(* IEC 61131-3 sources: STAR-PLC-Agent/results/raw/codex_matrix_resume_20261114/codex_deepseek/PUB020/functional/attempt_0001, 1 file *)

(* ---- test_program.st ---- *)
PROGRAM PLC_PRG
VAR
 BenchStep : UDINT := 0;
 BenchCalls : UDINT := 0;
 BenchDone : BOOL := FALSE;
 BenchUut0 : FB_Task;
 BenchUut1 : FB_Task;
 BenchUut2 : FB_Task;
 BenchUut3 : FB_Task;
 BenchUut4 : FB_Task;
 BenchUut5 : FB_Task;
 BenchUut6 : FB_Task;
 BenchUut7 : FB_Task;
 BenchUut8 : FB_Task;
 BenchUut9 : FB_Task;
 BenchUut10 : FB_Task;
 TraceIn_Mode : ARRAY[0..155] OF BOOL;
 TraceIn_ForwardButton : ARRAY[0..155] OF BOOL;
 TraceIn_ReverseButton : ARRAY[0..155] OF BOOL;
 TraceIn_SensorFeed : ARRAY[0..155] OF BOOL;
 TraceIn_SensorWash : ARRAY[0..155] OF BOOL;
 TraceIn_SensorWeight : ARRAY[0..155] OF BOOL;
 TraceIn_SensorFiring : ARRAY[0..155] OF BOOL;
 TraceIn_SensorOutput : ARRAY[0..155] OF BOOL;
 TraceIn_washComplete : ARRAY[0..155] OF BOOL;
 TraceIn_weightComplete : ARRAY[0..155] OF BOOL;
 TraceIn_weight : ARRAY[0..155] OF REAL;
 TraceIn_firingComplete : ARRAY[0..155] OF BOOL;
 TraceOut_MotorForward : ARRAY[0..155] OF BOOL;
 TraceOut_MotorReverse : ARRAY[0..155] OF BOOL;
 TraceOut_kick : ARRAY[0..155] OF BOOL;
 TraceOut_CompletionLight : ARRAY[0..155] OF BOOL;
 TraceOut_firingTemp : ARRAY[0..155] OF REAL;
END_VAR

IF NOT BenchDone THEN
 CASE BenchStep OF
 0:
   BenchUut0.Mode := FALSE;
   BenchUut0.ForwardButton := FALSE;
   BenchUut0.ReverseButton := FALSE;
   BenchUut0.SensorFeed := FALSE;
   BenchUut0.SensorWash := FALSE;
   BenchUut0.SensorWeight := FALSE;
   BenchUut0.SensorFiring := FALSE;
   BenchUut0.SensorOutput := FALSE;
   BenchUut0.washComplete := FALSE;
   BenchUut0.weightComplete := FALSE;
   BenchUut0.weight := REAL#0.0;
   BenchUut0.firingComplete := FALSE;
   TraceIn_Mode[0] := BenchUut0.Mode;
   TraceIn_ForwardButton[0] := BenchUut0.ForwardButton;
   TraceIn_ReverseButton[0] := BenchUut0.ReverseButton;
   TraceIn_SensorFeed[0] := BenchUut0.SensorFeed;
   TraceIn_SensorWash[0] := BenchUut0.SensorWash;
   TraceIn_SensorWeight[0] := BenchUut0.SensorWeight;
   TraceIn_SensorFiring[0] := BenchUut0.SensorFiring;
   TraceIn_SensorOutput[0] := BenchUut0.SensorOutput;
   TraceIn_washComplete[0] := BenchUut0.washComplete;
   TraceIn_weightComplete[0] := BenchUut0.weightComplete;
   TraceIn_weight[0] := BenchUut0.weight;
   TraceIn_firingComplete[0] := BenchUut0.firingComplete;
   BenchUut0();
   TraceOut_MotorForward[0] := BenchUut0.MotorForward;
   TraceOut_MotorReverse[0] := BenchUut0.MotorReverse;
   TraceOut_kick[0] := BenchUut0.kick;
   TraceOut_CompletionLight[0] := BenchUut0.CompletionLight;
   TraceOut_firingTemp[0] := BenchUut0.firingTemp;
   BenchCalls := BenchCalls + 1;
 1:
   BenchUut0.Mode := FALSE;
   BenchUut0.ForwardButton := TRUE;
   BenchUut0.ReverseButton := FALSE;
   BenchUut0.SensorFeed := FALSE;
   BenchUut0.SensorWash := FALSE;
   BenchUut0.SensorWeight := FALSE;
   BenchUut0.SensorFiring := FALSE;
   BenchUut0.SensorOutput := FALSE;
   BenchUut0.washComplete := FALSE;
   BenchUut0.weightComplete := FALSE;
   BenchUut0.weight := REAL#0.0;
   BenchUut0.firingComplete := FALSE;
   TraceIn_Mode[1] := BenchUut0.Mode;
   TraceIn_ForwardButton[1] := BenchUut0.ForwardButton;
   TraceIn_ReverseButton[1] := BenchUut0.ReverseButton;
   TraceIn_SensorFeed[1] := BenchUut0.SensorFeed;
   TraceIn_SensorWash[1] := BenchUut0.SensorWash;
   TraceIn_SensorWeight[1] := BenchUut0.SensorWeight;
   TraceIn_SensorFiring[1] := BenchUut0.SensorFiring;
   TraceIn_SensorOutput[1] := BenchUut0.SensorOutput;
   TraceIn_washComplete[1] := BenchUut0.washComplete;
   TraceIn_weightComplete[1] := BenchUut0.weightComplete;
   TraceIn_weight[1] := BenchUut0.weight;
   TraceIn_firingComplete[1] := BenchUut0.firingComplete;
   BenchUut0();
   TraceOut_MotorForward[1] := BenchUut0.MotorForward;
   TraceOut_MotorReverse[1] := BenchUut0.MotorReverse;
   TraceOut_kick[1] := BenchUut0.kick;
   TraceOut_CompletionLight[1] := BenchUut0.CompletionLight;
   TraceOut_firingTemp[1] := BenchUut0.firingTemp;
   BenchCalls := BenchCalls + 1;
 2:
   BenchUut0.Mode := FALSE;
   BenchUut0.ForwardButton := FALSE;
   BenchUut0.ReverseButton := TRUE;
   BenchUut0.SensorFeed := FALSE;
   BenchUut0.SensorWash := FALSE;
   BenchUut0.SensorWeight := FALSE;
   BenchUut0.SensorFiring := FALSE;
   BenchUut0.SensorOutput := FALSE;
   BenchUut0.washComplete := FALSE;
   BenchUut0.weightComplete := FALSE;
   BenchUut0.weight := REAL#0.0;
   BenchUut0.firingComplete := FALSE;
   TraceIn_Mode[2] := BenchUut0.Mode;
   TraceIn_ForwardButton[2] := BenchUut0.ForwardButton;
   TraceIn_ReverseButton[2] := BenchUut0.ReverseButton;
   TraceIn_SensorFeed[2] := BenchUut0.SensorFeed;
   TraceIn_SensorWash[2] := BenchUut0.SensorWash;
   TraceIn_SensorWeight[2] := BenchUut0.SensorWeight;
   TraceIn_SensorFiring[2] := BenchUut0.SensorFiring;
   TraceIn_SensorOutput[2] := BenchUut0.SensorOutput;
   TraceIn_washComplete[2] := BenchUut0.washComplete;
   TraceIn_weightComplete[2] := BenchUut0.weightComplete;
   TraceIn_weight[2] := BenchUut0.weight;
   TraceIn_firingComplete[2] := BenchUut0.firingComplete;
   BenchUut0();
   TraceOut_MotorForward[2] := BenchUut0.MotorForward;
   TraceOut_MotorReverse[2] := BenchUut0.MotorReverse;
   TraceOut_kick[2] := BenchUut0.kick;
   TraceOut_CompletionLight[2] := BenchUut0.CompletionLight;
   TraceOut_firingTemp[2] := BenchUut0.firingTemp;
   BenchCalls := BenchCalls + 1;
 3:
   BenchUut0.Mode := FALSE;
   BenchUut0.ForwardButton := TRUE;
   BenchUut0.ReverseButton := TRUE;
   BenchUut0.SensorFeed := FALSE;
   BenchUut0.SensorWash := FALSE;
   BenchUut0.SensorWeight := FALSE;
   BenchUut0.SensorFiring := FALSE;
   BenchUut0.SensorOutput := FALSE;
   BenchUut0.washComplete := FALSE;
   BenchUut0.weightComplete := FALSE;
   BenchUut0.weight := REAL#0.0;
   BenchUut0.firingComplete := FALSE;
   TraceIn_Mode[3] := BenchUut0.Mode;
   TraceIn_ForwardButton[3] := BenchUut0.ForwardButton;
   TraceIn_ReverseButton[3] := BenchUut0.ReverseButton;
   TraceIn_SensorFeed[3] := BenchUut0.SensorFeed;
   TraceIn_SensorWash[3] := BenchUut0.SensorWash;
   TraceIn_SensorWeight[3] := BenchUut0.SensorWeight;
   TraceIn_SensorFiring[3] := BenchUut0.SensorFiring;
   TraceIn_SensorOutput[3] := BenchUut0.SensorOutput;
   TraceIn_washComplete[3] := BenchUut0.washComplete;
   TraceIn_weightComplete[3] := BenchUut0.weightComplete;
   TraceIn_weight[3] := BenchUut0.weight;
   TraceIn_firingComplete[3] := BenchUut0.firingComplete;
   BenchUut0();
   TraceOut_MotorForward[3] := BenchUut0.MotorForward;
   TraceOut_MotorReverse[3] := BenchUut0.MotorReverse;
   TraceOut_kick[3] := BenchUut0.kick;
   TraceOut_CompletionLight[3] := BenchUut0.CompletionLight;
   TraceOut_firingTemp[3] := BenchUut0.firingTemp;
   BenchCalls := BenchCalls + 1;
 4:
   BenchUut1.Mode := TRUE;
   BenchUut1.ForwardButton := FALSE;
   BenchUut1.ReverseButton := FALSE;
   BenchUut1.SensorFeed := FALSE;
   BenchUut1.SensorWash := FALSE;
   BenchUut1.SensorWeight := FALSE;
   BenchUut1.SensorFiring := FALSE;
   BenchUut1.SensorOutput := FALSE;
   BenchUut1.washComplete := FALSE;
   BenchUut1.weightComplete := FALSE;
   BenchUut1.weight := REAL#0.0;
   BenchUut1.firingComplete := FALSE;
   TraceIn_Mode[4] := BenchUut1.Mode;
   TraceIn_ForwardButton[4] := BenchUut1.ForwardButton;
   TraceIn_ReverseButton[4] := BenchUut1.ReverseButton;
   TraceIn_SensorFeed[4] := BenchUut1.SensorFeed;
   TraceIn_SensorWash[4] := BenchUut1.SensorWash;
   TraceIn_SensorWeight[4] := BenchUut1.SensorWeight;
   TraceIn_SensorFiring[4] := BenchUut1.SensorFiring;
   TraceIn_SensorOutput[4] := BenchUut1.SensorOutput;
   TraceIn_washComplete[4] := BenchUut1.washComplete;
   TraceIn_weightComplete[4] := BenchUut1.weightComplete;
   TraceIn_weight[4] := BenchUut1.weight;
   TraceIn_firingComplete[4] := BenchUut1.firingComplete;
   BenchUut1();
   TraceOut_MotorForward[4] := BenchUut1.MotorForward;
   TraceOut_MotorReverse[4] := BenchUut1.MotorReverse;
   TraceOut_kick[4] := BenchUut1.kick;
   TraceOut_CompletionLight[4] := BenchUut1.CompletionLight;
   TraceOut_firingTemp[4] := BenchUut1.firingTemp;
   BenchCalls := BenchCalls + 1;
 5:
   BenchUut1.Mode := TRUE;
   BenchUut1.ForwardButton := FALSE;
   BenchUut1.ReverseButton := FALSE;
   BenchUut1.SensorFeed := TRUE;
   BenchUut1.SensorWash := FALSE;
   BenchUut1.SensorWeight := FALSE;
   BenchUut1.SensorFiring := FALSE;
   BenchUut1.SensorOutput := FALSE;
   BenchUut1.washComplete := FALSE;
   BenchUut1.weightComplete := FALSE;
   BenchUut1.weight := REAL#0.0;
   BenchUut1.firingComplete := FALSE;
   TraceIn_Mode[5] := BenchUut1.Mode;
   TraceIn_ForwardButton[5] := BenchUut1.ForwardButton;
   TraceIn_ReverseButton[5] := BenchUut1.ReverseButton;
   TraceIn_SensorFeed[5] := BenchUut1.SensorFeed;
   TraceIn_SensorWash[5] := BenchUut1.SensorWash;
   TraceIn_SensorWeight[5] := BenchUut1.SensorWeight;
   TraceIn_SensorFiring[5] := BenchUut1.SensorFiring;
   TraceIn_SensorOutput[5] := BenchUut1.SensorOutput;
   TraceIn_washComplete[5] := BenchUut1.washComplete;
   TraceIn_weightComplete[5] := BenchUut1.weightComplete;
   TraceIn_weight[5] := BenchUut1.weight;
   TraceIn_firingComplete[5] := BenchUut1.firingComplete;
   BenchUut1();
   TraceOut_MotorForward[5] := BenchUut1.MotorForward;
   TraceOut_MotorReverse[5] := BenchUut1.MotorReverse;
   TraceOut_kick[5] := BenchUut1.kick;
   TraceOut_CompletionLight[5] := BenchUut1.CompletionLight;
   TraceOut_firingTemp[5] := BenchUut1.firingTemp;
   BenchCalls := BenchCalls + 1;
 6:
   BenchUut1.Mode := TRUE;
   BenchUut1.ForwardButton := FALSE;
   BenchUut1.ReverseButton := FALSE;
   BenchUut1.SensorFeed := FALSE;
   BenchUut1.SensorWash := TRUE;
   BenchUut1.SensorWeight := FALSE;
   BenchUut1.SensorFiring := FALSE;
   BenchUut1.SensorOutput := FALSE;
   BenchUut1.washComplete := FALSE;
   BenchUut1.weightComplete := FALSE;
   BenchUut1.weight := REAL#0.0;
   BenchUut1.firingComplete := FALSE;
   TraceIn_Mode[6] := BenchUut1.Mode;
   TraceIn_ForwardButton[6] := BenchUut1.ForwardButton;
   TraceIn_ReverseButton[6] := BenchUut1.ReverseButton;
   TraceIn_SensorFeed[6] := BenchUut1.SensorFeed;
   TraceIn_SensorWash[6] := BenchUut1.SensorWash;
   TraceIn_SensorWeight[6] := BenchUut1.SensorWeight;
   TraceIn_SensorFiring[6] := BenchUut1.SensorFiring;
   TraceIn_SensorOutput[6] := BenchUut1.SensorOutput;
   TraceIn_washComplete[6] := BenchUut1.washComplete;
   TraceIn_weightComplete[6] := BenchUut1.weightComplete;
   TraceIn_weight[6] := BenchUut1.weight;
   TraceIn_firingComplete[6] := BenchUut1.firingComplete;
   BenchUut1();
   TraceOut_MotorForward[6] := BenchUut1.MotorForward;
   TraceOut_MotorReverse[6] := BenchUut1.MotorReverse;
   TraceOut_kick[6] := BenchUut1.kick;
   TraceOut_CompletionLight[6] := BenchUut1.CompletionLight;
   TraceOut_firingTemp[6] := BenchUut1.firingTemp;
   BenchCalls := BenchCalls + 1;
 7:
   BenchUut1.Mode := TRUE;
   BenchUut1.ForwardButton := FALSE;
   BenchUut1.ReverseButton := FALSE;
   BenchUut1.SensorFeed := FALSE;
   BenchUut1.SensorWash := TRUE;
   BenchUut1.SensorWeight := FALSE;
   BenchUut1.SensorFiring := FALSE;
   BenchUut1.SensorOutput := FALSE;
   BenchUut1.washComplete := TRUE;
   BenchUut1.weightComplete := FALSE;
   BenchUut1.weight := REAL#0.0;
   BenchUut1.firingComplete := FALSE;
   TraceIn_Mode[7] := BenchUut1.Mode;
   TraceIn_ForwardButton[7] := BenchUut1.ForwardButton;
   TraceIn_ReverseButton[7] := BenchUut1.ReverseButton;
   TraceIn_SensorFeed[7] := BenchUut1.SensorFeed;
   TraceIn_SensorWash[7] := BenchUut1.SensorWash;
   TraceIn_SensorWeight[7] := BenchUut1.SensorWeight;
   TraceIn_SensorFiring[7] := BenchUut1.SensorFiring;
   TraceIn_SensorOutput[7] := BenchUut1.SensorOutput;
   TraceIn_washComplete[7] := BenchUut1.washComplete;
   TraceIn_weightComplete[7] := BenchUut1.weightComplete;
   TraceIn_weight[7] := BenchUut1.weight;
   TraceIn_firingComplete[7] := BenchUut1.firingComplete;
   BenchUut1();
   TraceOut_MotorForward[7] := BenchUut1.MotorForward;
   TraceOut_MotorReverse[7] := BenchUut1.MotorReverse;
   TraceOut_kick[7] := BenchUut1.kick;
   TraceOut_CompletionLight[7] := BenchUut1.CompletionLight;
   TraceOut_firingTemp[7] := BenchUut1.firingTemp;
   BenchCalls := BenchCalls + 1;
 8:
   BenchUut1.Mode := TRUE;
   BenchUut1.ForwardButton := FALSE;
   BenchUut1.ReverseButton := FALSE;
   BenchUut1.SensorFeed := FALSE;
   BenchUut1.SensorWash := FALSE;
   BenchUut1.SensorWeight := TRUE;
   BenchUut1.SensorFiring := FALSE;
   BenchUut1.SensorOutput := FALSE;
   BenchUut1.washComplete := FALSE;
   BenchUut1.weightComplete := FALSE;
   BenchUut1.weight := REAL#0.0;
   BenchUut1.firingComplete := FALSE;
   TraceIn_Mode[8] := BenchUut1.Mode;
   TraceIn_ForwardButton[8] := BenchUut1.ForwardButton;
   TraceIn_ReverseButton[8] := BenchUut1.ReverseButton;
   TraceIn_SensorFeed[8] := BenchUut1.SensorFeed;
   TraceIn_SensorWash[8] := BenchUut1.SensorWash;
   TraceIn_SensorWeight[8] := BenchUut1.SensorWeight;
   TraceIn_SensorFiring[8] := BenchUut1.SensorFiring;
   TraceIn_SensorOutput[8] := BenchUut1.SensorOutput;
   TraceIn_washComplete[8] := BenchUut1.washComplete;
   TraceIn_weightComplete[8] := BenchUut1.weightComplete;
   TraceIn_weight[8] := BenchUut1.weight;
   TraceIn_firingComplete[8] := BenchUut1.firingComplete;
   BenchUut1();
   TraceOut_MotorForward[8] := BenchUut1.MotorForward;
   TraceOut_MotorReverse[8] := BenchUut1.MotorReverse;
   TraceOut_kick[8] := BenchUut1.kick;
   TraceOut_CompletionLight[8] := BenchUut1.CompletionLight;
   TraceOut_firingTemp[8] := BenchUut1.firingTemp;
   BenchCalls := BenchCalls + 1;
 9:
   BenchUut1.Mode := TRUE;
   BenchUut1.ForwardButton := FALSE;
   BenchUut1.ReverseButton := FALSE;
   BenchUut1.SensorFeed := FALSE;
   BenchUut1.SensorWash := FALSE;
   BenchUut1.SensorWeight := TRUE;
   BenchUut1.SensorFiring := FALSE;
   BenchUut1.SensorOutput := FALSE;
   BenchUut1.washComplete := FALSE;
   BenchUut1.weightComplete := TRUE;
   BenchUut1.weight := REAL#100.0;
   BenchUut1.firingComplete := FALSE;
   TraceIn_Mode[9] := BenchUut1.Mode;
   TraceIn_ForwardButton[9] := BenchUut1.ForwardButton;
   TraceIn_ReverseButton[9] := BenchUut1.ReverseButton;
   TraceIn_SensorFeed[9] := BenchUut1.SensorFeed;
   TraceIn_SensorWash[9] := BenchUut1.SensorWash;
   TraceIn_SensorWeight[9] := BenchUut1.SensorWeight;
   TraceIn_SensorFiring[9] := BenchUut1.SensorFiring;
   TraceIn_SensorOutput[9] := BenchUut1.SensorOutput;
   TraceIn_washComplete[9] := BenchUut1.washComplete;
   TraceIn_weightComplete[9] := BenchUut1.weightComplete;
   TraceIn_weight[9] := BenchUut1.weight;
   TraceIn_firingComplete[9] := BenchUut1.firingComplete;
   BenchUut1();
   TraceOut_MotorForward[9] := BenchUut1.MotorForward;
   TraceOut_MotorReverse[9] := BenchUut1.MotorReverse;
   TraceOut_kick[9] := BenchUut1.kick;
   TraceOut_CompletionLight[9] := BenchUut1.CompletionLight;
   TraceOut_firingTemp[9] := BenchUut1.firingTemp;
   BenchCalls := BenchCalls + 1;
 10:
   BenchUut1.Mode := TRUE;
   BenchUut1.ForwardButton := FALSE;
   BenchUut1.ReverseButton := FALSE;
   BenchUut1.SensorFeed := FALSE;
   BenchUut1.SensorWash := FALSE;
   BenchUut1.SensorWeight := FALSE;
   BenchUut1.SensorFiring := TRUE;
   BenchUut1.SensorOutput := FALSE;
   BenchUut1.washComplete := FALSE;
   BenchUut1.weightComplete := FALSE;
   BenchUut1.weight := REAL#0.0;
   BenchUut1.firingComplete := FALSE;
   TraceIn_Mode[10] := BenchUut1.Mode;
   TraceIn_ForwardButton[10] := BenchUut1.ForwardButton;
   TraceIn_ReverseButton[10] := BenchUut1.ReverseButton;
   TraceIn_SensorFeed[10] := BenchUut1.SensorFeed;
   TraceIn_SensorWash[10] := BenchUut1.SensorWash;
   TraceIn_SensorWeight[10] := BenchUut1.SensorWeight;
   TraceIn_SensorFiring[10] := BenchUut1.SensorFiring;
   TraceIn_SensorOutput[10] := BenchUut1.SensorOutput;
   TraceIn_washComplete[10] := BenchUut1.washComplete;
   TraceIn_weightComplete[10] := BenchUut1.weightComplete;
   TraceIn_weight[10] := BenchUut1.weight;
   TraceIn_firingComplete[10] := BenchUut1.firingComplete;
   BenchUut1();
   TraceOut_MotorForward[10] := BenchUut1.MotorForward;
   TraceOut_MotorReverse[10] := BenchUut1.MotorReverse;
   TraceOut_kick[10] := BenchUut1.kick;
   TraceOut_CompletionLight[10] := BenchUut1.CompletionLight;
   TraceOut_firingTemp[10] := BenchUut1.firingTemp;
   BenchCalls := BenchCalls + 1;
 11:
   BenchUut1.Mode := TRUE;
   BenchUut1.ForwardButton := FALSE;
   BenchUut1.ReverseButton := FALSE;
   BenchUut1.SensorFeed := FALSE;
   BenchUut1.SensorWash := FALSE;
   BenchUut1.SensorWeight := FALSE;
   BenchUut1.SensorFiring := TRUE;
   BenchUut1.SensorOutput := FALSE;
   BenchUut1.washComplete := FALSE;
   BenchUut1.weightComplete := FALSE;
   BenchUut1.weight := REAL#0.0;
   BenchUut1.firingComplete := TRUE;
   TraceIn_Mode[11] := BenchUut1.Mode;
   TraceIn_ForwardButton[11] := BenchUut1.ForwardButton;
   TraceIn_ReverseButton[11] := BenchUut1.ReverseButton;
   TraceIn_SensorFeed[11] := BenchUut1.SensorFeed;
   TraceIn_SensorWash[11] := BenchUut1.SensorWash;
   TraceIn_SensorWeight[11] := BenchUut1.SensorWeight;
   TraceIn_SensorFiring[11] := BenchUut1.SensorFiring;
   TraceIn_SensorOutput[11] := BenchUut1.SensorOutput;
   TraceIn_washComplete[11] := BenchUut1.washComplete;
   TraceIn_weightComplete[11] := BenchUut1.weightComplete;
   TraceIn_weight[11] := BenchUut1.weight;
   TraceIn_firingComplete[11] := BenchUut1.firingComplete;
   BenchUut1();
   TraceOut_MotorForward[11] := BenchUut1.MotorForward;
   TraceOut_MotorReverse[11] := BenchUut1.MotorReverse;
   TraceOut_kick[11] := BenchUut1.kick;
   TraceOut_CompletionLight[11] := BenchUut1.CompletionLight;
   TraceOut_firingTemp[11] := BenchUut1.firingTemp;
   BenchCalls := BenchCalls + 1;
 12:
   BenchUut1.Mode := TRUE;
   BenchUut1.ForwardButton := FALSE;
   BenchUut1.ReverseButton := FALSE;
   BenchUut1.SensorFeed := FALSE;
   BenchUut1.SensorWash := FALSE;
   BenchUut1.SensorWeight := FALSE;
   BenchUut1.SensorFiring := FALSE;
   BenchUut1.SensorOutput := TRUE;
   BenchUut1.washComplete := FALSE;
   BenchUut1.weightComplete := FALSE;
   BenchUut1.weight := REAL#0.0;
   BenchUut1.firingComplete := FALSE;
   TraceIn_Mode[12] := BenchUut1.Mode;
   TraceIn_ForwardButton[12] := BenchUut1.ForwardButton;
   TraceIn_ReverseButton[12] := BenchUut1.ReverseButton;
   TraceIn_SensorFeed[12] := BenchUut1.SensorFeed;
   TraceIn_SensorWash[12] := BenchUut1.SensorWash;
   TraceIn_SensorWeight[12] := BenchUut1.SensorWeight;
   TraceIn_SensorFiring[12] := BenchUut1.SensorFiring;
   TraceIn_SensorOutput[12] := BenchUut1.SensorOutput;
   TraceIn_washComplete[12] := BenchUut1.washComplete;
   TraceIn_weightComplete[12] := BenchUut1.weightComplete;
   TraceIn_weight[12] := BenchUut1.weight;
   TraceIn_firingComplete[12] := BenchUut1.firingComplete;
   BenchUut1();
   TraceOut_MotorForward[12] := BenchUut1.MotorForward;
   TraceOut_MotorReverse[12] := BenchUut1.MotorReverse;
   TraceOut_kick[12] := BenchUut1.kick;
   TraceOut_CompletionLight[12] := BenchUut1.CompletionLight;
   TraceOut_firingTemp[12] := BenchUut1.firingTemp;
   BenchCalls := BenchCalls + 1;
 13:
   BenchUut1.Mode := TRUE;
   BenchUut1.ForwardButton := FALSE;
   BenchUut1.ReverseButton := FALSE;
   BenchUut1.SensorFeed := FALSE;
   BenchUut1.SensorWash := FALSE;
   BenchUut1.SensorWeight := FALSE;
   BenchUut1.SensorFiring := FALSE;
   BenchUut1.SensorOutput := TRUE;
   BenchUut1.washComplete := FALSE;
   BenchUut1.weightComplete := FALSE;
   BenchUut1.weight := REAL#0.0;
   BenchUut1.firingComplete := FALSE;
   TraceIn_Mode[13] := BenchUut1.Mode;
   TraceIn_ForwardButton[13] := BenchUut1.ForwardButton;
   TraceIn_ReverseButton[13] := BenchUut1.ReverseButton;
   TraceIn_SensorFeed[13] := BenchUut1.SensorFeed;
   TraceIn_SensorWash[13] := BenchUut1.SensorWash;
   TraceIn_SensorWeight[13] := BenchUut1.SensorWeight;
   TraceIn_SensorFiring[13] := BenchUut1.SensorFiring;
   TraceIn_SensorOutput[13] := BenchUut1.SensorOutput;
   TraceIn_washComplete[13] := BenchUut1.washComplete;
   TraceIn_weightComplete[13] := BenchUut1.weightComplete;
   TraceIn_weight[13] := BenchUut1.weight;
   TraceIn_firingComplete[13] := BenchUut1.firingComplete;
   BenchUut1();
   TraceOut_MotorForward[13] := BenchUut1.MotorForward;
   TraceOut_MotorReverse[13] := BenchUut1.MotorReverse;
   TraceOut_kick[13] := BenchUut1.kick;
   TraceOut_CompletionLight[13] := BenchUut1.CompletionLight;
   TraceOut_firingTemp[13] := BenchUut1.firingTemp;
   BenchCalls := BenchCalls + 1;
 14:
   BenchUut1.Mode := TRUE;
   BenchUut1.ForwardButton := FALSE;
   BenchUut1.ReverseButton := FALSE;
   BenchUut1.SensorFeed := FALSE;
   BenchUut1.SensorWash := FALSE;
   BenchUut1.SensorWeight := FALSE;
   BenchUut1.SensorFiring := FALSE;
   BenchUut1.SensorOutput := FALSE;
   BenchUut1.washComplete := FALSE;
   BenchUut1.weightComplete := FALSE;
   BenchUut1.weight := REAL#0.0;
   BenchUut1.firingComplete := FALSE;
   TraceIn_Mode[14] := BenchUut1.Mode;
   TraceIn_ForwardButton[14] := BenchUut1.ForwardButton;
   TraceIn_ReverseButton[14] := BenchUut1.ReverseButton;
   TraceIn_SensorFeed[14] := BenchUut1.SensorFeed;
   TraceIn_SensorWash[14] := BenchUut1.SensorWash;
   TraceIn_SensorWeight[14] := BenchUut1.SensorWeight;
   TraceIn_SensorFiring[14] := BenchUut1.SensorFiring;
   TraceIn_SensorOutput[14] := BenchUut1.SensorOutput;
   TraceIn_washComplete[14] := BenchUut1.washComplete;
   TraceIn_weightComplete[14] := BenchUut1.weightComplete;
   TraceIn_weight[14] := BenchUut1.weight;
   TraceIn_firingComplete[14] := BenchUut1.firingComplete;
   BenchUut1();
   TraceOut_MotorForward[14] := BenchUut1.MotorForward;
   TraceOut_MotorReverse[14] := BenchUut1.MotorReverse;
   TraceOut_kick[14] := BenchUut1.kick;
   TraceOut_CompletionLight[14] := BenchUut1.CompletionLight;
   TraceOut_firingTemp[14] := BenchUut1.firingTemp;
   BenchCalls := BenchCalls + 1;
 15:
   BenchUut2.Mode := TRUE;
   BenchUut2.ForwardButton := FALSE;
   BenchUut2.ReverseButton := FALSE;
   BenchUut2.SensorFeed := FALSE;
   BenchUut2.SensorWash := FALSE;
   BenchUut2.SensorWeight := FALSE;
   BenchUut2.SensorFiring := FALSE;
   BenchUut2.SensorOutput := FALSE;
   BenchUut2.washComplete := FALSE;
   BenchUut2.weightComplete := FALSE;
   BenchUut2.weight := REAL#0.0;
   BenchUut2.firingComplete := FALSE;
   TraceIn_Mode[15] := BenchUut2.Mode;
   TraceIn_ForwardButton[15] := BenchUut2.ForwardButton;
   TraceIn_ReverseButton[15] := BenchUut2.ReverseButton;
   TraceIn_SensorFeed[15] := BenchUut2.SensorFeed;
   TraceIn_SensorWash[15] := BenchUut2.SensorWash;
   TraceIn_SensorWeight[15] := BenchUut2.SensorWeight;
   TraceIn_SensorFiring[15] := BenchUut2.SensorFiring;
   TraceIn_SensorOutput[15] := BenchUut2.SensorOutput;
   TraceIn_washComplete[15] := BenchUut2.washComplete;
   TraceIn_weightComplete[15] := BenchUut2.weightComplete;
   TraceIn_weight[15] := BenchUut2.weight;
   TraceIn_firingComplete[15] := BenchUut2.firingComplete;
   BenchUut2();
   TraceOut_MotorForward[15] := BenchUut2.MotorForward;
   TraceOut_MotorReverse[15] := BenchUut2.MotorReverse;
   TraceOut_kick[15] := BenchUut2.kick;
   TraceOut_CompletionLight[15] := BenchUut2.CompletionLight;
   TraceOut_firingTemp[15] := BenchUut2.firingTemp;
   BenchCalls := BenchCalls + 1;
 16:
   BenchUut2.Mode := TRUE;
   BenchUut2.ForwardButton := FALSE;
   BenchUut2.ReverseButton := FALSE;
   BenchUut2.SensorFeed := TRUE;
   BenchUut2.SensorWash := FALSE;
   BenchUut2.SensorWeight := FALSE;
   BenchUut2.SensorFiring := FALSE;
   BenchUut2.SensorOutput := FALSE;
   BenchUut2.washComplete := FALSE;
   BenchUut2.weightComplete := FALSE;
   BenchUut2.weight := REAL#0.0;
   BenchUut2.firingComplete := FALSE;
   TraceIn_Mode[16] := BenchUut2.Mode;
   TraceIn_ForwardButton[16] := BenchUut2.ForwardButton;
   TraceIn_ReverseButton[16] := BenchUut2.ReverseButton;
   TraceIn_SensorFeed[16] := BenchUut2.SensorFeed;
   TraceIn_SensorWash[16] := BenchUut2.SensorWash;
   TraceIn_SensorWeight[16] := BenchUut2.SensorWeight;
   TraceIn_SensorFiring[16] := BenchUut2.SensorFiring;
   TraceIn_SensorOutput[16] := BenchUut2.SensorOutput;
   TraceIn_washComplete[16] := BenchUut2.washComplete;
   TraceIn_weightComplete[16] := BenchUut2.weightComplete;
   TraceIn_weight[16] := BenchUut2.weight;
   TraceIn_firingComplete[16] := BenchUut2.firingComplete;
   BenchUut2();
   TraceOut_MotorForward[16] := BenchUut2.MotorForward;
   TraceOut_MotorReverse[16] := BenchUut2.MotorReverse;
   TraceOut_kick[16] := BenchUut2.kick;
   TraceOut_CompletionLight[16] := BenchUut2.CompletionLight;
   TraceOut_firingTemp[16] := BenchUut2.firingTemp;
   BenchCalls := BenchCalls + 1;
 17:
   BenchUut2.Mode := TRUE;
   BenchUut2.ForwardButton := FALSE;
   BenchUut2.ReverseButton := FALSE;
   BenchUut2.SensorFeed := FALSE;
   BenchUut2.SensorWash := TRUE;
   BenchUut2.SensorWeight := FALSE;
   BenchUut2.SensorFiring := FALSE;
   BenchUut2.SensorOutput := FALSE;
   BenchUut2.washComplete := FALSE;
   BenchUut2.weightComplete := FALSE;
   BenchUut2.weight := REAL#0.0;
   BenchUut2.firingComplete := FALSE;
   TraceIn_Mode[17] := BenchUut2.Mode;
   TraceIn_ForwardButton[17] := BenchUut2.ForwardButton;
   TraceIn_ReverseButton[17] := BenchUut2.ReverseButton;
   TraceIn_SensorFeed[17] := BenchUut2.SensorFeed;
   TraceIn_SensorWash[17] := BenchUut2.SensorWash;
   TraceIn_SensorWeight[17] := BenchUut2.SensorWeight;
   TraceIn_SensorFiring[17] := BenchUut2.SensorFiring;
   TraceIn_SensorOutput[17] := BenchUut2.SensorOutput;
   TraceIn_washComplete[17] := BenchUut2.washComplete;
   TraceIn_weightComplete[17] := BenchUut2.weightComplete;
   TraceIn_weight[17] := BenchUut2.weight;
   TraceIn_firingComplete[17] := BenchUut2.firingComplete;
   BenchUut2();
   TraceOut_MotorForward[17] := BenchUut2.MotorForward;
   TraceOut_MotorReverse[17] := BenchUut2.MotorReverse;
   TraceOut_kick[17] := BenchUut2.kick;
   TraceOut_CompletionLight[17] := BenchUut2.CompletionLight;
   TraceOut_firingTemp[17] := BenchUut2.firingTemp;
   BenchCalls := BenchCalls + 1;
 18:
   BenchUut2.Mode := TRUE;
   BenchUut2.ForwardButton := FALSE;
   BenchUut2.ReverseButton := FALSE;
   BenchUut2.SensorFeed := FALSE;
   BenchUut2.SensorWash := TRUE;
   BenchUut2.SensorWeight := FALSE;
   BenchUut2.SensorFiring := FALSE;
   BenchUut2.SensorOutput := FALSE;
   BenchUut2.washComplete := TRUE;
   BenchUut2.weightComplete := FALSE;
   BenchUut2.weight := REAL#0.0;
   BenchUut2.firingComplete := FALSE;
   TraceIn_Mode[18] := BenchUut2.Mode;
   TraceIn_ForwardButton[18] := BenchUut2.ForwardButton;
   TraceIn_ReverseButton[18] := BenchUut2.ReverseButton;
   TraceIn_SensorFeed[18] := BenchUut2.SensorFeed;
   TraceIn_SensorWash[18] := BenchUut2.SensorWash;
   TraceIn_SensorWeight[18] := BenchUut2.SensorWeight;
   TraceIn_SensorFiring[18] := BenchUut2.SensorFiring;
   TraceIn_SensorOutput[18] := BenchUut2.SensorOutput;
   TraceIn_washComplete[18] := BenchUut2.washComplete;
   TraceIn_weightComplete[18] := BenchUut2.weightComplete;
   TraceIn_weight[18] := BenchUut2.weight;
   TraceIn_firingComplete[18] := BenchUut2.firingComplete;
   BenchUut2();
   TraceOut_MotorForward[18] := BenchUut2.MotorForward;
   TraceOut_MotorReverse[18] := BenchUut2.MotorReverse;
   TraceOut_kick[18] := BenchUut2.kick;
   TraceOut_CompletionLight[18] := BenchUut2.CompletionLight;
   TraceOut_firingTemp[18] := BenchUut2.firingTemp;
   BenchCalls := BenchCalls + 1;
 19:
   BenchUut2.Mode := TRUE;
   BenchUut2.ForwardButton := FALSE;
   BenchUut2.ReverseButton := FALSE;
   BenchUut2.SensorFeed := FALSE;
   BenchUut2.SensorWash := FALSE;
   BenchUut2.SensorWeight := TRUE;
   BenchUut2.SensorFiring := FALSE;
   BenchUut2.SensorOutput := FALSE;
   BenchUut2.washComplete := FALSE;
   BenchUut2.weightComplete := FALSE;
   BenchUut2.weight := REAL#0.0;
   BenchUut2.firingComplete := FALSE;
   TraceIn_Mode[19] := BenchUut2.Mode;
   TraceIn_ForwardButton[19] := BenchUut2.ForwardButton;
   TraceIn_ReverseButton[19] := BenchUut2.ReverseButton;
   TraceIn_SensorFeed[19] := BenchUut2.SensorFeed;
   TraceIn_SensorWash[19] := BenchUut2.SensorWash;
   TraceIn_SensorWeight[19] := BenchUut2.SensorWeight;
   TraceIn_SensorFiring[19] := BenchUut2.SensorFiring;
   TraceIn_SensorOutput[19] := BenchUut2.SensorOutput;
   TraceIn_washComplete[19] := BenchUut2.washComplete;
   TraceIn_weightComplete[19] := BenchUut2.weightComplete;
   TraceIn_weight[19] := BenchUut2.weight;
   TraceIn_firingComplete[19] := BenchUut2.firingComplete;
   BenchUut2();
   TraceOut_MotorForward[19] := BenchUut2.MotorForward;
   TraceOut_MotorReverse[19] := BenchUut2.MotorReverse;
   TraceOut_kick[19] := BenchUut2.kick;
   TraceOut_CompletionLight[19] := BenchUut2.CompletionLight;
   TraceOut_firingTemp[19] := BenchUut2.firingTemp;
   BenchCalls := BenchCalls + 1;
 20:
   BenchUut2.Mode := TRUE;
   BenchUut2.ForwardButton := FALSE;
   BenchUut2.ReverseButton := FALSE;
   BenchUut2.SensorFeed := FALSE;
   BenchUut2.SensorWash := FALSE;
   BenchUut2.SensorWeight := TRUE;
   BenchUut2.SensorFiring := FALSE;
   BenchUut2.SensorOutput := FALSE;
   BenchUut2.washComplete := FALSE;
   BenchUut2.weightComplete := TRUE;
   BenchUut2.weight := REAL#150.0;
   BenchUut2.firingComplete := FALSE;
   TraceIn_Mode[20] := BenchUut2.Mode;
   TraceIn_ForwardButton[20] := BenchUut2.ForwardButton;
   TraceIn_ReverseButton[20] := BenchUut2.ReverseButton;
   TraceIn_SensorFeed[20] := BenchUut2.SensorFeed;
   TraceIn_SensorWash[20] := BenchUut2.SensorWash;
   TraceIn_SensorWeight[20] := BenchUut2.SensorWeight;
   TraceIn_SensorFiring[20] := BenchUut2.SensorFiring;
   TraceIn_SensorOutput[20] := BenchUut2.SensorOutput;
   TraceIn_washComplete[20] := BenchUut2.washComplete;
   TraceIn_weightComplete[20] := BenchUut2.weightComplete;
   TraceIn_weight[20] := BenchUut2.weight;
   TraceIn_firingComplete[20] := BenchUut2.firingComplete;
   BenchUut2();
   TraceOut_MotorForward[20] := BenchUut2.MotorForward;
   TraceOut_MotorReverse[20] := BenchUut2.MotorReverse;
   TraceOut_kick[20] := BenchUut2.kick;
   TraceOut_CompletionLight[20] := BenchUut2.CompletionLight;
   TraceOut_firingTemp[20] := BenchUut2.firingTemp;
   BenchCalls := BenchCalls + 1;
 21:
   BenchUut2.Mode := TRUE;
   BenchUut2.ForwardButton := FALSE;
   BenchUut2.ReverseButton := FALSE;
   BenchUut2.SensorFeed := FALSE;
   BenchUut2.SensorWash := FALSE;
   BenchUut2.SensorWeight := FALSE;
   BenchUut2.SensorFiring := TRUE;
   BenchUut2.SensorOutput := FALSE;
   BenchUut2.washComplete := FALSE;
   BenchUut2.weightComplete := FALSE;
   BenchUut2.weight := REAL#0.0;
   BenchUut2.firingComplete := FALSE;
   TraceIn_Mode[21] := BenchUut2.Mode;
   TraceIn_ForwardButton[21] := BenchUut2.ForwardButton;
   TraceIn_ReverseButton[21] := BenchUut2.ReverseButton;
   TraceIn_SensorFeed[21] := BenchUut2.SensorFeed;
   TraceIn_SensorWash[21] := BenchUut2.SensorWash;
   TraceIn_SensorWeight[21] := BenchUut2.SensorWeight;
   TraceIn_SensorFiring[21] := BenchUut2.SensorFiring;
   TraceIn_SensorOutput[21] := BenchUut2.SensorOutput;
   TraceIn_washComplete[21] := BenchUut2.washComplete;
   TraceIn_weightComplete[21] := BenchUut2.weightComplete;
   TraceIn_weight[21] := BenchUut2.weight;
   TraceIn_firingComplete[21] := BenchUut2.firingComplete;
   BenchUut2();
   TraceOut_MotorForward[21] := BenchUut2.MotorForward;
   TraceOut_MotorReverse[21] := BenchUut2.MotorReverse;
   TraceOut_kick[21] := BenchUut2.kick;
   TraceOut_CompletionLight[21] := BenchUut2.CompletionLight;
   TraceOut_firingTemp[21] := BenchUut2.firingTemp;
   BenchCalls := BenchCalls + 1;
 22:
   BenchUut2.Mode := TRUE;
   BenchUut2.ForwardButton := FALSE;
   BenchUut2.ReverseButton := FALSE;
   BenchUut2.SensorFeed := FALSE;
   BenchUut2.SensorWash := FALSE;
   BenchUut2.SensorWeight := FALSE;
   BenchUut2.SensorFiring := TRUE;
   BenchUut2.SensorOutput := FALSE;
   BenchUut2.washComplete := FALSE;
   BenchUut2.weightComplete := FALSE;
   BenchUut2.weight := REAL#0.0;
   BenchUut2.firingComplete := TRUE;
   TraceIn_Mode[22] := BenchUut2.Mode;
   TraceIn_ForwardButton[22] := BenchUut2.ForwardButton;
   TraceIn_ReverseButton[22] := BenchUut2.ReverseButton;
   TraceIn_SensorFeed[22] := BenchUut2.SensorFeed;
   TraceIn_SensorWash[22] := BenchUut2.SensorWash;
   TraceIn_SensorWeight[22] := BenchUut2.SensorWeight;
   TraceIn_SensorFiring[22] := BenchUut2.SensorFiring;
   TraceIn_SensorOutput[22] := BenchUut2.SensorOutput;
   TraceIn_washComplete[22] := BenchUut2.washComplete;
   TraceIn_weightComplete[22] := BenchUut2.weightComplete;
   TraceIn_weight[22] := BenchUut2.weight;
   TraceIn_firingComplete[22] := BenchUut2.firingComplete;
   BenchUut2();
   TraceOut_MotorForward[22] := BenchUut2.MotorForward;
   TraceOut_MotorReverse[22] := BenchUut2.MotorReverse;
   TraceOut_kick[22] := BenchUut2.kick;
   TraceOut_CompletionLight[22] := BenchUut2.CompletionLight;
   TraceOut_firingTemp[22] := BenchUut2.firingTemp;
   BenchCalls := BenchCalls + 1;
 23:
   BenchUut2.Mode := TRUE;
   BenchUut2.ForwardButton := FALSE;
   BenchUut2.ReverseButton := FALSE;
   BenchUut2.SensorFeed := FALSE;
   BenchUut2.SensorWash := FALSE;
   BenchUut2.SensorWeight := FALSE;
   BenchUut2.SensorFiring := FALSE;
   BenchUut2.SensorOutput := TRUE;
   BenchUut2.washComplete := FALSE;
   BenchUut2.weightComplete := FALSE;
   BenchUut2.weight := REAL#0.0;
   BenchUut2.firingComplete := FALSE;
   TraceIn_Mode[23] := BenchUut2.Mode;
   TraceIn_ForwardButton[23] := BenchUut2.ForwardButton;
   TraceIn_ReverseButton[23] := BenchUut2.ReverseButton;
   TraceIn_SensorFeed[23] := BenchUut2.SensorFeed;
   TraceIn_SensorWash[23] := BenchUut2.SensorWash;
   TraceIn_SensorWeight[23] := BenchUut2.SensorWeight;
   TraceIn_SensorFiring[23] := BenchUut2.SensorFiring;
   TraceIn_SensorOutput[23] := BenchUut2.SensorOutput;
   TraceIn_washComplete[23] := BenchUut2.washComplete;
   TraceIn_weightComplete[23] := BenchUut2.weightComplete;
   TraceIn_weight[23] := BenchUut2.weight;
   TraceIn_firingComplete[23] := BenchUut2.firingComplete;
   BenchUut2();
   TraceOut_MotorForward[23] := BenchUut2.MotorForward;
   TraceOut_MotorReverse[23] := BenchUut2.MotorReverse;
   TraceOut_kick[23] := BenchUut2.kick;
   TraceOut_CompletionLight[23] := BenchUut2.CompletionLight;
   TraceOut_firingTemp[23] := BenchUut2.firingTemp;
   BenchCalls := BenchCalls + 1;
 24:
   BenchUut2.Mode := TRUE;
   BenchUut2.ForwardButton := FALSE;
   BenchUut2.ReverseButton := FALSE;
   BenchUut2.SensorFeed := FALSE;
   BenchUut2.SensorWash := FALSE;
   BenchUut2.SensorWeight := FALSE;
   BenchUut2.SensorFiring := FALSE;
   BenchUut2.SensorOutput := TRUE;
   BenchUut2.washComplete := FALSE;
   BenchUut2.weightComplete := FALSE;
   BenchUut2.weight := REAL#0.0;
   BenchUut2.firingComplete := FALSE;
   TraceIn_Mode[24] := BenchUut2.Mode;
   TraceIn_ForwardButton[24] := BenchUut2.ForwardButton;
   TraceIn_ReverseButton[24] := BenchUut2.ReverseButton;
   TraceIn_SensorFeed[24] := BenchUut2.SensorFeed;
   TraceIn_SensorWash[24] := BenchUut2.SensorWash;
   TraceIn_SensorWeight[24] := BenchUut2.SensorWeight;
   TraceIn_SensorFiring[24] := BenchUut2.SensorFiring;
   TraceIn_SensorOutput[24] := BenchUut2.SensorOutput;
   TraceIn_washComplete[24] := BenchUut2.washComplete;
   TraceIn_weightComplete[24] := BenchUut2.weightComplete;
   TraceIn_weight[24] := BenchUut2.weight;
   TraceIn_firingComplete[24] := BenchUut2.firingComplete;
   BenchUut2();
   TraceOut_MotorForward[24] := BenchUut2.MotorForward;
   TraceOut_MotorReverse[24] := BenchUut2.MotorReverse;
   TraceOut_kick[24] := BenchUut2.kick;
   TraceOut_CompletionLight[24] := BenchUut2.CompletionLight;
   TraceOut_firingTemp[24] := BenchUut2.firingTemp;
   BenchCalls := BenchCalls + 1;
 25:
   BenchUut2.Mode := TRUE;
   BenchUut2.ForwardButton := FALSE;
   BenchUut2.ReverseButton := FALSE;
   BenchUut2.SensorFeed := FALSE;
   BenchUut2.SensorWash := FALSE;
   BenchUut2.SensorWeight := FALSE;
   BenchUut2.SensorFiring := FALSE;
   BenchUut2.SensorOutput := FALSE;
   BenchUut2.washComplete := FALSE;
   BenchUut2.weightComplete := FALSE;
   BenchUut2.weight := REAL#0.0;
   BenchUut2.firingComplete := FALSE;
   TraceIn_Mode[25] := BenchUut2.Mode;
   TraceIn_ForwardButton[25] := BenchUut2.ForwardButton;
   TraceIn_ReverseButton[25] := BenchUut2.ReverseButton;
   TraceIn_SensorFeed[25] := BenchUut2.SensorFeed;
   TraceIn_SensorWash[25] := BenchUut2.SensorWash;
   TraceIn_SensorWeight[25] := BenchUut2.SensorWeight;
   TraceIn_SensorFiring[25] := BenchUut2.SensorFiring;
   TraceIn_SensorOutput[25] := BenchUut2.SensorOutput;
   TraceIn_washComplete[25] := BenchUut2.washComplete;
   TraceIn_weightComplete[25] := BenchUut2.weightComplete;
   TraceIn_weight[25] := BenchUut2.weight;
   TraceIn_firingComplete[25] := BenchUut2.firingComplete;
   BenchUut2();
   TraceOut_MotorForward[25] := BenchUut2.MotorForward;
   TraceOut_MotorReverse[25] := BenchUut2.MotorReverse;
   TraceOut_kick[25] := BenchUut2.kick;
   TraceOut_CompletionLight[25] := BenchUut2.CompletionLight;
   TraceOut_firingTemp[25] := BenchUut2.firingTemp;
   BenchCalls := BenchCalls + 1;
 26:
   BenchUut3.Mode := TRUE;
   BenchUut3.ForwardButton := FALSE;
   BenchUut3.ReverseButton := FALSE;
   BenchUut3.SensorFeed := FALSE;
   BenchUut3.SensorWash := FALSE;
   BenchUut3.SensorWeight := FALSE;
   BenchUut3.SensorFiring := FALSE;
   BenchUut3.SensorOutput := FALSE;
   BenchUut3.washComplete := FALSE;
   BenchUut3.weightComplete := FALSE;
   BenchUut3.weight := REAL#0.0;
   BenchUut3.firingComplete := FALSE;
   TraceIn_Mode[26] := BenchUut3.Mode;
   TraceIn_ForwardButton[26] := BenchUut3.ForwardButton;
   TraceIn_ReverseButton[26] := BenchUut3.ReverseButton;
   TraceIn_SensorFeed[26] := BenchUut3.SensorFeed;
   TraceIn_SensorWash[26] := BenchUut3.SensorWash;
   TraceIn_SensorWeight[26] := BenchUut3.SensorWeight;
   TraceIn_SensorFiring[26] := BenchUut3.SensorFiring;
   TraceIn_SensorOutput[26] := BenchUut3.SensorOutput;
   TraceIn_washComplete[26] := BenchUut3.washComplete;
   TraceIn_weightComplete[26] := BenchUut3.weightComplete;
   TraceIn_weight[26] := BenchUut3.weight;
   TraceIn_firingComplete[26] := BenchUut3.firingComplete;
   BenchUut3();
   TraceOut_MotorForward[26] := BenchUut3.MotorForward;
   TraceOut_MotorReverse[26] := BenchUut3.MotorReverse;
   TraceOut_kick[26] := BenchUut3.kick;
   TraceOut_CompletionLight[26] := BenchUut3.CompletionLight;
   TraceOut_firingTemp[26] := BenchUut3.firingTemp;
   BenchCalls := BenchCalls + 1;
 27:
   BenchUut3.Mode := TRUE;
   BenchUut3.ForwardButton := FALSE;
   BenchUut3.ReverseButton := FALSE;
   BenchUut3.SensorFeed := TRUE;
   BenchUut3.SensorWash := FALSE;
   BenchUut3.SensorWeight := FALSE;
   BenchUut3.SensorFiring := FALSE;
   BenchUut3.SensorOutput := FALSE;
   BenchUut3.washComplete := FALSE;
   BenchUut3.weightComplete := FALSE;
   BenchUut3.weight := REAL#0.0;
   BenchUut3.firingComplete := FALSE;
   TraceIn_Mode[27] := BenchUut3.Mode;
   TraceIn_ForwardButton[27] := BenchUut3.ForwardButton;
   TraceIn_ReverseButton[27] := BenchUut3.ReverseButton;
   TraceIn_SensorFeed[27] := BenchUut3.SensorFeed;
   TraceIn_SensorWash[27] := BenchUut3.SensorWash;
   TraceIn_SensorWeight[27] := BenchUut3.SensorWeight;
   TraceIn_SensorFiring[27] := BenchUut3.SensorFiring;
   TraceIn_SensorOutput[27] := BenchUut3.SensorOutput;
   TraceIn_washComplete[27] := BenchUut3.washComplete;
   TraceIn_weightComplete[27] := BenchUut3.weightComplete;
   TraceIn_weight[27] := BenchUut3.weight;
   TraceIn_firingComplete[27] := BenchUut3.firingComplete;
   BenchUut3();
   TraceOut_MotorForward[27] := BenchUut3.MotorForward;
   TraceOut_MotorReverse[27] := BenchUut3.MotorReverse;
   TraceOut_kick[27] := BenchUut3.kick;
   TraceOut_CompletionLight[27] := BenchUut3.CompletionLight;
   TraceOut_firingTemp[27] := BenchUut3.firingTemp;
   BenchCalls := BenchCalls + 1;
 28:
   BenchUut3.Mode := TRUE;
   BenchUut3.ForwardButton := FALSE;
   BenchUut3.ReverseButton := FALSE;
   BenchUut3.SensorFeed := FALSE;
   BenchUut3.SensorWash := TRUE;
   BenchUut3.SensorWeight := FALSE;
   BenchUut3.SensorFiring := FALSE;
   BenchUut3.SensorOutput := FALSE;
   BenchUut3.washComplete := FALSE;
   BenchUut3.weightComplete := FALSE;
   BenchUut3.weight := REAL#0.0;
   BenchUut3.firingComplete := FALSE;
   TraceIn_Mode[28] := BenchUut3.Mode;
   TraceIn_ForwardButton[28] := BenchUut3.ForwardButton;
   TraceIn_ReverseButton[28] := BenchUut3.ReverseButton;
   TraceIn_SensorFeed[28] := BenchUut3.SensorFeed;
   TraceIn_SensorWash[28] := BenchUut3.SensorWash;
   TraceIn_SensorWeight[28] := BenchUut3.SensorWeight;
   TraceIn_SensorFiring[28] := BenchUut3.SensorFiring;
   TraceIn_SensorOutput[28] := BenchUut3.SensorOutput;
   TraceIn_washComplete[28] := BenchUut3.washComplete;
   TraceIn_weightComplete[28] := BenchUut3.weightComplete;
   TraceIn_weight[28] := BenchUut3.weight;
   TraceIn_firingComplete[28] := BenchUut3.firingComplete;
   BenchUut3();
   TraceOut_MotorForward[28] := BenchUut3.MotorForward;
   TraceOut_MotorReverse[28] := BenchUut3.MotorReverse;
   TraceOut_kick[28] := BenchUut3.kick;
   TraceOut_CompletionLight[28] := BenchUut3.CompletionLight;
   TraceOut_firingTemp[28] := BenchUut3.firingTemp;
   BenchCalls := BenchCalls + 1;
 29:
   BenchUut3.Mode := TRUE;
   BenchUut3.ForwardButton := FALSE;
   BenchUut3.ReverseButton := FALSE;
   BenchUut3.SensorFeed := FALSE;
   BenchUut3.SensorWash := TRUE;
   BenchUut3.SensorWeight := FALSE;
   BenchUut3.SensorFiring := FALSE;
   BenchUut3.SensorOutput := FALSE;
   BenchUut3.washComplete := TRUE;
   BenchUut3.weightComplete := FALSE;
   BenchUut3.weight := REAL#0.0;
   BenchUut3.firingComplete := FALSE;
   TraceIn_Mode[29] := BenchUut3.Mode;
   TraceIn_ForwardButton[29] := BenchUut3.ForwardButton;
   TraceIn_ReverseButton[29] := BenchUut3.ReverseButton;
   TraceIn_SensorFeed[29] := BenchUut3.SensorFeed;
   TraceIn_SensorWash[29] := BenchUut3.SensorWash;
   TraceIn_SensorWeight[29] := BenchUut3.SensorWeight;
   TraceIn_SensorFiring[29] := BenchUut3.SensorFiring;
   TraceIn_SensorOutput[29] := BenchUut3.SensorOutput;
   TraceIn_washComplete[29] := BenchUut3.washComplete;
   TraceIn_weightComplete[29] := BenchUut3.weightComplete;
   TraceIn_weight[29] := BenchUut3.weight;
   TraceIn_firingComplete[29] := BenchUut3.firingComplete;
   BenchUut3();
   TraceOut_MotorForward[29] := BenchUut3.MotorForward;
   TraceOut_MotorReverse[29] := BenchUut3.MotorReverse;
   TraceOut_kick[29] := BenchUut3.kick;
   TraceOut_CompletionLight[29] := BenchUut3.CompletionLight;
   TraceOut_firingTemp[29] := BenchUut3.firingTemp;
   BenchCalls := BenchCalls + 1;
 30:
   BenchUut3.Mode := TRUE;
   BenchUut3.ForwardButton := FALSE;
   BenchUut3.ReverseButton := FALSE;
   BenchUut3.SensorFeed := FALSE;
   BenchUut3.SensorWash := FALSE;
   BenchUut3.SensorWeight := TRUE;
   BenchUut3.SensorFiring := FALSE;
   BenchUut3.SensorOutput := FALSE;
   BenchUut3.washComplete := FALSE;
   BenchUut3.weightComplete := FALSE;
   BenchUut3.weight := REAL#0.0;
   BenchUut3.firingComplete := FALSE;
   TraceIn_Mode[30] := BenchUut3.Mode;
   TraceIn_ForwardButton[30] := BenchUut3.ForwardButton;
   TraceIn_ReverseButton[30] := BenchUut3.ReverseButton;
   TraceIn_SensorFeed[30] := BenchUut3.SensorFeed;
   TraceIn_SensorWash[30] := BenchUut3.SensorWash;
   TraceIn_SensorWeight[30] := BenchUut3.SensorWeight;
   TraceIn_SensorFiring[30] := BenchUut3.SensorFiring;
   TraceIn_SensorOutput[30] := BenchUut3.SensorOutput;
   TraceIn_washComplete[30] := BenchUut3.washComplete;
   TraceIn_weightComplete[30] := BenchUut3.weightComplete;
   TraceIn_weight[30] := BenchUut3.weight;
   TraceIn_firingComplete[30] := BenchUut3.firingComplete;
   BenchUut3();
   TraceOut_MotorForward[30] := BenchUut3.MotorForward;
   TraceOut_MotorReverse[30] := BenchUut3.MotorReverse;
   TraceOut_kick[30] := BenchUut3.kick;
   TraceOut_CompletionLight[30] := BenchUut3.CompletionLight;
   TraceOut_firingTemp[30] := BenchUut3.firingTemp;
   BenchCalls := BenchCalls + 1;
 31:
   BenchUut3.Mode := TRUE;
   BenchUut3.ForwardButton := FALSE;
   BenchUut3.ReverseButton := FALSE;
   BenchUut3.SensorFeed := FALSE;
   BenchUut3.SensorWash := FALSE;
   BenchUut3.SensorWeight := TRUE;
   BenchUut3.SensorFiring := FALSE;
   BenchUut3.SensorOutput := FALSE;
   BenchUut3.washComplete := FALSE;
   BenchUut3.weightComplete := TRUE;
   BenchUut3.weight := REAL#200.0;
   BenchUut3.firingComplete := FALSE;
   TraceIn_Mode[31] := BenchUut3.Mode;
   TraceIn_ForwardButton[31] := BenchUut3.ForwardButton;
   TraceIn_ReverseButton[31] := BenchUut3.ReverseButton;
   TraceIn_SensorFeed[31] := BenchUut3.SensorFeed;
   TraceIn_SensorWash[31] := BenchUut3.SensorWash;
   TraceIn_SensorWeight[31] := BenchUut3.SensorWeight;
   TraceIn_SensorFiring[31] := BenchUut3.SensorFiring;
   TraceIn_SensorOutput[31] := BenchUut3.SensorOutput;
   TraceIn_washComplete[31] := BenchUut3.washComplete;
   TraceIn_weightComplete[31] := BenchUut3.weightComplete;
   TraceIn_weight[31] := BenchUut3.weight;
   TraceIn_firingComplete[31] := BenchUut3.firingComplete;
   BenchUut3();
   TraceOut_MotorForward[31] := BenchUut3.MotorForward;
   TraceOut_MotorReverse[31] := BenchUut3.MotorReverse;
   TraceOut_kick[31] := BenchUut3.kick;
   TraceOut_CompletionLight[31] := BenchUut3.CompletionLight;
   TraceOut_firingTemp[31] := BenchUut3.firingTemp;
   BenchCalls := BenchCalls + 1;
 32:
   BenchUut3.Mode := TRUE;
   BenchUut3.ForwardButton := FALSE;
   BenchUut3.ReverseButton := FALSE;
   BenchUut3.SensorFeed := FALSE;
   BenchUut3.SensorWash := FALSE;
   BenchUut3.SensorWeight := FALSE;
   BenchUut3.SensorFiring := TRUE;
   BenchUut3.SensorOutput := FALSE;
   BenchUut3.washComplete := FALSE;
   BenchUut3.weightComplete := FALSE;
   BenchUut3.weight := REAL#0.0;
   BenchUut3.firingComplete := FALSE;
   TraceIn_Mode[32] := BenchUut3.Mode;
   TraceIn_ForwardButton[32] := BenchUut3.ForwardButton;
   TraceIn_ReverseButton[32] := BenchUut3.ReverseButton;
   TraceIn_SensorFeed[32] := BenchUut3.SensorFeed;
   TraceIn_SensorWash[32] := BenchUut3.SensorWash;
   TraceIn_SensorWeight[32] := BenchUut3.SensorWeight;
   TraceIn_SensorFiring[32] := BenchUut3.SensorFiring;
   TraceIn_SensorOutput[32] := BenchUut3.SensorOutput;
   TraceIn_washComplete[32] := BenchUut3.washComplete;
   TraceIn_weightComplete[32] := BenchUut3.weightComplete;
   TraceIn_weight[32] := BenchUut3.weight;
   TraceIn_firingComplete[32] := BenchUut3.firingComplete;
   BenchUut3();
   TraceOut_MotorForward[32] := BenchUut3.MotorForward;
   TraceOut_MotorReverse[32] := BenchUut3.MotorReverse;
   TraceOut_kick[32] := BenchUut3.kick;
   TraceOut_CompletionLight[32] := BenchUut3.CompletionLight;
   TraceOut_firingTemp[32] := BenchUut3.firingTemp;
   BenchCalls := BenchCalls + 1;
 33:
   BenchUut3.Mode := TRUE;
   BenchUut3.ForwardButton := FALSE;
   BenchUut3.ReverseButton := FALSE;
   BenchUut3.SensorFeed := FALSE;
   BenchUut3.SensorWash := FALSE;
   BenchUut3.SensorWeight := FALSE;
   BenchUut3.SensorFiring := TRUE;
   BenchUut3.SensorOutput := FALSE;
   BenchUut3.washComplete := FALSE;
   BenchUut3.weightComplete := FALSE;
   BenchUut3.weight := REAL#0.0;
   BenchUut3.firingComplete := TRUE;
   TraceIn_Mode[33] := BenchUut3.Mode;
   TraceIn_ForwardButton[33] := BenchUut3.ForwardButton;
   TraceIn_ReverseButton[33] := BenchUut3.ReverseButton;
   TraceIn_SensorFeed[33] := BenchUut3.SensorFeed;
   TraceIn_SensorWash[33] := BenchUut3.SensorWash;
   TraceIn_SensorWeight[33] := BenchUut3.SensorWeight;
   TraceIn_SensorFiring[33] := BenchUut3.SensorFiring;
   TraceIn_SensorOutput[33] := BenchUut3.SensorOutput;
   TraceIn_washComplete[33] := BenchUut3.washComplete;
   TraceIn_weightComplete[33] := BenchUut3.weightComplete;
   TraceIn_weight[33] := BenchUut3.weight;
   TraceIn_firingComplete[33] := BenchUut3.firingComplete;
   BenchUut3();
   TraceOut_MotorForward[33] := BenchUut3.MotorForward;
   TraceOut_MotorReverse[33] := BenchUut3.MotorReverse;
   TraceOut_kick[33] := BenchUut3.kick;
   TraceOut_CompletionLight[33] := BenchUut3.CompletionLight;
   TraceOut_firingTemp[33] := BenchUut3.firingTemp;
   BenchCalls := BenchCalls + 1;
 34:
   BenchUut3.Mode := TRUE;
   BenchUut3.ForwardButton := FALSE;
   BenchUut3.ReverseButton := FALSE;
   BenchUut3.SensorFeed := FALSE;
   BenchUut3.SensorWash := FALSE;
   BenchUut3.SensorWeight := FALSE;
   BenchUut3.SensorFiring := FALSE;
   BenchUut3.SensorOutput := TRUE;
   BenchUut3.washComplete := FALSE;
   BenchUut3.weightComplete := FALSE;
   BenchUut3.weight := REAL#0.0;
   BenchUut3.firingComplete := FALSE;
   TraceIn_Mode[34] := BenchUut3.Mode;
   TraceIn_ForwardButton[34] := BenchUut3.ForwardButton;
   TraceIn_ReverseButton[34] := BenchUut3.ReverseButton;
   TraceIn_SensorFeed[34] := BenchUut3.SensorFeed;
   TraceIn_SensorWash[34] := BenchUut3.SensorWash;
   TraceIn_SensorWeight[34] := BenchUut3.SensorWeight;
   TraceIn_SensorFiring[34] := BenchUut3.SensorFiring;
   TraceIn_SensorOutput[34] := BenchUut3.SensorOutput;
   TraceIn_washComplete[34] := BenchUut3.washComplete;
   TraceIn_weightComplete[34] := BenchUut3.weightComplete;
   TraceIn_weight[34] := BenchUut3.weight;
   TraceIn_firingComplete[34] := BenchUut3.firingComplete;
   BenchUut3();
   TraceOut_MotorForward[34] := BenchUut3.MotorForward;
   TraceOut_MotorReverse[34] := BenchUut3.MotorReverse;
   TraceOut_kick[34] := BenchUut3.kick;
   TraceOut_CompletionLight[34] := BenchUut3.CompletionLight;
   TraceOut_firingTemp[34] := BenchUut3.firingTemp;
   BenchCalls := BenchCalls + 1;
 35:
   BenchUut3.Mode := TRUE;
   BenchUut3.ForwardButton := FALSE;
   BenchUut3.ReverseButton := FALSE;
   BenchUut3.SensorFeed := FALSE;
   BenchUut3.SensorWash := FALSE;
   BenchUut3.SensorWeight := FALSE;
   BenchUut3.SensorFiring := FALSE;
   BenchUut3.SensorOutput := TRUE;
   BenchUut3.washComplete := FALSE;
   BenchUut3.weightComplete := FALSE;
   BenchUut3.weight := REAL#0.0;
   BenchUut3.firingComplete := FALSE;
   TraceIn_Mode[35] := BenchUut3.Mode;
   TraceIn_ForwardButton[35] := BenchUut3.ForwardButton;
   TraceIn_ReverseButton[35] := BenchUut3.ReverseButton;
   TraceIn_SensorFeed[35] := BenchUut3.SensorFeed;
   TraceIn_SensorWash[35] := BenchUut3.SensorWash;
   TraceIn_SensorWeight[35] := BenchUut3.SensorWeight;
   TraceIn_SensorFiring[35] := BenchUut3.SensorFiring;
   TraceIn_SensorOutput[35] := BenchUut3.SensorOutput;
   TraceIn_washComplete[35] := BenchUut3.washComplete;
   TraceIn_weightComplete[35] := BenchUut3.weightComplete;
   TraceIn_weight[35] := BenchUut3.weight;
   TraceIn_firingComplete[35] := BenchUut3.firingComplete;
   BenchUut3();
   TraceOut_MotorForward[35] := BenchUut3.MotorForward;
   TraceOut_MotorReverse[35] := BenchUut3.MotorReverse;
   TraceOut_kick[35] := BenchUut3.kick;
   TraceOut_CompletionLight[35] := BenchUut3.CompletionLight;
   TraceOut_firingTemp[35] := BenchUut3.firingTemp;
   BenchCalls := BenchCalls + 1;
 36:
   BenchUut3.Mode := TRUE;
   BenchUut3.ForwardButton := FALSE;
   BenchUut3.ReverseButton := FALSE;
   BenchUut3.SensorFeed := FALSE;
   BenchUut3.SensorWash := FALSE;
   BenchUut3.SensorWeight := FALSE;
   BenchUut3.SensorFiring := FALSE;
   BenchUut3.SensorOutput := FALSE;
   BenchUut3.washComplete := FALSE;
   BenchUut3.weightComplete := FALSE;
   BenchUut3.weight := REAL#0.0;
   BenchUut3.firingComplete := FALSE;
   TraceIn_Mode[36] := BenchUut3.Mode;
   TraceIn_ForwardButton[36] := BenchUut3.ForwardButton;
   TraceIn_ReverseButton[36] := BenchUut3.ReverseButton;
   TraceIn_SensorFeed[36] := BenchUut3.SensorFeed;
   TraceIn_SensorWash[36] := BenchUut3.SensorWash;
   TraceIn_SensorWeight[36] := BenchUut3.SensorWeight;
   TraceIn_SensorFiring[36] := BenchUut3.SensorFiring;
   TraceIn_SensorOutput[36] := BenchUut3.SensorOutput;
   TraceIn_washComplete[36] := BenchUut3.washComplete;
   TraceIn_weightComplete[36] := BenchUut3.weightComplete;
   TraceIn_weight[36] := BenchUut3.weight;
   TraceIn_firingComplete[36] := BenchUut3.firingComplete;
   BenchUut3();
   TraceOut_MotorForward[36] := BenchUut3.MotorForward;
   TraceOut_MotorReverse[36] := BenchUut3.MotorReverse;
   TraceOut_kick[36] := BenchUut3.kick;
   TraceOut_CompletionLight[36] := BenchUut3.CompletionLight;
   TraceOut_firingTemp[36] := BenchUut3.firingTemp;
   BenchCalls := BenchCalls + 1;
 37:
   BenchUut4.Mode := TRUE;
   BenchUut4.ForwardButton := FALSE;
   BenchUut4.ReverseButton := FALSE;
   BenchUut4.SensorFeed := FALSE;
   BenchUut4.SensorWash := FALSE;
   BenchUut4.SensorWeight := FALSE;
   BenchUut4.SensorFiring := FALSE;
   BenchUut4.SensorOutput := FALSE;
   BenchUut4.washComplete := FALSE;
   BenchUut4.weightComplete := FALSE;
   BenchUut4.weight := REAL#0.0;
   BenchUut4.firingComplete := FALSE;
   TraceIn_Mode[37] := BenchUut4.Mode;
   TraceIn_ForwardButton[37] := BenchUut4.ForwardButton;
   TraceIn_ReverseButton[37] := BenchUut4.ReverseButton;
   TraceIn_SensorFeed[37] := BenchUut4.SensorFeed;
   TraceIn_SensorWash[37] := BenchUut4.SensorWash;
   TraceIn_SensorWeight[37] := BenchUut4.SensorWeight;
   TraceIn_SensorFiring[37] := BenchUut4.SensorFiring;
   TraceIn_SensorOutput[37] := BenchUut4.SensorOutput;
   TraceIn_washComplete[37] := BenchUut4.washComplete;
   TraceIn_weightComplete[37] := BenchUut4.weightComplete;
   TraceIn_weight[37] := BenchUut4.weight;
   TraceIn_firingComplete[37] := BenchUut4.firingComplete;
   BenchUut4();
   TraceOut_MotorForward[37] := BenchUut4.MotorForward;
   TraceOut_MotorReverse[37] := BenchUut4.MotorReverse;
   TraceOut_kick[37] := BenchUut4.kick;
   TraceOut_CompletionLight[37] := BenchUut4.CompletionLight;
   TraceOut_firingTemp[37] := BenchUut4.firingTemp;
   BenchCalls := BenchCalls + 1;
 38:
   BenchUut4.Mode := TRUE;
   BenchUut4.ForwardButton := FALSE;
   BenchUut4.ReverseButton := FALSE;
   BenchUut4.SensorFeed := TRUE;
   BenchUut4.SensorWash := FALSE;
   BenchUut4.SensorWeight := FALSE;
   BenchUut4.SensorFiring := FALSE;
   BenchUut4.SensorOutput := FALSE;
   BenchUut4.washComplete := FALSE;
   BenchUut4.weightComplete := FALSE;
   BenchUut4.weight := REAL#0.0;
   BenchUut4.firingComplete := FALSE;
   TraceIn_Mode[38] := BenchUut4.Mode;
   TraceIn_ForwardButton[38] := BenchUut4.ForwardButton;
   TraceIn_ReverseButton[38] := BenchUut4.ReverseButton;
   TraceIn_SensorFeed[38] := BenchUut4.SensorFeed;
   TraceIn_SensorWash[38] := BenchUut4.SensorWash;
   TraceIn_SensorWeight[38] := BenchUut4.SensorWeight;
   TraceIn_SensorFiring[38] := BenchUut4.SensorFiring;
   TraceIn_SensorOutput[38] := BenchUut4.SensorOutput;
   TraceIn_washComplete[38] := BenchUut4.washComplete;
   TraceIn_weightComplete[38] := BenchUut4.weightComplete;
   TraceIn_weight[38] := BenchUut4.weight;
   TraceIn_firingComplete[38] := BenchUut4.firingComplete;
   BenchUut4();
   TraceOut_MotorForward[38] := BenchUut4.MotorForward;
   TraceOut_MotorReverse[38] := BenchUut4.MotorReverse;
   TraceOut_kick[38] := BenchUut4.kick;
   TraceOut_CompletionLight[38] := BenchUut4.CompletionLight;
   TraceOut_firingTemp[38] := BenchUut4.firingTemp;
   BenchCalls := BenchCalls + 1;
 39:
   BenchUut4.Mode := TRUE;
   BenchUut4.ForwardButton := FALSE;
   BenchUut4.ReverseButton := FALSE;
   BenchUut4.SensorFeed := FALSE;
   BenchUut4.SensorWash := TRUE;
   BenchUut4.SensorWeight := FALSE;
   BenchUut4.SensorFiring := FALSE;
   BenchUut4.SensorOutput := FALSE;
   BenchUut4.washComplete := FALSE;
   BenchUut4.weightComplete := FALSE;
   BenchUut4.weight := REAL#0.0;
   BenchUut4.firingComplete := FALSE;
   TraceIn_Mode[39] := BenchUut4.Mode;
   TraceIn_ForwardButton[39] := BenchUut4.ForwardButton;
   TraceIn_ReverseButton[39] := BenchUut4.ReverseButton;
   TraceIn_SensorFeed[39] := BenchUut4.SensorFeed;
   TraceIn_SensorWash[39] := BenchUut4.SensorWash;
   TraceIn_SensorWeight[39] := BenchUut4.SensorWeight;
   TraceIn_SensorFiring[39] := BenchUut4.SensorFiring;
   TraceIn_SensorOutput[39] := BenchUut4.SensorOutput;
   TraceIn_washComplete[39] := BenchUut4.washComplete;
   TraceIn_weightComplete[39] := BenchUut4.weightComplete;
   TraceIn_weight[39] := BenchUut4.weight;
   TraceIn_firingComplete[39] := BenchUut4.firingComplete;
   BenchUut4();
   TraceOut_MotorForward[39] := BenchUut4.MotorForward;
   TraceOut_MotorReverse[39] := BenchUut4.MotorReverse;
   TraceOut_kick[39] := BenchUut4.kick;
   TraceOut_CompletionLight[39] := BenchUut4.CompletionLight;
   TraceOut_firingTemp[39] := BenchUut4.firingTemp;
   BenchCalls := BenchCalls + 1;
 40:
   BenchUut4.Mode := TRUE;
   BenchUut4.ForwardButton := FALSE;
   BenchUut4.ReverseButton := FALSE;
   BenchUut4.SensorFeed := FALSE;
   BenchUut4.SensorWash := TRUE;
   BenchUut4.SensorWeight := FALSE;
   BenchUut4.SensorFiring := FALSE;
   BenchUut4.SensorOutput := FALSE;
   BenchUut4.washComplete := TRUE;
   BenchUut4.weightComplete := FALSE;
   BenchUut4.weight := REAL#0.0;
   BenchUut4.firingComplete := FALSE;
   TraceIn_Mode[40] := BenchUut4.Mode;
   TraceIn_ForwardButton[40] := BenchUut4.ForwardButton;
   TraceIn_ReverseButton[40] := BenchUut4.ReverseButton;
   TraceIn_SensorFeed[40] := BenchUut4.SensorFeed;
   TraceIn_SensorWash[40] := BenchUut4.SensorWash;
   TraceIn_SensorWeight[40] := BenchUut4.SensorWeight;
   TraceIn_SensorFiring[40] := BenchUut4.SensorFiring;
   TraceIn_SensorOutput[40] := BenchUut4.SensorOutput;
   TraceIn_washComplete[40] := BenchUut4.washComplete;
   TraceIn_weightComplete[40] := BenchUut4.weightComplete;
   TraceIn_weight[40] := BenchUut4.weight;
   TraceIn_firingComplete[40] := BenchUut4.firingComplete;
   BenchUut4();
   TraceOut_MotorForward[40] := BenchUut4.MotorForward;
   TraceOut_MotorReverse[40] := BenchUut4.MotorReverse;
   TraceOut_kick[40] := BenchUut4.kick;
   TraceOut_CompletionLight[40] := BenchUut4.CompletionLight;
   TraceOut_firingTemp[40] := BenchUut4.firingTemp;
   BenchCalls := BenchCalls + 1;
 41:
   BenchUut4.Mode := TRUE;
   BenchUut4.ForwardButton := FALSE;
   BenchUut4.ReverseButton := FALSE;
   BenchUut4.SensorFeed := FALSE;
   BenchUut4.SensorWash := FALSE;
   BenchUut4.SensorWeight := TRUE;
   BenchUut4.SensorFiring := FALSE;
   BenchUut4.SensorOutput := FALSE;
   BenchUut4.washComplete := FALSE;
   BenchUut4.weightComplete := FALSE;
   BenchUut4.weight := REAL#0.0;
   BenchUut4.firingComplete := FALSE;
   TraceIn_Mode[41] := BenchUut4.Mode;
   TraceIn_ForwardButton[41] := BenchUut4.ForwardButton;
   TraceIn_ReverseButton[41] := BenchUut4.ReverseButton;
   TraceIn_SensorFeed[41] := BenchUut4.SensorFeed;
   TraceIn_SensorWash[41] := BenchUut4.SensorWash;
   TraceIn_SensorWeight[41] := BenchUut4.SensorWeight;
   TraceIn_SensorFiring[41] := BenchUut4.SensorFiring;
   TraceIn_SensorOutput[41] := BenchUut4.SensorOutput;
   TraceIn_washComplete[41] := BenchUut4.washComplete;
   TraceIn_weightComplete[41] := BenchUut4.weightComplete;
   TraceIn_weight[41] := BenchUut4.weight;
   TraceIn_firingComplete[41] := BenchUut4.firingComplete;
   BenchUut4();
   TraceOut_MotorForward[41] := BenchUut4.MotorForward;
   TraceOut_MotorReverse[41] := BenchUut4.MotorReverse;
   TraceOut_kick[41] := BenchUut4.kick;
   TraceOut_CompletionLight[41] := BenchUut4.CompletionLight;
   TraceOut_firingTemp[41] := BenchUut4.firingTemp;
   BenchCalls := BenchCalls + 1;
 42:
   BenchUut4.Mode := TRUE;
   BenchUut4.ForwardButton := FALSE;
   BenchUut4.ReverseButton := FALSE;
   BenchUut4.SensorFeed := FALSE;
   BenchUut4.SensorWash := FALSE;
   BenchUut4.SensorWeight := TRUE;
   BenchUut4.SensorFiring := FALSE;
   BenchUut4.SensorOutput := FALSE;
   BenchUut4.washComplete := FALSE;
   BenchUut4.weightComplete := TRUE;
   BenchUut4.weight := REAL#99.9;
   BenchUut4.firingComplete := FALSE;
   TraceIn_Mode[42] := BenchUut4.Mode;
   TraceIn_ForwardButton[42] := BenchUut4.ForwardButton;
   TraceIn_ReverseButton[42] := BenchUut4.ReverseButton;
   TraceIn_SensorFeed[42] := BenchUut4.SensorFeed;
   TraceIn_SensorWash[42] := BenchUut4.SensorWash;
   TraceIn_SensorWeight[42] := BenchUut4.SensorWeight;
   TraceIn_SensorFiring[42] := BenchUut4.SensorFiring;
   TraceIn_SensorOutput[42] := BenchUut4.SensorOutput;
   TraceIn_washComplete[42] := BenchUut4.washComplete;
   TraceIn_weightComplete[42] := BenchUut4.weightComplete;
   TraceIn_weight[42] := BenchUut4.weight;
   TraceIn_firingComplete[42] := BenchUut4.firingComplete;
   BenchUut4();
   TraceOut_MotorForward[42] := BenchUut4.MotorForward;
   TraceOut_MotorReverse[42] := BenchUut4.MotorReverse;
   TraceOut_kick[42] := BenchUut4.kick;
   TraceOut_CompletionLight[42] := BenchUut4.CompletionLight;
   TraceOut_firingTemp[42] := BenchUut4.firingTemp;
   BenchCalls := BenchCalls + 1;
 43:
   BenchUut4.Mode := TRUE;
   BenchUut4.ForwardButton := FALSE;
   BenchUut4.ReverseButton := FALSE;
   BenchUut4.SensorFeed := FALSE;
   BenchUut4.SensorWash := FALSE;
   BenchUut4.SensorWeight := TRUE;
   BenchUut4.SensorFiring := FALSE;
   BenchUut4.SensorOutput := FALSE;
   BenchUut4.washComplete := FALSE;
   BenchUut4.weightComplete := FALSE;
   BenchUut4.weight := REAL#0.0;
   BenchUut4.firingComplete := FALSE;
   TraceIn_Mode[43] := BenchUut4.Mode;
   TraceIn_ForwardButton[43] := BenchUut4.ForwardButton;
   TraceIn_ReverseButton[43] := BenchUut4.ReverseButton;
   TraceIn_SensorFeed[43] := BenchUut4.SensorFeed;
   TraceIn_SensorWash[43] := BenchUut4.SensorWash;
   TraceIn_SensorWeight[43] := BenchUut4.SensorWeight;
   TraceIn_SensorFiring[43] := BenchUut4.SensorFiring;
   TraceIn_SensorOutput[43] := BenchUut4.SensorOutput;
   TraceIn_washComplete[43] := BenchUut4.washComplete;
   TraceIn_weightComplete[43] := BenchUut4.weightComplete;
   TraceIn_weight[43] := BenchUut4.weight;
   TraceIn_firingComplete[43] := BenchUut4.firingComplete;
   BenchUut4();
   TraceOut_MotorForward[43] := BenchUut4.MotorForward;
   TraceOut_MotorReverse[43] := BenchUut4.MotorReverse;
   TraceOut_kick[43] := BenchUut4.kick;
   TraceOut_CompletionLight[43] := BenchUut4.CompletionLight;
   TraceOut_firingTemp[43] := BenchUut4.firingTemp;
   BenchCalls := BenchCalls + 1;
 44:
   BenchUut4.Mode := TRUE;
   BenchUut4.ForwardButton := FALSE;
   BenchUut4.ReverseButton := FALSE;
   BenchUut4.SensorFeed := FALSE;
   BenchUut4.SensorWash := FALSE;
   BenchUut4.SensorWeight := FALSE;
   BenchUut4.SensorFiring := FALSE;
   BenchUut4.SensorOutput := FALSE;
   BenchUut4.washComplete := FALSE;
   BenchUut4.weightComplete := FALSE;
   BenchUut4.weight := REAL#0.0;
   BenchUut4.firingComplete := FALSE;
   TraceIn_Mode[44] := BenchUut4.Mode;
   TraceIn_ForwardButton[44] := BenchUut4.ForwardButton;
   TraceIn_ReverseButton[44] := BenchUut4.ReverseButton;
   TraceIn_SensorFeed[44] := BenchUut4.SensorFeed;
   TraceIn_SensorWash[44] := BenchUut4.SensorWash;
   TraceIn_SensorWeight[44] := BenchUut4.SensorWeight;
   TraceIn_SensorFiring[44] := BenchUut4.SensorFiring;
   TraceIn_SensorOutput[44] := BenchUut4.SensorOutput;
   TraceIn_washComplete[44] := BenchUut4.washComplete;
   TraceIn_weightComplete[44] := BenchUut4.weightComplete;
   TraceIn_weight[44] := BenchUut4.weight;
   TraceIn_firingComplete[44] := BenchUut4.firingComplete;
   BenchUut4();
   TraceOut_MotorForward[44] := BenchUut4.MotorForward;
   TraceOut_MotorReverse[44] := BenchUut4.MotorReverse;
   TraceOut_kick[44] := BenchUut4.kick;
   TraceOut_CompletionLight[44] := BenchUut4.CompletionLight;
   TraceOut_firingTemp[44] := BenchUut4.firingTemp;
   BenchCalls := BenchCalls + 1;
 45:
   BenchUut4.Mode := TRUE;
   BenchUut4.ForwardButton := FALSE;
   BenchUut4.ReverseButton := FALSE;
   BenchUut4.SensorFeed := TRUE;
   BenchUut4.SensorWash := FALSE;
   BenchUut4.SensorWeight := FALSE;
   BenchUut4.SensorFiring := FALSE;
   BenchUut4.SensorOutput := FALSE;
   BenchUut4.washComplete := FALSE;
   BenchUut4.weightComplete := FALSE;
   BenchUut4.weight := REAL#0.0;
   BenchUut4.firingComplete := FALSE;
   TraceIn_Mode[45] := BenchUut4.Mode;
   TraceIn_ForwardButton[45] := BenchUut4.ForwardButton;
   TraceIn_ReverseButton[45] := BenchUut4.ReverseButton;
   TraceIn_SensorFeed[45] := BenchUut4.SensorFeed;
   TraceIn_SensorWash[45] := BenchUut4.SensorWash;
   TraceIn_SensorWeight[45] := BenchUut4.SensorWeight;
   TraceIn_SensorFiring[45] := BenchUut4.SensorFiring;
   TraceIn_SensorOutput[45] := BenchUut4.SensorOutput;
   TraceIn_washComplete[45] := BenchUut4.washComplete;
   TraceIn_weightComplete[45] := BenchUut4.weightComplete;
   TraceIn_weight[45] := BenchUut4.weight;
   TraceIn_firingComplete[45] := BenchUut4.firingComplete;
   BenchUut4();
   TraceOut_MotorForward[45] := BenchUut4.MotorForward;
   TraceOut_MotorReverse[45] := BenchUut4.MotorReverse;
   TraceOut_kick[45] := BenchUut4.kick;
   TraceOut_CompletionLight[45] := BenchUut4.CompletionLight;
   TraceOut_firingTemp[45] := BenchUut4.firingTemp;
   BenchCalls := BenchCalls + 1;
 46:
   BenchUut5.Mode := TRUE;
   BenchUut5.ForwardButton := FALSE;
   BenchUut5.ReverseButton := FALSE;
   BenchUut5.SensorFeed := FALSE;
   BenchUut5.SensorWash := FALSE;
   BenchUut5.SensorWeight := FALSE;
   BenchUut5.SensorFiring := FALSE;
   BenchUut5.SensorOutput := FALSE;
   BenchUut5.washComplete := FALSE;
   BenchUut5.weightComplete := FALSE;
   BenchUut5.weight := REAL#0.0;
   BenchUut5.firingComplete := FALSE;
   TraceIn_Mode[46] := BenchUut5.Mode;
   TraceIn_ForwardButton[46] := BenchUut5.ForwardButton;
   TraceIn_ReverseButton[46] := BenchUut5.ReverseButton;
   TraceIn_SensorFeed[46] := BenchUut5.SensorFeed;
   TraceIn_SensorWash[46] := BenchUut5.SensorWash;
   TraceIn_SensorWeight[46] := BenchUut5.SensorWeight;
   TraceIn_SensorFiring[46] := BenchUut5.SensorFiring;
   TraceIn_SensorOutput[46] := BenchUut5.SensorOutput;
   TraceIn_washComplete[46] := BenchUut5.washComplete;
   TraceIn_weightComplete[46] := BenchUut5.weightComplete;
   TraceIn_weight[46] := BenchUut5.weight;
   TraceIn_firingComplete[46] := BenchUut5.firingComplete;
   BenchUut5();
   TraceOut_MotorForward[46] := BenchUut5.MotorForward;
   TraceOut_MotorReverse[46] := BenchUut5.MotorReverse;
   TraceOut_kick[46] := BenchUut5.kick;
   TraceOut_CompletionLight[46] := BenchUut5.CompletionLight;
   TraceOut_firingTemp[46] := BenchUut5.firingTemp;
   BenchCalls := BenchCalls + 1;
 47:
   BenchUut5.Mode := TRUE;
   BenchUut5.ForwardButton := FALSE;
   BenchUut5.ReverseButton := FALSE;
   BenchUut5.SensorFeed := TRUE;
   BenchUut5.SensorWash := FALSE;
   BenchUut5.SensorWeight := FALSE;
   BenchUut5.SensorFiring := FALSE;
   BenchUut5.SensorOutput := FALSE;
   BenchUut5.washComplete := FALSE;
   BenchUut5.weightComplete := FALSE;
   BenchUut5.weight := REAL#0.0;
   BenchUut5.firingComplete := FALSE;
   TraceIn_Mode[47] := BenchUut5.Mode;
   TraceIn_ForwardButton[47] := BenchUut5.ForwardButton;
   TraceIn_ReverseButton[47] := BenchUut5.ReverseButton;
   TraceIn_SensorFeed[47] := BenchUut5.SensorFeed;
   TraceIn_SensorWash[47] := BenchUut5.SensorWash;
   TraceIn_SensorWeight[47] := BenchUut5.SensorWeight;
   TraceIn_SensorFiring[47] := BenchUut5.SensorFiring;
   TraceIn_SensorOutput[47] := BenchUut5.SensorOutput;
   TraceIn_washComplete[47] := BenchUut5.washComplete;
   TraceIn_weightComplete[47] := BenchUut5.weightComplete;
   TraceIn_weight[47] := BenchUut5.weight;
   TraceIn_firingComplete[47] := BenchUut5.firingComplete;
   BenchUut5();
   TraceOut_MotorForward[47] := BenchUut5.MotorForward;
   TraceOut_MotorReverse[47] := BenchUut5.MotorReverse;
   TraceOut_kick[47] := BenchUut5.kick;
   TraceOut_CompletionLight[47] := BenchUut5.CompletionLight;
   TraceOut_firingTemp[47] := BenchUut5.firingTemp;
   BenchCalls := BenchCalls + 1;
 48:
   BenchUut5.Mode := TRUE;
   BenchUut5.ForwardButton := FALSE;
   BenchUut5.ReverseButton := FALSE;
   BenchUut5.SensorFeed := FALSE;
   BenchUut5.SensorWash := TRUE;
   BenchUut5.SensorWeight := FALSE;
   BenchUut5.SensorFiring := FALSE;
   BenchUut5.SensorOutput := FALSE;
   BenchUut5.washComplete := FALSE;
   BenchUut5.weightComplete := FALSE;
   BenchUut5.weight := REAL#0.0;
   BenchUut5.firingComplete := FALSE;
   TraceIn_Mode[48] := BenchUut5.Mode;
   TraceIn_ForwardButton[48] := BenchUut5.ForwardButton;
   TraceIn_ReverseButton[48] := BenchUut5.ReverseButton;
   TraceIn_SensorFeed[48] := BenchUut5.SensorFeed;
   TraceIn_SensorWash[48] := BenchUut5.SensorWash;
   TraceIn_SensorWeight[48] := BenchUut5.SensorWeight;
   TraceIn_SensorFiring[48] := BenchUut5.SensorFiring;
   TraceIn_SensorOutput[48] := BenchUut5.SensorOutput;
   TraceIn_washComplete[48] := BenchUut5.washComplete;
   TraceIn_weightComplete[48] := BenchUut5.weightComplete;
   TraceIn_weight[48] := BenchUut5.weight;
   TraceIn_firingComplete[48] := BenchUut5.firingComplete;
   BenchUut5();
   TraceOut_MotorForward[48] := BenchUut5.MotorForward;
   TraceOut_MotorReverse[48] := BenchUut5.MotorReverse;
   TraceOut_kick[48] := BenchUut5.kick;
   TraceOut_CompletionLight[48] := BenchUut5.CompletionLight;
   TraceOut_firingTemp[48] := BenchUut5.firingTemp;
   BenchCalls := BenchCalls + 1;
 49:
   BenchUut5.Mode := TRUE;
   BenchUut5.ForwardButton := FALSE;
   BenchUut5.ReverseButton := FALSE;
   BenchUut5.SensorFeed := FALSE;
   BenchUut5.SensorWash := TRUE;
   BenchUut5.SensorWeight := FALSE;
   BenchUut5.SensorFiring := FALSE;
   BenchUut5.SensorOutput := FALSE;
   BenchUut5.washComplete := TRUE;
   BenchUut5.weightComplete := FALSE;
   BenchUut5.weight := REAL#0.0;
   BenchUut5.firingComplete := FALSE;
   TraceIn_Mode[49] := BenchUut5.Mode;
   TraceIn_ForwardButton[49] := BenchUut5.ForwardButton;
   TraceIn_ReverseButton[49] := BenchUut5.ReverseButton;
   TraceIn_SensorFeed[49] := BenchUut5.SensorFeed;
   TraceIn_SensorWash[49] := BenchUut5.SensorWash;
   TraceIn_SensorWeight[49] := BenchUut5.SensorWeight;
   TraceIn_SensorFiring[49] := BenchUut5.SensorFiring;
   TraceIn_SensorOutput[49] := BenchUut5.SensorOutput;
   TraceIn_washComplete[49] := BenchUut5.washComplete;
   TraceIn_weightComplete[49] := BenchUut5.weightComplete;
   TraceIn_weight[49] := BenchUut5.weight;
   TraceIn_firingComplete[49] := BenchUut5.firingComplete;
   BenchUut5();
   TraceOut_MotorForward[49] := BenchUut5.MotorForward;
   TraceOut_MotorReverse[49] := BenchUut5.MotorReverse;
   TraceOut_kick[49] := BenchUut5.kick;
   TraceOut_CompletionLight[49] := BenchUut5.CompletionLight;
   TraceOut_firingTemp[49] := BenchUut5.firingTemp;
   BenchCalls := BenchCalls + 1;
 50:
   BenchUut5.Mode := TRUE;
   BenchUut5.ForwardButton := FALSE;
   BenchUut5.ReverseButton := FALSE;
   BenchUut5.SensorFeed := FALSE;
   BenchUut5.SensorWash := FALSE;
   BenchUut5.SensorWeight := TRUE;
   BenchUut5.SensorFiring := FALSE;
   BenchUut5.SensorOutput := FALSE;
   BenchUut5.washComplete := FALSE;
   BenchUut5.weightComplete := FALSE;
   BenchUut5.weight := REAL#0.0;
   BenchUut5.firingComplete := FALSE;
   TraceIn_Mode[50] := BenchUut5.Mode;
   TraceIn_ForwardButton[50] := BenchUut5.ForwardButton;
   TraceIn_ReverseButton[50] := BenchUut5.ReverseButton;
   TraceIn_SensorFeed[50] := BenchUut5.SensorFeed;
   TraceIn_SensorWash[50] := BenchUut5.SensorWash;
   TraceIn_SensorWeight[50] := BenchUut5.SensorWeight;
   TraceIn_SensorFiring[50] := BenchUut5.SensorFiring;
   TraceIn_SensorOutput[50] := BenchUut5.SensorOutput;
   TraceIn_washComplete[50] := BenchUut5.washComplete;
   TraceIn_weightComplete[50] := BenchUut5.weightComplete;
   TraceIn_weight[50] := BenchUut5.weight;
   TraceIn_firingComplete[50] := BenchUut5.firingComplete;
   BenchUut5();
   TraceOut_MotorForward[50] := BenchUut5.MotorForward;
   TraceOut_MotorReverse[50] := BenchUut5.MotorReverse;
   TraceOut_kick[50] := BenchUut5.kick;
   TraceOut_CompletionLight[50] := BenchUut5.CompletionLight;
   TraceOut_firingTemp[50] := BenchUut5.firingTemp;
   BenchCalls := BenchCalls + 1;
 51:
   BenchUut5.Mode := TRUE;
   BenchUut5.ForwardButton := FALSE;
   BenchUut5.ReverseButton := FALSE;
   BenchUut5.SensorFeed := FALSE;
   BenchUut5.SensorWash := FALSE;
   BenchUut5.SensorWeight := TRUE;
   BenchUut5.SensorFiring := FALSE;
   BenchUut5.SensorOutput := FALSE;
   BenchUut5.washComplete := FALSE;
   BenchUut5.weightComplete := TRUE;
   BenchUut5.weight := REAL#200.1;
   BenchUut5.firingComplete := FALSE;
   TraceIn_Mode[51] := BenchUut5.Mode;
   TraceIn_ForwardButton[51] := BenchUut5.ForwardButton;
   TraceIn_ReverseButton[51] := BenchUut5.ReverseButton;
   TraceIn_SensorFeed[51] := BenchUut5.SensorFeed;
   TraceIn_SensorWash[51] := BenchUut5.SensorWash;
   TraceIn_SensorWeight[51] := BenchUut5.SensorWeight;
   TraceIn_SensorFiring[51] := BenchUut5.SensorFiring;
   TraceIn_SensorOutput[51] := BenchUut5.SensorOutput;
   TraceIn_washComplete[51] := BenchUut5.washComplete;
   TraceIn_weightComplete[51] := BenchUut5.weightComplete;
   TraceIn_weight[51] := BenchUut5.weight;
   TraceIn_firingComplete[51] := BenchUut5.firingComplete;
   BenchUut5();
   TraceOut_MotorForward[51] := BenchUut5.MotorForward;
   TraceOut_MotorReverse[51] := BenchUut5.MotorReverse;
   TraceOut_kick[51] := BenchUut5.kick;
   TraceOut_CompletionLight[51] := BenchUut5.CompletionLight;
   TraceOut_firingTemp[51] := BenchUut5.firingTemp;
   BenchCalls := BenchCalls + 1;
 52:
   BenchUut5.Mode := TRUE;
   BenchUut5.ForwardButton := FALSE;
   BenchUut5.ReverseButton := FALSE;
   BenchUut5.SensorFeed := FALSE;
   BenchUut5.SensorWash := FALSE;
   BenchUut5.SensorWeight := TRUE;
   BenchUut5.SensorFiring := FALSE;
   BenchUut5.SensorOutput := FALSE;
   BenchUut5.washComplete := FALSE;
   BenchUut5.weightComplete := FALSE;
   BenchUut5.weight := REAL#0.0;
   BenchUut5.firingComplete := FALSE;
   TraceIn_Mode[52] := BenchUut5.Mode;
   TraceIn_ForwardButton[52] := BenchUut5.ForwardButton;
   TraceIn_ReverseButton[52] := BenchUut5.ReverseButton;
   TraceIn_SensorFeed[52] := BenchUut5.SensorFeed;
   TraceIn_SensorWash[52] := BenchUut5.SensorWash;
   TraceIn_SensorWeight[52] := BenchUut5.SensorWeight;
   TraceIn_SensorFiring[52] := BenchUut5.SensorFiring;
   TraceIn_SensorOutput[52] := BenchUut5.SensorOutput;
   TraceIn_washComplete[52] := BenchUut5.washComplete;
   TraceIn_weightComplete[52] := BenchUut5.weightComplete;
   TraceIn_weight[52] := BenchUut5.weight;
   TraceIn_firingComplete[52] := BenchUut5.firingComplete;
   BenchUut5();
   TraceOut_MotorForward[52] := BenchUut5.MotorForward;
   TraceOut_MotorReverse[52] := BenchUut5.MotorReverse;
   TraceOut_kick[52] := BenchUut5.kick;
   TraceOut_CompletionLight[52] := BenchUut5.CompletionLight;
   TraceOut_firingTemp[52] := BenchUut5.firingTemp;
   BenchCalls := BenchCalls + 1;
 53:
   BenchUut5.Mode := TRUE;
   BenchUut5.ForwardButton := FALSE;
   BenchUut5.ReverseButton := FALSE;
   BenchUut5.SensorFeed := FALSE;
   BenchUut5.SensorWash := FALSE;
   BenchUut5.SensorWeight := FALSE;
   BenchUut5.SensorFiring := FALSE;
   BenchUut5.SensorOutput := FALSE;
   BenchUut5.washComplete := FALSE;
   BenchUut5.weightComplete := FALSE;
   BenchUut5.weight := REAL#0.0;
   BenchUut5.firingComplete := FALSE;
   TraceIn_Mode[53] := BenchUut5.Mode;
   TraceIn_ForwardButton[53] := BenchUut5.ForwardButton;
   TraceIn_ReverseButton[53] := BenchUut5.ReverseButton;
   TraceIn_SensorFeed[53] := BenchUut5.SensorFeed;
   TraceIn_SensorWash[53] := BenchUut5.SensorWash;
   TraceIn_SensorWeight[53] := BenchUut5.SensorWeight;
   TraceIn_SensorFiring[53] := BenchUut5.SensorFiring;
   TraceIn_SensorOutput[53] := BenchUut5.SensorOutput;
   TraceIn_washComplete[53] := BenchUut5.washComplete;
   TraceIn_weightComplete[53] := BenchUut5.weightComplete;
   TraceIn_weight[53] := BenchUut5.weight;
   TraceIn_firingComplete[53] := BenchUut5.firingComplete;
   BenchUut5();
   TraceOut_MotorForward[53] := BenchUut5.MotorForward;
   TraceOut_MotorReverse[53] := BenchUut5.MotorReverse;
   TraceOut_kick[53] := BenchUut5.kick;
   TraceOut_CompletionLight[53] := BenchUut5.CompletionLight;
   TraceOut_firingTemp[53] := BenchUut5.firingTemp;
   BenchCalls := BenchCalls + 1;
 54:
   BenchUut5.Mode := TRUE;
   BenchUut5.ForwardButton := FALSE;
   BenchUut5.ReverseButton := FALSE;
   BenchUut5.SensorFeed := TRUE;
   BenchUut5.SensorWash := FALSE;
   BenchUut5.SensorWeight := FALSE;
   BenchUut5.SensorFiring := FALSE;
   BenchUut5.SensorOutput := FALSE;
   BenchUut5.washComplete := FALSE;
   BenchUut5.weightComplete := FALSE;
   BenchUut5.weight := REAL#0.0;
   BenchUut5.firingComplete := FALSE;
   TraceIn_Mode[54] := BenchUut5.Mode;
   TraceIn_ForwardButton[54] := BenchUut5.ForwardButton;
   TraceIn_ReverseButton[54] := BenchUut5.ReverseButton;
   TraceIn_SensorFeed[54] := BenchUut5.SensorFeed;
   TraceIn_SensorWash[54] := BenchUut5.SensorWash;
   TraceIn_SensorWeight[54] := BenchUut5.SensorWeight;
   TraceIn_SensorFiring[54] := BenchUut5.SensorFiring;
   TraceIn_SensorOutput[54] := BenchUut5.SensorOutput;
   TraceIn_washComplete[54] := BenchUut5.washComplete;
   TraceIn_weightComplete[54] := BenchUut5.weightComplete;
   TraceIn_weight[54] := BenchUut5.weight;
   TraceIn_firingComplete[54] := BenchUut5.firingComplete;
   BenchUut5();
   TraceOut_MotorForward[54] := BenchUut5.MotorForward;
   TraceOut_MotorReverse[54] := BenchUut5.MotorReverse;
   TraceOut_kick[54] := BenchUut5.kick;
   TraceOut_CompletionLight[54] := BenchUut5.CompletionLight;
   TraceOut_firingTemp[54] := BenchUut5.firingTemp;
   BenchCalls := BenchCalls + 1;
 55:
   BenchUut6.Mode := TRUE;
   BenchUut6.ForwardButton := FALSE;
   BenchUut6.ReverseButton := FALSE;
   BenchUut6.SensorFeed := FALSE;
   BenchUut6.SensorWash := FALSE;
   BenchUut6.SensorWeight := FALSE;
   BenchUut6.SensorFiring := FALSE;
   BenchUut6.SensorOutput := FALSE;
   BenchUut6.washComplete := TRUE;
   BenchUut6.weightComplete := TRUE;
   BenchUut6.weight := REAL#0.0;
   BenchUut6.firingComplete := TRUE;
   TraceIn_Mode[55] := BenchUut6.Mode;
   TraceIn_ForwardButton[55] := BenchUut6.ForwardButton;
   TraceIn_ReverseButton[55] := BenchUut6.ReverseButton;
   TraceIn_SensorFeed[55] := BenchUut6.SensorFeed;
   TraceIn_SensorWash[55] := BenchUut6.SensorWash;
   TraceIn_SensorWeight[55] := BenchUut6.SensorWeight;
   TraceIn_SensorFiring[55] := BenchUut6.SensorFiring;
   TraceIn_SensorOutput[55] := BenchUut6.SensorOutput;
   TraceIn_washComplete[55] := BenchUut6.washComplete;
   TraceIn_weightComplete[55] := BenchUut6.weightComplete;
   TraceIn_weight[55] := BenchUut6.weight;
   TraceIn_firingComplete[55] := BenchUut6.firingComplete;
   BenchUut6();
   TraceOut_MotorForward[55] := BenchUut6.MotorForward;
   TraceOut_MotorReverse[55] := BenchUut6.MotorReverse;
   TraceOut_kick[55] := BenchUut6.kick;
   TraceOut_CompletionLight[55] := BenchUut6.CompletionLight;
   TraceOut_firingTemp[55] := BenchUut6.firingTemp;
   BenchCalls := BenchCalls + 1;
 56:
   BenchUut6.Mode := TRUE;
   BenchUut6.ForwardButton := FALSE;
   BenchUut6.ReverseButton := FALSE;
   BenchUut6.SensorFeed := TRUE;
   BenchUut6.SensorWash := FALSE;
   BenchUut6.SensorWeight := FALSE;
   BenchUut6.SensorFiring := FALSE;
   BenchUut6.SensorOutput := FALSE;
   BenchUut6.washComplete := FALSE;
   BenchUut6.weightComplete := TRUE;
   BenchUut6.weight := REAL#0.0;
   BenchUut6.firingComplete := FALSE;
   TraceIn_Mode[56] := BenchUut6.Mode;
   TraceIn_ForwardButton[56] := BenchUut6.ForwardButton;
   TraceIn_ReverseButton[56] := BenchUut6.ReverseButton;
   TraceIn_SensorFeed[56] := BenchUut6.SensorFeed;
   TraceIn_SensorWash[56] := BenchUut6.SensorWash;
   TraceIn_SensorWeight[56] := BenchUut6.SensorWeight;
   TraceIn_SensorFiring[56] := BenchUut6.SensorFiring;
   TraceIn_SensorOutput[56] := BenchUut6.SensorOutput;
   TraceIn_washComplete[56] := BenchUut6.washComplete;
   TraceIn_weightComplete[56] := BenchUut6.weightComplete;
   TraceIn_weight[56] := BenchUut6.weight;
   TraceIn_firingComplete[56] := BenchUut6.firingComplete;
   BenchUut6();
   TraceOut_MotorForward[56] := BenchUut6.MotorForward;
   TraceOut_MotorReverse[56] := BenchUut6.MotorReverse;
   TraceOut_kick[56] := BenchUut6.kick;
   TraceOut_CompletionLight[56] := BenchUut6.CompletionLight;
   TraceOut_firingTemp[56] := BenchUut6.firingTemp;
   BenchCalls := BenchCalls + 1;
 57:
   BenchUut6.Mode := TRUE;
   BenchUut6.ForwardButton := FALSE;
   BenchUut6.ReverseButton := FALSE;
   BenchUut6.SensorFeed := FALSE;
   BenchUut6.SensorWash := TRUE;
   BenchUut6.SensorWeight := FALSE;
   BenchUut6.SensorFiring := FALSE;
   BenchUut6.SensorOutput := FALSE;
   BenchUut6.washComplete := TRUE;
   BenchUut6.weightComplete := FALSE;
   BenchUut6.weight := REAL#0.0;
   BenchUut6.firingComplete := FALSE;
   TraceIn_Mode[57] := BenchUut6.Mode;
   TraceIn_ForwardButton[57] := BenchUut6.ForwardButton;
   TraceIn_ReverseButton[57] := BenchUut6.ReverseButton;
   TraceIn_SensorFeed[57] := BenchUut6.SensorFeed;
   TraceIn_SensorWash[57] := BenchUut6.SensorWash;
   TraceIn_SensorWeight[57] := BenchUut6.SensorWeight;
   TraceIn_SensorFiring[57] := BenchUut6.SensorFiring;
   TraceIn_SensorOutput[57] := BenchUut6.SensorOutput;
   TraceIn_washComplete[57] := BenchUut6.washComplete;
   TraceIn_weightComplete[57] := BenchUut6.weightComplete;
   TraceIn_weight[57] := BenchUut6.weight;
   TraceIn_firingComplete[57] := BenchUut6.firingComplete;
   BenchUut6();
   TraceOut_MotorForward[57] := BenchUut6.MotorForward;
   TraceOut_MotorReverse[57] := BenchUut6.MotorReverse;
   TraceOut_kick[57] := BenchUut6.kick;
   TraceOut_CompletionLight[57] := BenchUut6.CompletionLight;
   TraceOut_firingTemp[57] := BenchUut6.firingTemp;
   BenchCalls := BenchCalls + 1;
 58:
   BenchUut6.Mode := TRUE;
   BenchUut6.ForwardButton := FALSE;
   BenchUut6.ReverseButton := FALSE;
   BenchUut6.SensorFeed := FALSE;
   BenchUut6.SensorWash := TRUE;
   BenchUut6.SensorWeight := FALSE;
   BenchUut6.SensorFiring := FALSE;
   BenchUut6.SensorOutput := FALSE;
   BenchUut6.washComplete := TRUE;
   BenchUut6.weightComplete := FALSE;
   BenchUut6.weight := REAL#0.0;
   BenchUut6.firingComplete := FALSE;
   TraceIn_Mode[58] := BenchUut6.Mode;
   TraceIn_ForwardButton[58] := BenchUut6.ForwardButton;
   TraceIn_ReverseButton[58] := BenchUut6.ReverseButton;
   TraceIn_SensorFeed[58] := BenchUut6.SensorFeed;
   TraceIn_SensorWash[58] := BenchUut6.SensorWash;
   TraceIn_SensorWeight[58] := BenchUut6.SensorWeight;
   TraceIn_SensorFiring[58] := BenchUut6.SensorFiring;
   TraceIn_SensorOutput[58] := BenchUut6.SensorOutput;
   TraceIn_washComplete[58] := BenchUut6.washComplete;
   TraceIn_weightComplete[58] := BenchUut6.weightComplete;
   TraceIn_weight[58] := BenchUut6.weight;
   TraceIn_firingComplete[58] := BenchUut6.firingComplete;
   BenchUut6();
   TraceOut_MotorForward[58] := BenchUut6.MotorForward;
   TraceOut_MotorReverse[58] := BenchUut6.MotorReverse;
   TraceOut_kick[58] := BenchUut6.kick;
   TraceOut_CompletionLight[58] := BenchUut6.CompletionLight;
   TraceOut_firingTemp[58] := BenchUut6.firingTemp;
   BenchCalls := BenchCalls + 1;
 59:
   BenchUut7.Mode := TRUE;
   BenchUut7.ForwardButton := FALSE;
   BenchUut7.ReverseButton := FALSE;
   BenchUut7.SensorFeed := TRUE;
   BenchUut7.SensorWash := FALSE;
   BenchUut7.SensorWeight := FALSE;
   BenchUut7.SensorFiring := FALSE;
   BenchUut7.SensorOutput := FALSE;
   BenchUut7.washComplete := FALSE;
   BenchUut7.weightComplete := FALSE;
   BenchUut7.weight := REAL#0.0;
   BenchUut7.firingComplete := FALSE;
   TraceIn_Mode[59] := BenchUut7.Mode;
   TraceIn_ForwardButton[59] := BenchUut7.ForwardButton;
   TraceIn_ReverseButton[59] := BenchUut7.ReverseButton;
   TraceIn_SensorFeed[59] := BenchUut7.SensorFeed;
   TraceIn_SensorWash[59] := BenchUut7.SensorWash;
   TraceIn_SensorWeight[59] := BenchUut7.SensorWeight;
   TraceIn_SensorFiring[59] := BenchUut7.SensorFiring;
   TraceIn_SensorOutput[59] := BenchUut7.SensorOutput;
   TraceIn_washComplete[59] := BenchUut7.washComplete;
   TraceIn_weightComplete[59] := BenchUut7.weightComplete;
   TraceIn_weight[59] := BenchUut7.weight;
   TraceIn_firingComplete[59] := BenchUut7.firingComplete;
   BenchUut7();
   TraceOut_MotorForward[59] := BenchUut7.MotorForward;
   TraceOut_MotorReverse[59] := BenchUut7.MotorReverse;
   TraceOut_kick[59] := BenchUut7.kick;
   TraceOut_CompletionLight[59] := BenchUut7.CompletionLight;
   TraceOut_firingTemp[59] := BenchUut7.firingTemp;
   BenchCalls := BenchCalls + 1;
 60:
   BenchUut7.Mode := TRUE;
   BenchUut7.ForwardButton := FALSE;
   BenchUut7.ReverseButton := FALSE;
   BenchUut7.SensorFeed := FALSE;
   BenchUut7.SensorWash := TRUE;
   BenchUut7.SensorWeight := FALSE;
   BenchUut7.SensorFiring := FALSE;
   BenchUut7.SensorOutput := FALSE;
   BenchUut7.washComplete := TRUE;
   BenchUut7.weightComplete := FALSE;
   BenchUut7.weight := REAL#0.0;
   BenchUut7.firingComplete := FALSE;
   TraceIn_Mode[60] := BenchUut7.Mode;
   TraceIn_ForwardButton[60] := BenchUut7.ForwardButton;
   TraceIn_ReverseButton[60] := BenchUut7.ReverseButton;
   TraceIn_SensorFeed[60] := BenchUut7.SensorFeed;
   TraceIn_SensorWash[60] := BenchUut7.SensorWash;
   TraceIn_SensorWeight[60] := BenchUut7.SensorWeight;
   TraceIn_SensorFiring[60] := BenchUut7.SensorFiring;
   TraceIn_SensorOutput[60] := BenchUut7.SensorOutput;
   TraceIn_washComplete[60] := BenchUut7.washComplete;
   TraceIn_weightComplete[60] := BenchUut7.weightComplete;
   TraceIn_weight[60] := BenchUut7.weight;
   TraceIn_firingComplete[60] := BenchUut7.firingComplete;
   BenchUut7();
   TraceOut_MotorForward[60] := BenchUut7.MotorForward;
   TraceOut_MotorReverse[60] := BenchUut7.MotorReverse;
   TraceOut_kick[60] := BenchUut7.kick;
   TraceOut_CompletionLight[60] := BenchUut7.CompletionLight;
   TraceOut_firingTemp[60] := BenchUut7.firingTemp;
   BenchCalls := BenchCalls + 1;
 61:
   BenchUut7.Mode := TRUE;
   BenchUut7.ForwardButton := FALSE;
   BenchUut7.ReverseButton := FALSE;
   BenchUut7.SensorFeed := FALSE;
   BenchUut7.SensorWash := TRUE;
   BenchUut7.SensorWeight := FALSE;
   BenchUut7.SensorFiring := FALSE;
   BenchUut7.SensorOutput := FALSE;
   BenchUut7.washComplete := TRUE;
   BenchUut7.weightComplete := FALSE;
   BenchUut7.weight := REAL#0.0;
   BenchUut7.firingComplete := FALSE;
   TraceIn_Mode[61] := BenchUut7.Mode;
   TraceIn_ForwardButton[61] := BenchUut7.ForwardButton;
   TraceIn_ReverseButton[61] := BenchUut7.ReverseButton;
   TraceIn_SensorFeed[61] := BenchUut7.SensorFeed;
   TraceIn_SensorWash[61] := BenchUut7.SensorWash;
   TraceIn_SensorWeight[61] := BenchUut7.SensorWeight;
   TraceIn_SensorFiring[61] := BenchUut7.SensorFiring;
   TraceIn_SensorOutput[61] := BenchUut7.SensorOutput;
   TraceIn_washComplete[61] := BenchUut7.washComplete;
   TraceIn_weightComplete[61] := BenchUut7.weightComplete;
   TraceIn_weight[61] := BenchUut7.weight;
   TraceIn_firingComplete[61] := BenchUut7.firingComplete;
   BenchUut7();
   TraceOut_MotorForward[61] := BenchUut7.MotorForward;
   TraceOut_MotorReverse[61] := BenchUut7.MotorReverse;
   TraceOut_kick[61] := BenchUut7.kick;
   TraceOut_CompletionLight[61] := BenchUut7.CompletionLight;
   TraceOut_firingTemp[61] := BenchUut7.firingTemp;
   BenchCalls := BenchCalls + 1;
 62:
   BenchUut7.Mode := TRUE;
   BenchUut7.ForwardButton := FALSE;
   BenchUut7.ReverseButton := FALSE;
   BenchUut7.SensorFeed := FALSE;
   BenchUut7.SensorWash := FALSE;
   BenchUut7.SensorWeight := TRUE;
   BenchUut7.SensorFiring := FALSE;
   BenchUut7.SensorOutput := FALSE;
   BenchUut7.washComplete := FALSE;
   BenchUut7.weightComplete := FALSE;
   BenchUut7.weight := REAL#0.0;
   BenchUut7.firingComplete := FALSE;
   TraceIn_Mode[62] := BenchUut7.Mode;
   TraceIn_ForwardButton[62] := BenchUut7.ForwardButton;
   TraceIn_ReverseButton[62] := BenchUut7.ReverseButton;
   TraceIn_SensorFeed[62] := BenchUut7.SensorFeed;
   TraceIn_SensorWash[62] := BenchUut7.SensorWash;
   TraceIn_SensorWeight[62] := BenchUut7.SensorWeight;
   TraceIn_SensorFiring[62] := BenchUut7.SensorFiring;
   TraceIn_SensorOutput[62] := BenchUut7.SensorOutput;
   TraceIn_washComplete[62] := BenchUut7.washComplete;
   TraceIn_weightComplete[62] := BenchUut7.weightComplete;
   TraceIn_weight[62] := BenchUut7.weight;
   TraceIn_firingComplete[62] := BenchUut7.firingComplete;
   BenchUut7();
   TraceOut_MotorForward[62] := BenchUut7.MotorForward;
   TraceOut_MotorReverse[62] := BenchUut7.MotorReverse;
   TraceOut_kick[62] := BenchUut7.kick;
   TraceOut_CompletionLight[62] := BenchUut7.CompletionLight;
   TraceOut_firingTemp[62] := BenchUut7.firingTemp;
   BenchCalls := BenchCalls + 1;
 63:
   BenchUut7.Mode := TRUE;
   BenchUut7.ForwardButton := FALSE;
   BenchUut7.ReverseButton := FALSE;
   BenchUut7.SensorFeed := FALSE;
   BenchUut7.SensorWash := FALSE;
   BenchUut7.SensorWeight := TRUE;
   BenchUut7.SensorFiring := FALSE;
   BenchUut7.SensorOutput := FALSE;
   BenchUut7.washComplete := FALSE;
   BenchUut7.weightComplete := TRUE;
   BenchUut7.weight := REAL#150.0;
   BenchUut7.firingComplete := FALSE;
   TraceIn_Mode[63] := BenchUut7.Mode;
   TraceIn_ForwardButton[63] := BenchUut7.ForwardButton;
   TraceIn_ReverseButton[63] := BenchUut7.ReverseButton;
   TraceIn_SensorFeed[63] := BenchUut7.SensorFeed;
   TraceIn_SensorWash[63] := BenchUut7.SensorWash;
   TraceIn_SensorWeight[63] := BenchUut7.SensorWeight;
   TraceIn_SensorFiring[63] := BenchUut7.SensorFiring;
   TraceIn_SensorOutput[63] := BenchUut7.SensorOutput;
   TraceIn_washComplete[63] := BenchUut7.washComplete;
   TraceIn_weightComplete[63] := BenchUut7.weightComplete;
   TraceIn_weight[63] := BenchUut7.weight;
   TraceIn_firingComplete[63] := BenchUut7.firingComplete;
   BenchUut7();
   TraceOut_MotorForward[63] := BenchUut7.MotorForward;
   TraceOut_MotorReverse[63] := BenchUut7.MotorReverse;
   TraceOut_kick[63] := BenchUut7.kick;
   TraceOut_CompletionLight[63] := BenchUut7.CompletionLight;
   TraceOut_firingTemp[63] := BenchUut7.firingTemp;
   BenchCalls := BenchCalls + 1;
 64:
   BenchUut7.Mode := TRUE;
   BenchUut7.ForwardButton := FALSE;
   BenchUut7.ReverseButton := FALSE;
   BenchUut7.SensorFeed := FALSE;
   BenchUut7.SensorWash := FALSE;
   BenchUut7.SensorWeight := FALSE;
   BenchUut7.SensorFiring := TRUE;
   BenchUut7.SensorOutput := FALSE;
   BenchUut7.washComplete := FALSE;
   BenchUut7.weightComplete := FALSE;
   BenchUut7.weight := REAL#0.0;
   BenchUut7.firingComplete := FALSE;
   TraceIn_Mode[64] := BenchUut7.Mode;
   TraceIn_ForwardButton[64] := BenchUut7.ForwardButton;
   TraceIn_ReverseButton[64] := BenchUut7.ReverseButton;
   TraceIn_SensorFeed[64] := BenchUut7.SensorFeed;
   TraceIn_SensorWash[64] := BenchUut7.SensorWash;
   TraceIn_SensorWeight[64] := BenchUut7.SensorWeight;
   TraceIn_SensorFiring[64] := BenchUut7.SensorFiring;
   TraceIn_SensorOutput[64] := BenchUut7.SensorOutput;
   TraceIn_washComplete[64] := BenchUut7.washComplete;
   TraceIn_weightComplete[64] := BenchUut7.weightComplete;
   TraceIn_weight[64] := BenchUut7.weight;
   TraceIn_firingComplete[64] := BenchUut7.firingComplete;
   BenchUut7();
   TraceOut_MotorForward[64] := BenchUut7.MotorForward;
   TraceOut_MotorReverse[64] := BenchUut7.MotorReverse;
   TraceOut_kick[64] := BenchUut7.kick;
   TraceOut_CompletionLight[64] := BenchUut7.CompletionLight;
   TraceOut_firingTemp[64] := BenchUut7.firingTemp;
   BenchCalls := BenchCalls + 1;
 65:
   BenchUut7.Mode := TRUE;
   BenchUut7.ForwardButton := FALSE;
   BenchUut7.ReverseButton := FALSE;
   BenchUut7.SensorFeed := FALSE;
   BenchUut7.SensorWash := FALSE;
   BenchUut7.SensorWeight := FALSE;
   BenchUut7.SensorFiring := TRUE;
   BenchUut7.SensorOutput := FALSE;
   BenchUut7.washComplete := FALSE;
   BenchUut7.weightComplete := FALSE;
   BenchUut7.weight := REAL#0.0;
   BenchUut7.firingComplete := TRUE;
   TraceIn_Mode[65] := BenchUut7.Mode;
   TraceIn_ForwardButton[65] := BenchUut7.ForwardButton;
   TraceIn_ReverseButton[65] := BenchUut7.ReverseButton;
   TraceIn_SensorFeed[65] := BenchUut7.SensorFeed;
   TraceIn_SensorWash[65] := BenchUut7.SensorWash;
   TraceIn_SensorWeight[65] := BenchUut7.SensorWeight;
   TraceIn_SensorFiring[65] := BenchUut7.SensorFiring;
   TraceIn_SensorOutput[65] := BenchUut7.SensorOutput;
   TraceIn_washComplete[65] := BenchUut7.washComplete;
   TraceIn_weightComplete[65] := BenchUut7.weightComplete;
   TraceIn_weight[65] := BenchUut7.weight;
   TraceIn_firingComplete[65] := BenchUut7.firingComplete;
   BenchUut7();
   TraceOut_MotorForward[65] := BenchUut7.MotorForward;
   TraceOut_MotorReverse[65] := BenchUut7.MotorReverse;
   TraceOut_kick[65] := BenchUut7.kick;
   TraceOut_CompletionLight[65] := BenchUut7.CompletionLight;
   TraceOut_firingTemp[65] := BenchUut7.firingTemp;
   BenchCalls := BenchCalls + 1;
 66:
   BenchUut7.Mode := TRUE;
   BenchUut7.ForwardButton := FALSE;
   BenchUut7.ReverseButton := FALSE;
   BenchUut7.SensorFeed := FALSE;
   BenchUut7.SensorWash := FALSE;
   BenchUut7.SensorWeight := FALSE;
   BenchUut7.SensorFiring := FALSE;
   BenchUut7.SensorOutput := TRUE;
   BenchUut7.washComplete := FALSE;
   BenchUut7.weightComplete := FALSE;
   BenchUut7.weight := REAL#0.0;
   BenchUut7.firingComplete := FALSE;
   TraceIn_Mode[66] := BenchUut7.Mode;
   TraceIn_ForwardButton[66] := BenchUut7.ForwardButton;
   TraceIn_ReverseButton[66] := BenchUut7.ReverseButton;
   TraceIn_SensorFeed[66] := BenchUut7.SensorFeed;
   TraceIn_SensorWash[66] := BenchUut7.SensorWash;
   TraceIn_SensorWeight[66] := BenchUut7.SensorWeight;
   TraceIn_SensorFiring[66] := BenchUut7.SensorFiring;
   TraceIn_SensorOutput[66] := BenchUut7.SensorOutput;
   TraceIn_washComplete[66] := BenchUut7.washComplete;
   TraceIn_weightComplete[66] := BenchUut7.weightComplete;
   TraceIn_weight[66] := BenchUut7.weight;
   TraceIn_firingComplete[66] := BenchUut7.firingComplete;
   BenchUut7();
   TraceOut_MotorForward[66] := BenchUut7.MotorForward;
   TraceOut_MotorReverse[66] := BenchUut7.MotorReverse;
   TraceOut_kick[66] := BenchUut7.kick;
   TraceOut_CompletionLight[66] := BenchUut7.CompletionLight;
   TraceOut_firingTemp[66] := BenchUut7.firingTemp;
   BenchCalls := BenchCalls + 1;
 67:
   BenchUut7.Mode := TRUE;
   BenchUut7.ForwardButton := FALSE;
   BenchUut7.ReverseButton := FALSE;
   BenchUut7.SensorFeed := FALSE;
   BenchUut7.SensorWash := FALSE;
   BenchUut7.SensorWeight := FALSE;
   BenchUut7.SensorFiring := FALSE;
   BenchUut7.SensorOutput := FALSE;
   BenchUut7.washComplete := FALSE;
   BenchUut7.weightComplete := FALSE;
   BenchUut7.weight := REAL#0.0;
   BenchUut7.firingComplete := FALSE;
   TraceIn_Mode[67] := BenchUut7.Mode;
   TraceIn_ForwardButton[67] := BenchUut7.ForwardButton;
   TraceIn_ReverseButton[67] := BenchUut7.ReverseButton;
   TraceIn_SensorFeed[67] := BenchUut7.SensorFeed;
   TraceIn_SensorWash[67] := BenchUut7.SensorWash;
   TraceIn_SensorWeight[67] := BenchUut7.SensorWeight;
   TraceIn_SensorFiring[67] := BenchUut7.SensorFiring;
   TraceIn_SensorOutput[67] := BenchUut7.SensorOutput;
   TraceIn_washComplete[67] := BenchUut7.washComplete;
   TraceIn_weightComplete[67] := BenchUut7.weightComplete;
   TraceIn_weight[67] := BenchUut7.weight;
   TraceIn_firingComplete[67] := BenchUut7.firingComplete;
   BenchUut7();
   TraceOut_MotorForward[67] := BenchUut7.MotorForward;
   TraceOut_MotorReverse[67] := BenchUut7.MotorReverse;
   TraceOut_kick[67] := BenchUut7.kick;
   TraceOut_CompletionLight[67] := BenchUut7.CompletionLight;
   TraceOut_firingTemp[67] := BenchUut7.firingTemp;
   BenchCalls := BenchCalls + 1;
 68:
   BenchUut7.Mode := TRUE;
   BenchUut7.ForwardButton := FALSE;
   BenchUut7.ReverseButton := FALSE;
   BenchUut7.SensorFeed := TRUE;
   BenchUut7.SensorWash := FALSE;
   BenchUut7.SensorWeight := FALSE;
   BenchUut7.SensorFiring := FALSE;
   BenchUut7.SensorOutput := FALSE;
   BenchUut7.washComplete := FALSE;
   BenchUut7.weightComplete := FALSE;
   BenchUut7.weight := REAL#0.0;
   BenchUut7.firingComplete := FALSE;
   TraceIn_Mode[68] := BenchUut7.Mode;
   TraceIn_ForwardButton[68] := BenchUut7.ForwardButton;
   TraceIn_ReverseButton[68] := BenchUut7.ReverseButton;
   TraceIn_SensorFeed[68] := BenchUut7.SensorFeed;
   TraceIn_SensorWash[68] := BenchUut7.SensorWash;
   TraceIn_SensorWeight[68] := BenchUut7.SensorWeight;
   TraceIn_SensorFiring[68] := BenchUut7.SensorFiring;
   TraceIn_SensorOutput[68] := BenchUut7.SensorOutput;
   TraceIn_washComplete[68] := BenchUut7.washComplete;
   TraceIn_weightComplete[68] := BenchUut7.weightComplete;
   TraceIn_weight[68] := BenchUut7.weight;
   TraceIn_firingComplete[68] := BenchUut7.firingComplete;
   BenchUut7();
   TraceOut_MotorForward[68] := BenchUut7.MotorForward;
   TraceOut_MotorReverse[68] := BenchUut7.MotorReverse;
   TraceOut_kick[68] := BenchUut7.kick;
   TraceOut_CompletionLight[68] := BenchUut7.CompletionLight;
   TraceOut_firingTemp[68] := BenchUut7.firingTemp;
   BenchCalls := BenchCalls + 1;
 69:
   BenchUut7.Mode := TRUE;
   BenchUut7.ForwardButton := FALSE;
   BenchUut7.ReverseButton := FALSE;
   BenchUut7.SensorFeed := FALSE;
   BenchUut7.SensorWash := TRUE;
   BenchUut7.SensorWeight := FALSE;
   BenchUut7.SensorFiring := FALSE;
   BenchUut7.SensorOutput := FALSE;
   BenchUut7.washComplete := FALSE;
   BenchUut7.weightComplete := FALSE;
   BenchUut7.weight := REAL#0.0;
   BenchUut7.firingComplete := FALSE;
   TraceIn_Mode[69] := BenchUut7.Mode;
   TraceIn_ForwardButton[69] := BenchUut7.ForwardButton;
   TraceIn_ReverseButton[69] := BenchUut7.ReverseButton;
   TraceIn_SensorFeed[69] := BenchUut7.SensorFeed;
   TraceIn_SensorWash[69] := BenchUut7.SensorWash;
   TraceIn_SensorWeight[69] := BenchUut7.SensorWeight;
   TraceIn_SensorFiring[69] := BenchUut7.SensorFiring;
   TraceIn_SensorOutput[69] := BenchUut7.SensorOutput;
   TraceIn_washComplete[69] := BenchUut7.washComplete;
   TraceIn_weightComplete[69] := BenchUut7.weightComplete;
   TraceIn_weight[69] := BenchUut7.weight;
   TraceIn_firingComplete[69] := BenchUut7.firingComplete;
   BenchUut7();
   TraceOut_MotorForward[69] := BenchUut7.MotorForward;
   TraceOut_MotorReverse[69] := BenchUut7.MotorReverse;
   TraceOut_kick[69] := BenchUut7.kick;
   TraceOut_CompletionLight[69] := BenchUut7.CompletionLight;
   TraceOut_firingTemp[69] := BenchUut7.firingTemp;
   BenchCalls := BenchCalls + 1;
 70:
   BenchUut7.Mode := TRUE;
   BenchUut7.ForwardButton := FALSE;
   BenchUut7.ReverseButton := FALSE;
   BenchUut7.SensorFeed := FALSE;
   BenchUut7.SensorWash := TRUE;
   BenchUut7.SensorWeight := FALSE;
   BenchUut7.SensorFiring := FALSE;
   BenchUut7.SensorOutput := FALSE;
   BenchUut7.washComplete := TRUE;
   BenchUut7.weightComplete := FALSE;
   BenchUut7.weight := REAL#0.0;
   BenchUut7.firingComplete := FALSE;
   TraceIn_Mode[70] := BenchUut7.Mode;
   TraceIn_ForwardButton[70] := BenchUut7.ForwardButton;
   TraceIn_ReverseButton[70] := BenchUut7.ReverseButton;
   TraceIn_SensorFeed[70] := BenchUut7.SensorFeed;
   TraceIn_SensorWash[70] := BenchUut7.SensorWash;
   TraceIn_SensorWeight[70] := BenchUut7.SensorWeight;
   TraceIn_SensorFiring[70] := BenchUut7.SensorFiring;
   TraceIn_SensorOutput[70] := BenchUut7.SensorOutput;
   TraceIn_washComplete[70] := BenchUut7.washComplete;
   TraceIn_weightComplete[70] := BenchUut7.weightComplete;
   TraceIn_weight[70] := BenchUut7.weight;
   TraceIn_firingComplete[70] := BenchUut7.firingComplete;
   BenchUut7();
   TraceOut_MotorForward[70] := BenchUut7.MotorForward;
   TraceOut_MotorReverse[70] := BenchUut7.MotorReverse;
   TraceOut_kick[70] := BenchUut7.kick;
   TraceOut_CompletionLight[70] := BenchUut7.CompletionLight;
   TraceOut_firingTemp[70] := BenchUut7.firingTemp;
   BenchCalls := BenchCalls + 1;
 71:
   BenchUut7.Mode := TRUE;
   BenchUut7.ForwardButton := FALSE;
   BenchUut7.ReverseButton := FALSE;
   BenchUut7.SensorFeed := FALSE;
   BenchUut7.SensorWash := FALSE;
   BenchUut7.SensorWeight := TRUE;
   BenchUut7.SensorFiring := FALSE;
   BenchUut7.SensorOutput := FALSE;
   BenchUut7.washComplete := FALSE;
   BenchUut7.weightComplete := FALSE;
   BenchUut7.weight := REAL#0.0;
   BenchUut7.firingComplete := FALSE;
   TraceIn_Mode[71] := BenchUut7.Mode;
   TraceIn_ForwardButton[71] := BenchUut7.ForwardButton;
   TraceIn_ReverseButton[71] := BenchUut7.ReverseButton;
   TraceIn_SensorFeed[71] := BenchUut7.SensorFeed;
   TraceIn_SensorWash[71] := BenchUut7.SensorWash;
   TraceIn_SensorWeight[71] := BenchUut7.SensorWeight;
   TraceIn_SensorFiring[71] := BenchUut7.SensorFiring;
   TraceIn_SensorOutput[71] := BenchUut7.SensorOutput;
   TraceIn_washComplete[71] := BenchUut7.washComplete;
   TraceIn_weightComplete[71] := BenchUut7.weightComplete;
   TraceIn_weight[71] := BenchUut7.weight;
   TraceIn_firingComplete[71] := BenchUut7.firingComplete;
   BenchUut7();
   TraceOut_MotorForward[71] := BenchUut7.MotorForward;
   TraceOut_MotorReverse[71] := BenchUut7.MotorReverse;
   TraceOut_kick[71] := BenchUut7.kick;
   TraceOut_CompletionLight[71] := BenchUut7.CompletionLight;
   TraceOut_firingTemp[71] := BenchUut7.firingTemp;
   BenchCalls := BenchCalls + 1;
 72:
   BenchUut7.Mode := TRUE;
   BenchUut7.ForwardButton := FALSE;
   BenchUut7.ReverseButton := FALSE;
   BenchUut7.SensorFeed := FALSE;
   BenchUut7.SensorWash := FALSE;
   BenchUut7.SensorWeight := TRUE;
   BenchUut7.SensorFiring := FALSE;
   BenchUut7.SensorOutput := FALSE;
   BenchUut7.washComplete := FALSE;
   BenchUut7.weightComplete := TRUE;
   BenchUut7.weight := REAL#99.9;
   BenchUut7.firingComplete := FALSE;
   TraceIn_Mode[72] := BenchUut7.Mode;
   TraceIn_ForwardButton[72] := BenchUut7.ForwardButton;
   TraceIn_ReverseButton[72] := BenchUut7.ReverseButton;
   TraceIn_SensorFeed[72] := BenchUut7.SensorFeed;
   TraceIn_SensorWash[72] := BenchUut7.SensorWash;
   TraceIn_SensorWeight[72] := BenchUut7.SensorWeight;
   TraceIn_SensorFiring[72] := BenchUut7.SensorFiring;
   TraceIn_SensorOutput[72] := BenchUut7.SensorOutput;
   TraceIn_washComplete[72] := BenchUut7.washComplete;
   TraceIn_weightComplete[72] := BenchUut7.weightComplete;
   TraceIn_weight[72] := BenchUut7.weight;
   TraceIn_firingComplete[72] := BenchUut7.firingComplete;
   BenchUut7();
   TraceOut_MotorForward[72] := BenchUut7.MotorForward;
   TraceOut_MotorReverse[72] := BenchUut7.MotorReverse;
   TraceOut_kick[72] := BenchUut7.kick;
   TraceOut_CompletionLight[72] := BenchUut7.CompletionLight;
   TraceOut_firingTemp[72] := BenchUut7.firingTemp;
   BenchCalls := BenchCalls + 1;
 73:
   BenchUut7.Mode := TRUE;
   BenchUut7.ForwardButton := FALSE;
   BenchUut7.ReverseButton := FALSE;
   BenchUut7.SensorFeed := FALSE;
   BenchUut7.SensorWash := FALSE;
   BenchUut7.SensorWeight := TRUE;
   BenchUut7.SensorFiring := FALSE;
   BenchUut7.SensorOutput := FALSE;
   BenchUut7.washComplete := FALSE;
   BenchUut7.weightComplete := FALSE;
   BenchUut7.weight := REAL#0.0;
   BenchUut7.firingComplete := FALSE;
   TraceIn_Mode[73] := BenchUut7.Mode;
   TraceIn_ForwardButton[73] := BenchUut7.ForwardButton;
   TraceIn_ReverseButton[73] := BenchUut7.ReverseButton;
   TraceIn_SensorFeed[73] := BenchUut7.SensorFeed;
   TraceIn_SensorWash[73] := BenchUut7.SensorWash;
   TraceIn_SensorWeight[73] := BenchUut7.SensorWeight;
   TraceIn_SensorFiring[73] := BenchUut7.SensorFiring;
   TraceIn_SensorOutput[73] := BenchUut7.SensorOutput;
   TraceIn_washComplete[73] := BenchUut7.washComplete;
   TraceIn_weightComplete[73] := BenchUut7.weightComplete;
   TraceIn_weight[73] := BenchUut7.weight;
   TraceIn_firingComplete[73] := BenchUut7.firingComplete;
   BenchUut7();
   TraceOut_MotorForward[73] := BenchUut7.MotorForward;
   TraceOut_MotorReverse[73] := BenchUut7.MotorReverse;
   TraceOut_kick[73] := BenchUut7.kick;
   TraceOut_CompletionLight[73] := BenchUut7.CompletionLight;
   TraceOut_firingTemp[73] := BenchUut7.firingTemp;
   BenchCalls := BenchCalls + 1;
 74:
   BenchUut7.Mode := TRUE;
   BenchUut7.ForwardButton := FALSE;
   BenchUut7.ReverseButton := FALSE;
   BenchUut7.SensorFeed := FALSE;
   BenchUut7.SensorWash := FALSE;
   BenchUut7.SensorWeight := FALSE;
   BenchUut7.SensorFiring := FALSE;
   BenchUut7.SensorOutput := FALSE;
   BenchUut7.washComplete := FALSE;
   BenchUut7.weightComplete := FALSE;
   BenchUut7.weight := REAL#0.0;
   BenchUut7.firingComplete := FALSE;
   TraceIn_Mode[74] := BenchUut7.Mode;
   TraceIn_ForwardButton[74] := BenchUut7.ForwardButton;
   TraceIn_ReverseButton[74] := BenchUut7.ReverseButton;
   TraceIn_SensorFeed[74] := BenchUut7.SensorFeed;
   TraceIn_SensorWash[74] := BenchUut7.SensorWash;
   TraceIn_SensorWeight[74] := BenchUut7.SensorWeight;
   TraceIn_SensorFiring[74] := BenchUut7.SensorFiring;
   TraceIn_SensorOutput[74] := BenchUut7.SensorOutput;
   TraceIn_washComplete[74] := BenchUut7.washComplete;
   TraceIn_weightComplete[74] := BenchUut7.weightComplete;
   TraceIn_weight[74] := BenchUut7.weight;
   TraceIn_firingComplete[74] := BenchUut7.firingComplete;
   BenchUut7();
   TraceOut_MotorForward[74] := BenchUut7.MotorForward;
   TraceOut_MotorReverse[74] := BenchUut7.MotorReverse;
   TraceOut_kick[74] := BenchUut7.kick;
   TraceOut_CompletionLight[74] := BenchUut7.CompletionLight;
   TraceOut_firingTemp[74] := BenchUut7.firingTemp;
   BenchCalls := BenchCalls + 1;
 75:
   BenchUut8.Mode := TRUE;
   BenchUut8.ForwardButton := FALSE;
   BenchUut8.ReverseButton := FALSE;
   BenchUut8.SensorFeed := TRUE;
   BenchUut8.SensorWash := FALSE;
   BenchUut8.SensorWeight := FALSE;
   BenchUut8.SensorFiring := FALSE;
   BenchUut8.SensorOutput := FALSE;
   BenchUut8.washComplete := FALSE;
   BenchUut8.weightComplete := FALSE;
   BenchUut8.weight := REAL#150.0;
   BenchUut8.firingComplete := FALSE;
   TraceIn_Mode[75] := BenchUut8.Mode;
   TraceIn_ForwardButton[75] := BenchUut8.ForwardButton;
   TraceIn_ReverseButton[75] := BenchUut8.ReverseButton;
   TraceIn_SensorFeed[75] := BenchUut8.SensorFeed;
   TraceIn_SensorWash[75] := BenchUut8.SensorWash;
   TraceIn_SensorWeight[75] := BenchUut8.SensorWeight;
   TraceIn_SensorFiring[75] := BenchUut8.SensorFiring;
   TraceIn_SensorOutput[75] := BenchUut8.SensorOutput;
   TraceIn_washComplete[75] := BenchUut8.washComplete;
   TraceIn_weightComplete[75] := BenchUut8.weightComplete;
   TraceIn_weight[75] := BenchUut8.weight;
   TraceIn_firingComplete[75] := BenchUut8.firingComplete;
   BenchUut8();
   TraceOut_MotorForward[75] := BenchUut8.MotorForward;
   TraceOut_MotorReverse[75] := BenchUut8.MotorReverse;
   TraceOut_kick[75] := BenchUut8.kick;
   TraceOut_CompletionLight[75] := BenchUut8.CompletionLight;
   TraceOut_firingTemp[75] := BenchUut8.firingTemp;
   BenchCalls := BenchCalls + 1;
 76:
   BenchUut8.Mode := TRUE;
   BenchUut8.ForwardButton := FALSE;
   BenchUut8.ReverseButton := FALSE;
   BenchUut8.SensorFeed := FALSE;
   BenchUut8.SensorWash := FALSE;
   BenchUut8.SensorWeight := FALSE;
   BenchUut8.SensorFiring := FALSE;
   BenchUut8.SensorOutput := FALSE;
   BenchUut8.washComplete := FALSE;
   BenchUut8.weightComplete := FALSE;
   BenchUut8.weight := REAL#150.0;
   BenchUut8.firingComplete := FALSE;
   TraceIn_Mode[76] := BenchUut8.Mode;
   TraceIn_ForwardButton[76] := BenchUut8.ForwardButton;
   TraceIn_ReverseButton[76] := BenchUut8.ReverseButton;
   TraceIn_SensorFeed[76] := BenchUut8.SensorFeed;
   TraceIn_SensorWash[76] := BenchUut8.SensorWash;
   TraceIn_SensorWeight[76] := BenchUut8.SensorWeight;
   TraceIn_SensorFiring[76] := BenchUut8.SensorFiring;
   TraceIn_SensorOutput[76] := BenchUut8.SensorOutput;
   TraceIn_washComplete[76] := BenchUut8.washComplete;
   TraceIn_weightComplete[76] := BenchUut8.weightComplete;
   TraceIn_weight[76] := BenchUut8.weight;
   TraceIn_firingComplete[76] := BenchUut8.firingComplete;
   BenchUut8();
   TraceOut_MotorForward[76] := BenchUut8.MotorForward;
   TraceOut_MotorReverse[76] := BenchUut8.MotorReverse;
   TraceOut_kick[76] := BenchUut8.kick;
   TraceOut_CompletionLight[76] := BenchUut8.CompletionLight;
   TraceOut_firingTemp[76] := BenchUut8.firingTemp;
   BenchCalls := BenchCalls + 1;
 77:
   BenchUut8.Mode := TRUE;
   BenchUut8.ForwardButton := FALSE;
   BenchUut8.ReverseButton := FALSE;
   BenchUut8.SensorFeed := FALSE;
   BenchUut8.SensorWash := TRUE;
   BenchUut8.SensorWeight := FALSE;
   BenchUut8.SensorFiring := FALSE;
   BenchUut8.SensorOutput := FALSE;
   BenchUut8.washComplete := TRUE;
   BenchUut8.weightComplete := FALSE;
   BenchUut8.weight := REAL#150.0;
   BenchUut8.firingComplete := FALSE;
   TraceIn_Mode[77] := BenchUut8.Mode;
   TraceIn_ForwardButton[77] := BenchUut8.ForwardButton;
   TraceIn_ReverseButton[77] := BenchUut8.ReverseButton;
   TraceIn_SensorFeed[77] := BenchUut8.SensorFeed;
   TraceIn_SensorWash[77] := BenchUut8.SensorWash;
   TraceIn_SensorWeight[77] := BenchUut8.SensorWeight;
   TraceIn_SensorFiring[77] := BenchUut8.SensorFiring;
   TraceIn_SensorOutput[77] := BenchUut8.SensorOutput;
   TraceIn_washComplete[77] := BenchUut8.washComplete;
   TraceIn_weightComplete[77] := BenchUut8.weightComplete;
   TraceIn_weight[77] := BenchUut8.weight;
   TraceIn_firingComplete[77] := BenchUut8.firingComplete;
   BenchUut8();
   TraceOut_MotorForward[77] := BenchUut8.MotorForward;
   TraceOut_MotorReverse[77] := BenchUut8.MotorReverse;
   TraceOut_kick[77] := BenchUut8.kick;
   TraceOut_CompletionLight[77] := BenchUut8.CompletionLight;
   TraceOut_firingTemp[77] := BenchUut8.firingTemp;
   BenchCalls := BenchCalls + 1;
 78:
   BenchUut8.Mode := TRUE;
   BenchUut8.ForwardButton := FALSE;
   BenchUut8.ReverseButton := FALSE;
   BenchUut8.SensorFeed := FALSE;
   BenchUut8.SensorWash := TRUE;
   BenchUut8.SensorWeight := FALSE;
   BenchUut8.SensorFiring := FALSE;
   BenchUut8.SensorOutput := FALSE;
   BenchUut8.washComplete := TRUE;
   BenchUut8.weightComplete := FALSE;
   BenchUut8.weight := REAL#150.0;
   BenchUut8.firingComplete := FALSE;
   TraceIn_Mode[78] := BenchUut8.Mode;
   TraceIn_ForwardButton[78] := BenchUut8.ForwardButton;
   TraceIn_ReverseButton[78] := BenchUut8.ReverseButton;
   TraceIn_SensorFeed[78] := BenchUut8.SensorFeed;
   TraceIn_SensorWash[78] := BenchUut8.SensorWash;
   TraceIn_SensorWeight[78] := BenchUut8.SensorWeight;
   TraceIn_SensorFiring[78] := BenchUut8.SensorFiring;
   TraceIn_SensorOutput[78] := BenchUut8.SensorOutput;
   TraceIn_washComplete[78] := BenchUut8.washComplete;
   TraceIn_weightComplete[78] := BenchUut8.weightComplete;
   TraceIn_weight[78] := BenchUut8.weight;
   TraceIn_firingComplete[78] := BenchUut8.firingComplete;
   BenchUut8();
   TraceOut_MotorForward[78] := BenchUut8.MotorForward;
   TraceOut_MotorReverse[78] := BenchUut8.MotorReverse;
   TraceOut_kick[78] := BenchUut8.kick;
   TraceOut_CompletionLight[78] := BenchUut8.CompletionLight;
   TraceOut_firingTemp[78] := BenchUut8.firingTemp;
   BenchCalls := BenchCalls + 1;
 79:
   BenchUut8.Mode := TRUE;
   BenchUut8.ForwardButton := FALSE;
   BenchUut8.ReverseButton := FALSE;
   BenchUut8.SensorFeed := FALSE;
   BenchUut8.SensorWash := FALSE;
   BenchUut8.SensorWeight := FALSE;
   BenchUut8.SensorFiring := FALSE;
   BenchUut8.SensorOutput := FALSE;
   BenchUut8.washComplete := FALSE;
   BenchUut8.weightComplete := FALSE;
   BenchUut8.weight := REAL#150.0;
   BenchUut8.firingComplete := FALSE;
   TraceIn_Mode[79] := BenchUut8.Mode;
   TraceIn_ForwardButton[79] := BenchUut8.ForwardButton;
   TraceIn_ReverseButton[79] := BenchUut8.ReverseButton;
   TraceIn_SensorFeed[79] := BenchUut8.SensorFeed;
   TraceIn_SensorWash[79] := BenchUut8.SensorWash;
   TraceIn_SensorWeight[79] := BenchUut8.SensorWeight;
   TraceIn_SensorFiring[79] := BenchUut8.SensorFiring;
   TraceIn_SensorOutput[79] := BenchUut8.SensorOutput;
   TraceIn_washComplete[79] := BenchUut8.washComplete;
   TraceIn_weightComplete[79] := BenchUut8.weightComplete;
   TraceIn_weight[79] := BenchUut8.weight;
   TraceIn_firingComplete[79] := BenchUut8.firingComplete;
   BenchUut8();
   TraceOut_MotorForward[79] := BenchUut8.MotorForward;
   TraceOut_MotorReverse[79] := BenchUut8.MotorReverse;
   TraceOut_kick[79] := BenchUut8.kick;
   TraceOut_CompletionLight[79] := BenchUut8.CompletionLight;
   TraceOut_firingTemp[79] := BenchUut8.firingTemp;
   BenchCalls := BenchCalls + 1;
 80:
   BenchUut8.Mode := TRUE;
   BenchUut8.ForwardButton := FALSE;
   BenchUut8.ReverseButton := FALSE;
   BenchUut8.SensorFeed := FALSE;
   BenchUut8.SensorWash := FALSE;
   BenchUut8.SensorWeight := TRUE;
   BenchUut8.SensorFiring := FALSE;
   BenchUut8.SensorOutput := FALSE;
   BenchUut8.washComplete := FALSE;
   BenchUut8.weightComplete := FALSE;
   BenchUut8.weight := REAL#150.0;
   BenchUut8.firingComplete := FALSE;
   TraceIn_Mode[80] := BenchUut8.Mode;
   TraceIn_ForwardButton[80] := BenchUut8.ForwardButton;
   TraceIn_ReverseButton[80] := BenchUut8.ReverseButton;
   TraceIn_SensorFeed[80] := BenchUut8.SensorFeed;
   TraceIn_SensorWash[80] := BenchUut8.SensorWash;
   TraceIn_SensorWeight[80] := BenchUut8.SensorWeight;
   TraceIn_SensorFiring[80] := BenchUut8.SensorFiring;
   TraceIn_SensorOutput[80] := BenchUut8.SensorOutput;
   TraceIn_washComplete[80] := BenchUut8.washComplete;
   TraceIn_weightComplete[80] := BenchUut8.weightComplete;
   TraceIn_weight[80] := BenchUut8.weight;
   TraceIn_firingComplete[80] := BenchUut8.firingComplete;
   BenchUut8();
   TraceOut_MotorForward[80] := BenchUut8.MotorForward;
   TraceOut_MotorReverse[80] := BenchUut8.MotorReverse;
   TraceOut_kick[80] := BenchUut8.kick;
   TraceOut_CompletionLight[80] := BenchUut8.CompletionLight;
   TraceOut_firingTemp[80] := BenchUut8.firingTemp;
   BenchCalls := BenchCalls + 1;
 81:
   BenchUut8.Mode := TRUE;
   BenchUut8.ForwardButton := FALSE;
   BenchUut8.ReverseButton := FALSE;
   BenchUut8.SensorFeed := FALSE;
   BenchUut8.SensorWash := FALSE;
   BenchUut8.SensorWeight := TRUE;
   BenchUut8.SensorFiring := FALSE;
   BenchUut8.SensorOutput := FALSE;
   BenchUut8.washComplete := FALSE;
   BenchUut8.weightComplete := TRUE;
   BenchUut8.weight := REAL#100.0001;
   BenchUut8.firingComplete := FALSE;
   TraceIn_Mode[81] := BenchUut8.Mode;
   TraceIn_ForwardButton[81] := BenchUut8.ForwardButton;
   TraceIn_ReverseButton[81] := BenchUut8.ReverseButton;
   TraceIn_SensorFeed[81] := BenchUut8.SensorFeed;
   TraceIn_SensorWash[81] := BenchUut8.SensorWash;
   TraceIn_SensorWeight[81] := BenchUut8.SensorWeight;
   TraceIn_SensorFiring[81] := BenchUut8.SensorFiring;
   TraceIn_SensorOutput[81] := BenchUut8.SensorOutput;
   TraceIn_washComplete[81] := BenchUut8.washComplete;
   TraceIn_weightComplete[81] := BenchUut8.weightComplete;
   TraceIn_weight[81] := BenchUut8.weight;
   TraceIn_firingComplete[81] := BenchUut8.firingComplete;
   BenchUut8();
   TraceOut_MotorForward[81] := BenchUut8.MotorForward;
   TraceOut_MotorReverse[81] := BenchUut8.MotorReverse;
   TraceOut_kick[81] := BenchUut8.kick;
   TraceOut_CompletionLight[81] := BenchUut8.CompletionLight;
   TraceOut_firingTemp[81] := BenchUut8.firingTemp;
   BenchCalls := BenchCalls + 1;
 82:
   BenchUut8.Mode := FALSE;
   BenchUut8.ForwardButton := FALSE;
   BenchUut8.ReverseButton := TRUE;
   BenchUut8.SensorFeed := FALSE;
   BenchUut8.SensorWash := FALSE;
   BenchUut8.SensorWeight := FALSE;
   BenchUut8.SensorFiring := FALSE;
   BenchUut8.SensorOutput := FALSE;
   BenchUut8.washComplete := FALSE;
   BenchUut8.weightComplete := FALSE;
   BenchUut8.weight := REAL#150.0;
   BenchUut8.firingComplete := FALSE;
   TraceIn_Mode[82] := BenchUut8.Mode;
   TraceIn_ForwardButton[82] := BenchUut8.ForwardButton;
   TraceIn_ReverseButton[82] := BenchUut8.ReverseButton;
   TraceIn_SensorFeed[82] := BenchUut8.SensorFeed;
   TraceIn_SensorWash[82] := BenchUut8.SensorWash;
   TraceIn_SensorWeight[82] := BenchUut8.SensorWeight;
   TraceIn_SensorFiring[82] := BenchUut8.SensorFiring;
   TraceIn_SensorOutput[82] := BenchUut8.SensorOutput;
   TraceIn_washComplete[82] := BenchUut8.washComplete;
   TraceIn_weightComplete[82] := BenchUut8.weightComplete;
   TraceIn_weight[82] := BenchUut8.weight;
   TraceIn_firingComplete[82] := BenchUut8.firingComplete;
   BenchUut8();
   TraceOut_MotorForward[82] := BenchUut8.MotorForward;
   TraceOut_MotorReverse[82] := BenchUut8.MotorReverse;
   TraceOut_kick[82] := BenchUut8.kick;
   TraceOut_CompletionLight[82] := BenchUut8.CompletionLight;
   TraceOut_firingTemp[82] := BenchUut8.firingTemp;
   BenchCalls := BenchCalls + 1;
 83:
   BenchUut8.Mode := TRUE;
   BenchUut8.ForwardButton := FALSE;
   BenchUut8.ReverseButton := FALSE;
   BenchUut8.SensorFeed := TRUE;
   BenchUut8.SensorWash := FALSE;
   BenchUut8.SensorWeight := FALSE;
   BenchUut8.SensorFiring := FALSE;
   BenchUut8.SensorOutput := FALSE;
   BenchUut8.washComplete := FALSE;
   BenchUut8.weightComplete := FALSE;
   BenchUut8.weight := REAL#150.0;
   BenchUut8.firingComplete := FALSE;
   TraceIn_Mode[83] := BenchUut8.Mode;
   TraceIn_ForwardButton[83] := BenchUut8.ForwardButton;
   TraceIn_ReverseButton[83] := BenchUut8.ReverseButton;
   TraceIn_SensorFeed[83] := BenchUut8.SensorFeed;
   TraceIn_SensorWash[83] := BenchUut8.SensorWash;
   TraceIn_SensorWeight[83] := BenchUut8.SensorWeight;
   TraceIn_SensorFiring[83] := BenchUut8.SensorFiring;
   TraceIn_SensorOutput[83] := BenchUut8.SensorOutput;
   TraceIn_washComplete[83] := BenchUut8.washComplete;
   TraceIn_weightComplete[83] := BenchUut8.weightComplete;
   TraceIn_weight[83] := BenchUut8.weight;
   TraceIn_firingComplete[83] := BenchUut8.firingComplete;
   BenchUut8();
   TraceOut_MotorForward[83] := BenchUut8.MotorForward;
   TraceOut_MotorReverse[83] := BenchUut8.MotorReverse;
   TraceOut_kick[83] := BenchUut8.kick;
   TraceOut_CompletionLight[83] := BenchUut8.CompletionLight;
   TraceOut_firingTemp[83] := BenchUut8.firingTemp;
   BenchCalls := BenchCalls + 1;
 84:
   BenchUut8.Mode := TRUE;
   BenchUut8.ForwardButton := FALSE;
   BenchUut8.ReverseButton := FALSE;
   BenchUut8.SensorFeed := FALSE;
   BenchUut8.SensorWash := TRUE;
   BenchUut8.SensorWeight := FALSE;
   BenchUut8.SensorFiring := FALSE;
   BenchUut8.SensorOutput := FALSE;
   BenchUut8.washComplete := FALSE;
   BenchUut8.weightComplete := FALSE;
   BenchUut8.weight := REAL#150.0;
   BenchUut8.firingComplete := FALSE;
   TraceIn_Mode[84] := BenchUut8.Mode;
   TraceIn_ForwardButton[84] := BenchUut8.ForwardButton;
   TraceIn_ReverseButton[84] := BenchUut8.ReverseButton;
   TraceIn_SensorFeed[84] := BenchUut8.SensorFeed;
   TraceIn_SensorWash[84] := BenchUut8.SensorWash;
   TraceIn_SensorWeight[84] := BenchUut8.SensorWeight;
   TraceIn_SensorFiring[84] := BenchUut8.SensorFiring;
   TraceIn_SensorOutput[84] := BenchUut8.SensorOutput;
   TraceIn_washComplete[84] := BenchUut8.washComplete;
   TraceIn_weightComplete[84] := BenchUut8.weightComplete;
   TraceIn_weight[84] := BenchUut8.weight;
   TraceIn_firingComplete[84] := BenchUut8.firingComplete;
   BenchUut8();
   TraceOut_MotorForward[84] := BenchUut8.MotorForward;
   TraceOut_MotorReverse[84] := BenchUut8.MotorReverse;
   TraceOut_kick[84] := BenchUut8.kick;
   TraceOut_CompletionLight[84] := BenchUut8.CompletionLight;
   TraceOut_firingTemp[84] := BenchUut8.firingTemp;
   BenchCalls := BenchCalls + 1;
 85:
   BenchUut8.Mode := TRUE;
   BenchUut8.ForwardButton := FALSE;
   BenchUut8.ReverseButton := FALSE;
   BenchUut8.SensorFeed := FALSE;
   BenchUut8.SensorWash := TRUE;
   BenchUut8.SensorWeight := FALSE;
   BenchUut8.SensorFiring := FALSE;
   BenchUut8.SensorOutput := FALSE;
   BenchUut8.washComplete := TRUE;
   BenchUut8.weightComplete := FALSE;
   BenchUut8.weight := REAL#150.0;
   BenchUut8.firingComplete := FALSE;
   TraceIn_Mode[85] := BenchUut8.Mode;
   TraceIn_ForwardButton[85] := BenchUut8.ForwardButton;
   TraceIn_ReverseButton[85] := BenchUut8.ReverseButton;
   TraceIn_SensorFeed[85] := BenchUut8.SensorFeed;
   TraceIn_SensorWash[85] := BenchUut8.SensorWash;
   TraceIn_SensorWeight[85] := BenchUut8.SensorWeight;
   TraceIn_SensorFiring[85] := BenchUut8.SensorFiring;
   TraceIn_SensorOutput[85] := BenchUut8.SensorOutput;
   TraceIn_washComplete[85] := BenchUut8.washComplete;
   TraceIn_weightComplete[85] := BenchUut8.weightComplete;
   TraceIn_weight[85] := BenchUut8.weight;
   TraceIn_firingComplete[85] := BenchUut8.firingComplete;
   BenchUut8();
   TraceOut_MotorForward[85] := BenchUut8.MotorForward;
   TraceOut_MotorReverse[85] := BenchUut8.MotorReverse;
   TraceOut_kick[85] := BenchUut8.kick;
   TraceOut_CompletionLight[85] := BenchUut8.CompletionLight;
   TraceOut_firingTemp[85] := BenchUut8.firingTemp;
   BenchCalls := BenchCalls + 1;
 86:
   BenchUut8.Mode := TRUE;
   BenchUut8.ForwardButton := FALSE;
   BenchUut8.ReverseButton := FALSE;
   BenchUut8.SensorFeed := FALSE;
   BenchUut8.SensorWash := FALSE;
   BenchUut8.SensorWeight := TRUE;
   BenchUut8.SensorFiring := FALSE;
   BenchUut8.SensorOutput := FALSE;
   BenchUut8.washComplete := FALSE;
   BenchUut8.weightComplete := FALSE;
   BenchUut8.weight := REAL#150.0;
   BenchUut8.firingComplete := FALSE;
   TraceIn_Mode[86] := BenchUut8.Mode;
   TraceIn_ForwardButton[86] := BenchUut8.ForwardButton;
   TraceIn_ReverseButton[86] := BenchUut8.ReverseButton;
   TraceIn_SensorFeed[86] := BenchUut8.SensorFeed;
   TraceIn_SensorWash[86] := BenchUut8.SensorWash;
   TraceIn_SensorWeight[86] := BenchUut8.SensorWeight;
   TraceIn_SensorFiring[86] := BenchUut8.SensorFiring;
   TraceIn_SensorOutput[86] := BenchUut8.SensorOutput;
   TraceIn_washComplete[86] := BenchUut8.washComplete;
   TraceIn_weightComplete[86] := BenchUut8.weightComplete;
   TraceIn_weight[86] := BenchUut8.weight;
   TraceIn_firingComplete[86] := BenchUut8.firingComplete;
   BenchUut8();
   TraceOut_MotorForward[86] := BenchUut8.MotorForward;
   TraceOut_MotorReverse[86] := BenchUut8.MotorReverse;
   TraceOut_kick[86] := BenchUut8.kick;
   TraceOut_CompletionLight[86] := BenchUut8.CompletionLight;
   TraceOut_firingTemp[86] := BenchUut8.firingTemp;
   BenchCalls := BenchCalls + 1;
 87:
   BenchUut8.Mode := TRUE;
   BenchUut8.ForwardButton := FALSE;
   BenchUut8.ReverseButton := FALSE;
   BenchUut8.SensorFeed := FALSE;
   BenchUut8.SensorWash := FALSE;
   BenchUut8.SensorWeight := TRUE;
   BenchUut8.SensorFiring := FALSE;
   BenchUut8.SensorOutput := FALSE;
   BenchUut8.washComplete := FALSE;
   BenchUut8.weightComplete := TRUE;
   BenchUut8.weight := REAL#200.0001;
   BenchUut8.firingComplete := FALSE;
   TraceIn_Mode[87] := BenchUut8.Mode;
   TraceIn_ForwardButton[87] := BenchUut8.ForwardButton;
   TraceIn_ReverseButton[87] := BenchUut8.ReverseButton;
   TraceIn_SensorFeed[87] := BenchUut8.SensorFeed;
   TraceIn_SensorWash[87] := BenchUut8.SensorWash;
   TraceIn_SensorWeight[87] := BenchUut8.SensorWeight;
   TraceIn_SensorFiring[87] := BenchUut8.SensorFiring;
   TraceIn_SensorOutput[87] := BenchUut8.SensorOutput;
   TraceIn_washComplete[87] := BenchUut8.washComplete;
   TraceIn_weightComplete[87] := BenchUut8.weightComplete;
   TraceIn_weight[87] := BenchUut8.weight;
   TraceIn_firingComplete[87] := BenchUut8.firingComplete;
   BenchUut8();
   TraceOut_MotorForward[87] := BenchUut8.MotorForward;
   TraceOut_MotorReverse[87] := BenchUut8.MotorReverse;
   TraceOut_kick[87] := BenchUut8.kick;
   TraceOut_CompletionLight[87] := BenchUut8.CompletionLight;
   TraceOut_firingTemp[87] := BenchUut8.firingTemp;
   BenchCalls := BenchCalls + 1;
 88:
   BenchUut8.Mode := TRUE;
   BenchUut8.ForwardButton := FALSE;
   BenchUut8.ReverseButton := FALSE;
   BenchUut8.SensorFeed := FALSE;
   BenchUut8.SensorWash := FALSE;
   BenchUut8.SensorWeight := FALSE;
   BenchUut8.SensorFiring := FALSE;
   BenchUut8.SensorOutput := FALSE;
   BenchUut8.washComplete := FALSE;
   BenchUut8.weightComplete := FALSE;
   BenchUut8.weight := REAL#150.0;
   BenchUut8.firingComplete := FALSE;
   TraceIn_Mode[88] := BenchUut8.Mode;
   TraceIn_ForwardButton[88] := BenchUut8.ForwardButton;
   TraceIn_ReverseButton[88] := BenchUut8.ReverseButton;
   TraceIn_SensorFeed[88] := BenchUut8.SensorFeed;
   TraceIn_SensorWash[88] := BenchUut8.SensorWash;
   TraceIn_SensorWeight[88] := BenchUut8.SensorWeight;
   TraceIn_SensorFiring[88] := BenchUut8.SensorFiring;
   TraceIn_SensorOutput[88] := BenchUut8.SensorOutput;
   TraceIn_washComplete[88] := BenchUut8.washComplete;
   TraceIn_weightComplete[88] := BenchUut8.weightComplete;
   TraceIn_weight[88] := BenchUut8.weight;
   TraceIn_firingComplete[88] := BenchUut8.firingComplete;
   BenchUut8();
   TraceOut_MotorForward[88] := BenchUut8.MotorForward;
   TraceOut_MotorReverse[88] := BenchUut8.MotorReverse;
   TraceOut_kick[88] := BenchUut8.kick;
   TraceOut_CompletionLight[88] := BenchUut8.CompletionLight;
   TraceOut_firingTemp[88] := BenchUut8.firingTemp;
   BenchCalls := BenchCalls + 1;
 89:
   BenchUut9.Mode := TRUE;
   BenchUut9.ForwardButton := FALSE;
   BenchUut9.ReverseButton := FALSE;
   BenchUut9.SensorFeed := TRUE;
   BenchUut9.SensorWash := FALSE;
   BenchUut9.SensorWeight := FALSE;
   BenchUut9.SensorFiring := FALSE;
   BenchUut9.SensorOutput := FALSE;
   BenchUut9.washComplete := FALSE;
   BenchUut9.weightComplete := FALSE;
   BenchUut9.weight := REAL#150.0;
   BenchUut9.firingComplete := FALSE;
   TraceIn_Mode[89] := BenchUut9.Mode;
   TraceIn_ForwardButton[89] := BenchUut9.ForwardButton;
   TraceIn_ReverseButton[89] := BenchUut9.ReverseButton;
   TraceIn_SensorFeed[89] := BenchUut9.SensorFeed;
   TraceIn_SensorWash[89] := BenchUut9.SensorWash;
   TraceIn_SensorWeight[89] := BenchUut9.SensorWeight;
   TraceIn_SensorFiring[89] := BenchUut9.SensorFiring;
   TraceIn_SensorOutput[89] := BenchUut9.SensorOutput;
   TraceIn_washComplete[89] := BenchUut9.washComplete;
   TraceIn_weightComplete[89] := BenchUut9.weightComplete;
   TraceIn_weight[89] := BenchUut9.weight;
   TraceIn_firingComplete[89] := BenchUut9.firingComplete;
   BenchUut9();
   TraceOut_MotorForward[89] := BenchUut9.MotorForward;
   TraceOut_MotorReverse[89] := BenchUut9.MotorReverse;
   TraceOut_kick[89] := BenchUut9.kick;
   TraceOut_CompletionLight[89] := BenchUut9.CompletionLight;
   TraceOut_firingTemp[89] := BenchUut9.firingTemp;
   BenchCalls := BenchCalls + 1;
 90:
   BenchUut9.Mode := TRUE;
   BenchUut9.ForwardButton := FALSE;
   BenchUut9.ReverseButton := FALSE;
   BenchUut9.SensorFeed := FALSE;
   BenchUut9.SensorWash := FALSE;
   BenchUut9.SensorWeight := FALSE;
   BenchUut9.SensorFiring := FALSE;
   BenchUut9.SensorOutput := FALSE;
   BenchUut9.washComplete := FALSE;
   BenchUut9.weightComplete := FALSE;
   BenchUut9.weight := REAL#150.0;
   BenchUut9.firingComplete := FALSE;
   TraceIn_Mode[90] := BenchUut9.Mode;
   TraceIn_ForwardButton[90] := BenchUut9.ForwardButton;
   TraceIn_ReverseButton[90] := BenchUut9.ReverseButton;
   TraceIn_SensorFeed[90] := BenchUut9.SensorFeed;
   TraceIn_SensorWash[90] := BenchUut9.SensorWash;
   TraceIn_SensorWeight[90] := BenchUut9.SensorWeight;
   TraceIn_SensorFiring[90] := BenchUut9.SensorFiring;
   TraceIn_SensorOutput[90] := BenchUut9.SensorOutput;
   TraceIn_washComplete[90] := BenchUut9.washComplete;
   TraceIn_weightComplete[90] := BenchUut9.weightComplete;
   TraceIn_weight[90] := BenchUut9.weight;
   TraceIn_firingComplete[90] := BenchUut9.firingComplete;
   BenchUut9();
   TraceOut_MotorForward[90] := BenchUut9.MotorForward;
   TraceOut_MotorReverse[90] := BenchUut9.MotorReverse;
   TraceOut_kick[90] := BenchUut9.kick;
   TraceOut_CompletionLight[90] := BenchUut9.CompletionLight;
   TraceOut_firingTemp[90] := BenchUut9.firingTemp;
   BenchCalls := BenchCalls + 1;
 91:
   BenchUut9.Mode := TRUE;
   BenchUut9.ForwardButton := FALSE;
   BenchUut9.ReverseButton := FALSE;
   BenchUut9.SensorFeed := FALSE;
   BenchUut9.SensorWash := FALSE;
   BenchUut9.SensorWeight := FALSE;
   BenchUut9.SensorFiring := FALSE;
   BenchUut9.SensorOutput := FALSE;
   BenchUut9.washComplete := FALSE;
   BenchUut9.weightComplete := FALSE;
   BenchUut9.weight := REAL#150.0;
   BenchUut9.firingComplete := FALSE;
   TraceIn_Mode[91] := BenchUut9.Mode;
   TraceIn_ForwardButton[91] := BenchUut9.ForwardButton;
   TraceIn_ReverseButton[91] := BenchUut9.ReverseButton;
   TraceIn_SensorFeed[91] := BenchUut9.SensorFeed;
   TraceIn_SensorWash[91] := BenchUut9.SensorWash;
   TraceIn_SensorWeight[91] := BenchUut9.SensorWeight;
   TraceIn_SensorFiring[91] := BenchUut9.SensorFiring;
   TraceIn_SensorOutput[91] := BenchUut9.SensorOutput;
   TraceIn_washComplete[91] := BenchUut9.washComplete;
   TraceIn_weightComplete[91] := BenchUut9.weightComplete;
   TraceIn_weight[91] := BenchUut9.weight;
   TraceIn_firingComplete[91] := BenchUut9.firingComplete;
   BenchUut9();
   TraceOut_MotorForward[91] := BenchUut9.MotorForward;
   TraceOut_MotorReverse[91] := BenchUut9.MotorReverse;
   TraceOut_kick[91] := BenchUut9.kick;
   TraceOut_CompletionLight[91] := BenchUut9.CompletionLight;
   TraceOut_firingTemp[91] := BenchUut9.firingTemp;
   BenchCalls := BenchCalls + 1;
 92:
   BenchUut9.Mode := TRUE;
   BenchUut9.ForwardButton := FALSE;
   BenchUut9.ReverseButton := FALSE;
   BenchUut9.SensorFeed := FALSE;
   BenchUut9.SensorWash := FALSE;
   BenchUut9.SensorWeight := FALSE;
   BenchUut9.SensorFiring := FALSE;
   BenchUut9.SensorOutput := FALSE;
   BenchUut9.washComplete := FALSE;
   BenchUut9.weightComplete := FALSE;
   BenchUut9.weight := REAL#150.0;
   BenchUut9.firingComplete := FALSE;
   TraceIn_Mode[92] := BenchUut9.Mode;
   TraceIn_ForwardButton[92] := BenchUut9.ForwardButton;
   TraceIn_ReverseButton[92] := BenchUut9.ReverseButton;
   TraceIn_SensorFeed[92] := BenchUut9.SensorFeed;
   TraceIn_SensorWash[92] := BenchUut9.SensorWash;
   TraceIn_SensorWeight[92] := BenchUut9.SensorWeight;
   TraceIn_SensorFiring[92] := BenchUut9.SensorFiring;
   TraceIn_SensorOutput[92] := BenchUut9.SensorOutput;
   TraceIn_washComplete[92] := BenchUut9.washComplete;
   TraceIn_weightComplete[92] := BenchUut9.weightComplete;
   TraceIn_weight[92] := BenchUut9.weight;
   TraceIn_firingComplete[92] := BenchUut9.firingComplete;
   BenchUut9();
   TraceOut_MotorForward[92] := BenchUut9.MotorForward;
   TraceOut_MotorReverse[92] := BenchUut9.MotorReverse;
   TraceOut_kick[92] := BenchUut9.kick;
   TraceOut_CompletionLight[92] := BenchUut9.CompletionLight;
   TraceOut_firingTemp[92] := BenchUut9.firingTemp;
   BenchCalls := BenchCalls + 1;
 93:
   BenchUut9.Mode := TRUE;
   BenchUut9.ForwardButton := FALSE;
   BenchUut9.ReverseButton := FALSE;
   BenchUut9.SensorFeed := FALSE;
   BenchUut9.SensorWash := TRUE;
   BenchUut9.SensorWeight := FALSE;
   BenchUut9.SensorFiring := FALSE;
   BenchUut9.SensorOutput := FALSE;
   BenchUut9.washComplete := FALSE;
   BenchUut9.weightComplete := FALSE;
   BenchUut9.weight := REAL#150.0;
   BenchUut9.firingComplete := FALSE;
   TraceIn_Mode[93] := BenchUut9.Mode;
   TraceIn_ForwardButton[93] := BenchUut9.ForwardButton;
   TraceIn_ReverseButton[93] := BenchUut9.ReverseButton;
   TraceIn_SensorFeed[93] := BenchUut9.SensorFeed;
   TraceIn_SensorWash[93] := BenchUut9.SensorWash;
   TraceIn_SensorWeight[93] := BenchUut9.SensorWeight;
   TraceIn_SensorFiring[93] := BenchUut9.SensorFiring;
   TraceIn_SensorOutput[93] := BenchUut9.SensorOutput;
   TraceIn_washComplete[93] := BenchUut9.washComplete;
   TraceIn_weightComplete[93] := BenchUut9.weightComplete;
   TraceIn_weight[93] := BenchUut9.weight;
   TraceIn_firingComplete[93] := BenchUut9.firingComplete;
   BenchUut9();
   TraceOut_MotorForward[93] := BenchUut9.MotorForward;
   TraceOut_MotorReverse[93] := BenchUut9.MotorReverse;
   TraceOut_kick[93] := BenchUut9.kick;
   TraceOut_CompletionLight[93] := BenchUut9.CompletionLight;
   TraceOut_firingTemp[93] := BenchUut9.firingTemp;
   BenchCalls := BenchCalls + 1;
 94:
   BenchUut9.Mode := TRUE;
   BenchUut9.ForwardButton := FALSE;
   BenchUut9.ReverseButton := FALSE;
   BenchUut9.SensorFeed := FALSE;
   BenchUut9.SensorWash := TRUE;
   BenchUut9.SensorWeight := FALSE;
   BenchUut9.SensorFiring := FALSE;
   BenchUut9.SensorOutput := FALSE;
   BenchUut9.washComplete := FALSE;
   BenchUut9.weightComplete := FALSE;
   BenchUut9.weight := REAL#150.0;
   BenchUut9.firingComplete := FALSE;
   TraceIn_Mode[94] := BenchUut9.Mode;
   TraceIn_ForwardButton[94] := BenchUut9.ForwardButton;
   TraceIn_ReverseButton[94] := BenchUut9.ReverseButton;
   TraceIn_SensorFeed[94] := BenchUut9.SensorFeed;
   TraceIn_SensorWash[94] := BenchUut9.SensorWash;
   TraceIn_SensorWeight[94] := BenchUut9.SensorWeight;
   TraceIn_SensorFiring[94] := BenchUut9.SensorFiring;
   TraceIn_SensorOutput[94] := BenchUut9.SensorOutput;
   TraceIn_washComplete[94] := BenchUut9.washComplete;
   TraceIn_weightComplete[94] := BenchUut9.weightComplete;
   TraceIn_weight[94] := BenchUut9.weight;
   TraceIn_firingComplete[94] := BenchUut9.firingComplete;
   BenchUut9();
   TraceOut_MotorForward[94] := BenchUut9.MotorForward;
   TraceOut_MotorReverse[94] := BenchUut9.MotorReverse;
   TraceOut_kick[94] := BenchUut9.kick;
   TraceOut_CompletionLight[94] := BenchUut9.CompletionLight;
   TraceOut_firingTemp[94] := BenchUut9.firingTemp;
   BenchCalls := BenchCalls + 1;
 95:
   BenchUut9.Mode := TRUE;
   BenchUut9.ForwardButton := FALSE;
   BenchUut9.ReverseButton := FALSE;
   BenchUut9.SensorFeed := FALSE;
   BenchUut9.SensorWash := TRUE;
   BenchUut9.SensorWeight := FALSE;
   BenchUut9.SensorFiring := FALSE;
   BenchUut9.SensorOutput := FALSE;
   BenchUut9.washComplete := FALSE;
   BenchUut9.weightComplete := FALSE;
   BenchUut9.weight := REAL#150.0;
   BenchUut9.firingComplete := FALSE;
   TraceIn_Mode[95] := BenchUut9.Mode;
   TraceIn_ForwardButton[95] := BenchUut9.ForwardButton;
   TraceIn_ReverseButton[95] := BenchUut9.ReverseButton;
   TraceIn_SensorFeed[95] := BenchUut9.SensorFeed;
   TraceIn_SensorWash[95] := BenchUut9.SensorWash;
   TraceIn_SensorWeight[95] := BenchUut9.SensorWeight;
   TraceIn_SensorFiring[95] := BenchUut9.SensorFiring;
   TraceIn_SensorOutput[95] := BenchUut9.SensorOutput;
   TraceIn_washComplete[95] := BenchUut9.washComplete;
   TraceIn_weightComplete[95] := BenchUut9.weightComplete;
   TraceIn_weight[95] := BenchUut9.weight;
   TraceIn_firingComplete[95] := BenchUut9.firingComplete;
   BenchUut9();
   TraceOut_MotorForward[95] := BenchUut9.MotorForward;
   TraceOut_MotorReverse[95] := BenchUut9.MotorReverse;
   TraceOut_kick[95] := BenchUut9.kick;
   TraceOut_CompletionLight[95] := BenchUut9.CompletionLight;
   TraceOut_firingTemp[95] := BenchUut9.firingTemp;
   BenchCalls := BenchCalls + 1;
 96:
   BenchUut9.Mode := TRUE;
   BenchUut9.ForwardButton := FALSE;
   BenchUut9.ReverseButton := FALSE;
   BenchUut9.SensorFeed := FALSE;
   BenchUut9.SensorWash := TRUE;
   BenchUut9.SensorWeight := FALSE;
   BenchUut9.SensorFiring := FALSE;
   BenchUut9.SensorOutput := FALSE;
   BenchUut9.washComplete := TRUE;
   BenchUut9.weightComplete := FALSE;
   BenchUut9.weight := REAL#150.0;
   BenchUut9.firingComplete := FALSE;
   TraceIn_Mode[96] := BenchUut9.Mode;
   TraceIn_ForwardButton[96] := BenchUut9.ForwardButton;
   TraceIn_ReverseButton[96] := BenchUut9.ReverseButton;
   TraceIn_SensorFeed[96] := BenchUut9.SensorFeed;
   TraceIn_SensorWash[96] := BenchUut9.SensorWash;
   TraceIn_SensorWeight[96] := BenchUut9.SensorWeight;
   TraceIn_SensorFiring[96] := BenchUut9.SensorFiring;
   TraceIn_SensorOutput[96] := BenchUut9.SensorOutput;
   TraceIn_washComplete[96] := BenchUut9.washComplete;
   TraceIn_weightComplete[96] := BenchUut9.weightComplete;
   TraceIn_weight[96] := BenchUut9.weight;
   TraceIn_firingComplete[96] := BenchUut9.firingComplete;
   BenchUut9();
   TraceOut_MotorForward[96] := BenchUut9.MotorForward;
   TraceOut_MotorReverse[96] := BenchUut9.MotorReverse;
   TraceOut_kick[96] := BenchUut9.kick;
   TraceOut_CompletionLight[96] := BenchUut9.CompletionLight;
   TraceOut_firingTemp[96] := BenchUut9.firingTemp;
   BenchCalls := BenchCalls + 1;
 97:
   BenchUut9.Mode := TRUE;
   BenchUut9.ForwardButton := FALSE;
   BenchUut9.ReverseButton := FALSE;
   BenchUut9.SensorFeed := FALSE;
   BenchUut9.SensorWash := FALSE;
   BenchUut9.SensorWeight := FALSE;
   BenchUut9.SensorFiring := FALSE;
   BenchUut9.SensorOutput := FALSE;
   BenchUut9.washComplete := FALSE;
   BenchUut9.weightComplete := FALSE;
   BenchUut9.weight := REAL#150.0;
   BenchUut9.firingComplete := FALSE;
   TraceIn_Mode[97] := BenchUut9.Mode;
   TraceIn_ForwardButton[97] := BenchUut9.ForwardButton;
   TraceIn_ReverseButton[97] := BenchUut9.ReverseButton;
   TraceIn_SensorFeed[97] := BenchUut9.SensorFeed;
   TraceIn_SensorWash[97] := BenchUut9.SensorWash;
   TraceIn_SensorWeight[97] := BenchUut9.SensorWeight;
   TraceIn_SensorFiring[97] := BenchUut9.SensorFiring;
   TraceIn_SensorOutput[97] := BenchUut9.SensorOutput;
   TraceIn_washComplete[97] := BenchUut9.washComplete;
   TraceIn_weightComplete[97] := BenchUut9.weightComplete;
   TraceIn_weight[97] := BenchUut9.weight;
   TraceIn_firingComplete[97] := BenchUut9.firingComplete;
   BenchUut9();
   TraceOut_MotorForward[97] := BenchUut9.MotorForward;
   TraceOut_MotorReverse[97] := BenchUut9.MotorReverse;
   TraceOut_kick[97] := BenchUut9.kick;
   TraceOut_CompletionLight[97] := BenchUut9.CompletionLight;
   TraceOut_firingTemp[97] := BenchUut9.firingTemp;
   BenchCalls := BenchCalls + 1;
 98:
   BenchUut9.Mode := TRUE;
   BenchUut9.ForwardButton := FALSE;
   BenchUut9.ReverseButton := FALSE;
   BenchUut9.SensorFeed := FALSE;
   BenchUut9.SensorWash := FALSE;
   BenchUut9.SensorWeight := FALSE;
   BenchUut9.SensorFiring := FALSE;
   BenchUut9.SensorOutput := FALSE;
   BenchUut9.washComplete := FALSE;
   BenchUut9.weightComplete := FALSE;
   BenchUut9.weight := REAL#150.0;
   BenchUut9.firingComplete := FALSE;
   TraceIn_Mode[98] := BenchUut9.Mode;
   TraceIn_ForwardButton[98] := BenchUut9.ForwardButton;
   TraceIn_ReverseButton[98] := BenchUut9.ReverseButton;
   TraceIn_SensorFeed[98] := BenchUut9.SensorFeed;
   TraceIn_SensorWash[98] := BenchUut9.SensorWash;
   TraceIn_SensorWeight[98] := BenchUut9.SensorWeight;
   TraceIn_SensorFiring[98] := BenchUut9.SensorFiring;
   TraceIn_SensorOutput[98] := BenchUut9.SensorOutput;
   TraceIn_washComplete[98] := BenchUut9.washComplete;
   TraceIn_weightComplete[98] := BenchUut9.weightComplete;
   TraceIn_weight[98] := BenchUut9.weight;
   TraceIn_firingComplete[98] := BenchUut9.firingComplete;
   BenchUut9();
   TraceOut_MotorForward[98] := BenchUut9.MotorForward;
   TraceOut_MotorReverse[98] := BenchUut9.MotorReverse;
   TraceOut_kick[98] := BenchUut9.kick;
   TraceOut_CompletionLight[98] := BenchUut9.CompletionLight;
   TraceOut_firingTemp[98] := BenchUut9.firingTemp;
   BenchCalls := BenchCalls + 1;
 99:
   BenchUut9.Mode := TRUE;
   BenchUut9.ForwardButton := FALSE;
   BenchUut9.ReverseButton := FALSE;
   BenchUut9.SensorFeed := FALSE;
   BenchUut9.SensorWash := FALSE;
   BenchUut9.SensorWeight := FALSE;
   BenchUut9.SensorFiring := FALSE;
   BenchUut9.SensorOutput := FALSE;
   BenchUut9.washComplete := FALSE;
   BenchUut9.weightComplete := FALSE;
   BenchUut9.weight := REAL#150.0;
   BenchUut9.firingComplete := FALSE;
   TraceIn_Mode[99] := BenchUut9.Mode;
   TraceIn_ForwardButton[99] := BenchUut9.ForwardButton;
   TraceIn_ReverseButton[99] := BenchUut9.ReverseButton;
   TraceIn_SensorFeed[99] := BenchUut9.SensorFeed;
   TraceIn_SensorWash[99] := BenchUut9.SensorWash;
   TraceIn_SensorWeight[99] := BenchUut9.SensorWeight;
   TraceIn_SensorFiring[99] := BenchUut9.SensorFiring;
   TraceIn_SensorOutput[99] := BenchUut9.SensorOutput;
   TraceIn_washComplete[99] := BenchUut9.washComplete;
   TraceIn_weightComplete[99] := BenchUut9.weightComplete;
   TraceIn_weight[99] := BenchUut9.weight;
   TraceIn_firingComplete[99] := BenchUut9.firingComplete;
   BenchUut9();
   TraceOut_MotorForward[99] := BenchUut9.MotorForward;
   TraceOut_MotorReverse[99] := BenchUut9.MotorReverse;
   TraceOut_kick[99] := BenchUut9.kick;
   TraceOut_CompletionLight[99] := BenchUut9.CompletionLight;
   TraceOut_firingTemp[99] := BenchUut9.firingTemp;
   BenchCalls := BenchCalls + 1;
 100:
   BenchUut9.Mode := TRUE;
   BenchUut9.ForwardButton := FALSE;
   BenchUut9.ReverseButton := FALSE;
   BenchUut9.SensorFeed := FALSE;
   BenchUut9.SensorWash := FALSE;
   BenchUut9.SensorWeight := TRUE;
   BenchUut9.SensorFiring := FALSE;
   BenchUut9.SensorOutput := FALSE;
   BenchUut9.washComplete := FALSE;
   BenchUut9.weightComplete := FALSE;
   BenchUut9.weight := REAL#150.0;
   BenchUut9.firingComplete := FALSE;
   TraceIn_Mode[100] := BenchUut9.Mode;
   TraceIn_ForwardButton[100] := BenchUut9.ForwardButton;
   TraceIn_ReverseButton[100] := BenchUut9.ReverseButton;
   TraceIn_SensorFeed[100] := BenchUut9.SensorFeed;
   TraceIn_SensorWash[100] := BenchUut9.SensorWash;
   TraceIn_SensorWeight[100] := BenchUut9.SensorWeight;
   TraceIn_SensorFiring[100] := BenchUut9.SensorFiring;
   TraceIn_SensorOutput[100] := BenchUut9.SensorOutput;
   TraceIn_washComplete[100] := BenchUut9.washComplete;
   TraceIn_weightComplete[100] := BenchUut9.weightComplete;
   TraceIn_weight[100] := BenchUut9.weight;
   TraceIn_firingComplete[100] := BenchUut9.firingComplete;
   BenchUut9();
   TraceOut_MotorForward[100] := BenchUut9.MotorForward;
   TraceOut_MotorReverse[100] := BenchUut9.MotorReverse;
   TraceOut_kick[100] := BenchUut9.kick;
   TraceOut_CompletionLight[100] := BenchUut9.CompletionLight;
   TraceOut_firingTemp[100] := BenchUut9.firingTemp;
   BenchCalls := BenchCalls + 1;
 101:
   BenchUut9.Mode := TRUE;
   BenchUut9.ForwardButton := FALSE;
   BenchUut9.ReverseButton := FALSE;
   BenchUut9.SensorFeed := FALSE;
   BenchUut9.SensorWash := FALSE;
   BenchUut9.SensorWeight := TRUE;
   BenchUut9.SensorFiring := FALSE;
   BenchUut9.SensorOutput := FALSE;
   BenchUut9.washComplete := FALSE;
   BenchUut9.weightComplete := FALSE;
   BenchUut9.weight := REAL#150.0;
   BenchUut9.firingComplete := FALSE;
   TraceIn_Mode[101] := BenchUut9.Mode;
   TraceIn_ForwardButton[101] := BenchUut9.ForwardButton;
   TraceIn_ReverseButton[101] := BenchUut9.ReverseButton;
   TraceIn_SensorFeed[101] := BenchUut9.SensorFeed;
   TraceIn_SensorWash[101] := BenchUut9.SensorWash;
   TraceIn_SensorWeight[101] := BenchUut9.SensorWeight;
   TraceIn_SensorFiring[101] := BenchUut9.SensorFiring;
   TraceIn_SensorOutput[101] := BenchUut9.SensorOutput;
   TraceIn_washComplete[101] := BenchUut9.washComplete;
   TraceIn_weightComplete[101] := BenchUut9.weightComplete;
   TraceIn_weight[101] := BenchUut9.weight;
   TraceIn_firingComplete[101] := BenchUut9.firingComplete;
   BenchUut9();
   TraceOut_MotorForward[101] := BenchUut9.MotorForward;
   TraceOut_MotorReverse[101] := BenchUut9.MotorReverse;
   TraceOut_kick[101] := BenchUut9.kick;
   TraceOut_CompletionLight[101] := BenchUut9.CompletionLight;
   TraceOut_firingTemp[101] := BenchUut9.firingTemp;
   BenchCalls := BenchCalls + 1;
 102:
   BenchUut9.Mode := TRUE;
   BenchUut9.ForwardButton := FALSE;
   BenchUut9.ReverseButton := FALSE;
   BenchUut9.SensorFeed := FALSE;
   BenchUut9.SensorWash := FALSE;
   BenchUut9.SensorWeight := TRUE;
   BenchUut9.SensorFiring := FALSE;
   BenchUut9.SensorOutput := FALSE;
   BenchUut9.washComplete := FALSE;
   BenchUut9.weightComplete := FALSE;
   BenchUut9.weight := REAL#150.0;
   BenchUut9.firingComplete := FALSE;
   TraceIn_Mode[102] := BenchUut9.Mode;
   TraceIn_ForwardButton[102] := BenchUut9.ForwardButton;
   TraceIn_ReverseButton[102] := BenchUut9.ReverseButton;
   TraceIn_SensorFeed[102] := BenchUut9.SensorFeed;
   TraceIn_SensorWash[102] := BenchUut9.SensorWash;
   TraceIn_SensorWeight[102] := BenchUut9.SensorWeight;
   TraceIn_SensorFiring[102] := BenchUut9.SensorFiring;
   TraceIn_SensorOutput[102] := BenchUut9.SensorOutput;
   TraceIn_washComplete[102] := BenchUut9.washComplete;
   TraceIn_weightComplete[102] := BenchUut9.weightComplete;
   TraceIn_weight[102] := BenchUut9.weight;
   TraceIn_firingComplete[102] := BenchUut9.firingComplete;
   BenchUut9();
   TraceOut_MotorForward[102] := BenchUut9.MotorForward;
   TraceOut_MotorReverse[102] := BenchUut9.MotorReverse;
   TraceOut_kick[102] := BenchUut9.kick;
   TraceOut_CompletionLight[102] := BenchUut9.CompletionLight;
   TraceOut_firingTemp[102] := BenchUut9.firingTemp;
   BenchCalls := BenchCalls + 1;
 103:
   BenchUut9.Mode := TRUE;
   BenchUut9.ForwardButton := FALSE;
   BenchUut9.ReverseButton := FALSE;
   BenchUut9.SensorFeed := FALSE;
   BenchUut9.SensorWash := FALSE;
   BenchUut9.SensorWeight := TRUE;
   BenchUut9.SensorFiring := FALSE;
   BenchUut9.SensorOutput := FALSE;
   BenchUut9.washComplete := FALSE;
   BenchUut9.weightComplete := TRUE;
   BenchUut9.weight := REAL#150.0;
   BenchUut9.firingComplete := FALSE;
   TraceIn_Mode[103] := BenchUut9.Mode;
   TraceIn_ForwardButton[103] := BenchUut9.ForwardButton;
   TraceIn_ReverseButton[103] := BenchUut9.ReverseButton;
   TraceIn_SensorFeed[103] := BenchUut9.SensorFeed;
   TraceIn_SensorWash[103] := BenchUut9.SensorWash;
   TraceIn_SensorWeight[103] := BenchUut9.SensorWeight;
   TraceIn_SensorFiring[103] := BenchUut9.SensorFiring;
   TraceIn_SensorOutput[103] := BenchUut9.SensorOutput;
   TraceIn_washComplete[103] := BenchUut9.washComplete;
   TraceIn_weightComplete[103] := BenchUut9.weightComplete;
   TraceIn_weight[103] := BenchUut9.weight;
   TraceIn_firingComplete[103] := BenchUut9.firingComplete;
   BenchUut9();
   TraceOut_MotorForward[103] := BenchUut9.MotorForward;
   TraceOut_MotorReverse[103] := BenchUut9.MotorReverse;
   TraceOut_kick[103] := BenchUut9.kick;
   TraceOut_CompletionLight[103] := BenchUut9.CompletionLight;
   TraceOut_firingTemp[103] := BenchUut9.firingTemp;
   BenchCalls := BenchCalls + 1;
 104:
   BenchUut9.Mode := TRUE;
   BenchUut9.ForwardButton := FALSE;
   BenchUut9.ReverseButton := FALSE;
   BenchUut9.SensorFeed := FALSE;
   BenchUut9.SensorWash := FALSE;
   BenchUut9.SensorWeight := FALSE;
   BenchUut9.SensorFiring := FALSE;
   BenchUut9.SensorOutput := FALSE;
   BenchUut9.washComplete := FALSE;
   BenchUut9.weightComplete := FALSE;
   BenchUut9.weight := REAL#150.0;
   BenchUut9.firingComplete := FALSE;
   TraceIn_Mode[104] := BenchUut9.Mode;
   TraceIn_ForwardButton[104] := BenchUut9.ForwardButton;
   TraceIn_ReverseButton[104] := BenchUut9.ReverseButton;
   TraceIn_SensorFeed[104] := BenchUut9.SensorFeed;
   TraceIn_SensorWash[104] := BenchUut9.SensorWash;
   TraceIn_SensorWeight[104] := BenchUut9.SensorWeight;
   TraceIn_SensorFiring[104] := BenchUut9.SensorFiring;
   TraceIn_SensorOutput[104] := BenchUut9.SensorOutput;
   TraceIn_washComplete[104] := BenchUut9.washComplete;
   TraceIn_weightComplete[104] := BenchUut9.weightComplete;
   TraceIn_weight[104] := BenchUut9.weight;
   TraceIn_firingComplete[104] := BenchUut9.firingComplete;
   BenchUut9();
   TraceOut_MotorForward[104] := BenchUut9.MotorForward;
   TraceOut_MotorReverse[104] := BenchUut9.MotorReverse;
   TraceOut_kick[104] := BenchUut9.kick;
   TraceOut_CompletionLight[104] := BenchUut9.CompletionLight;
   TraceOut_firingTemp[104] := BenchUut9.firingTemp;
   BenchCalls := BenchCalls + 1;
 105:
   BenchUut9.Mode := TRUE;
   BenchUut9.ForwardButton := FALSE;
   BenchUut9.ReverseButton := FALSE;
   BenchUut9.SensorFeed := FALSE;
   BenchUut9.SensorWash := FALSE;
   BenchUut9.SensorWeight := FALSE;
   BenchUut9.SensorFiring := FALSE;
   BenchUut9.SensorOutput := FALSE;
   BenchUut9.washComplete := FALSE;
   BenchUut9.weightComplete := FALSE;
   BenchUut9.weight := REAL#150.0;
   BenchUut9.firingComplete := FALSE;
   TraceIn_Mode[105] := BenchUut9.Mode;
   TraceIn_ForwardButton[105] := BenchUut9.ForwardButton;
   TraceIn_ReverseButton[105] := BenchUut9.ReverseButton;
   TraceIn_SensorFeed[105] := BenchUut9.SensorFeed;
   TraceIn_SensorWash[105] := BenchUut9.SensorWash;
   TraceIn_SensorWeight[105] := BenchUut9.SensorWeight;
   TraceIn_SensorFiring[105] := BenchUut9.SensorFiring;
   TraceIn_SensorOutput[105] := BenchUut9.SensorOutput;
   TraceIn_washComplete[105] := BenchUut9.washComplete;
   TraceIn_weightComplete[105] := BenchUut9.weightComplete;
   TraceIn_weight[105] := BenchUut9.weight;
   TraceIn_firingComplete[105] := BenchUut9.firingComplete;
   BenchUut9();
   TraceOut_MotorForward[105] := BenchUut9.MotorForward;
   TraceOut_MotorReverse[105] := BenchUut9.MotorReverse;
   TraceOut_kick[105] := BenchUut9.kick;
   TraceOut_CompletionLight[105] := BenchUut9.CompletionLight;
   TraceOut_firingTemp[105] := BenchUut9.firingTemp;
   BenchCalls := BenchCalls + 1;
 106:
   BenchUut9.Mode := TRUE;
   BenchUut9.ForwardButton := FALSE;
   BenchUut9.ReverseButton := FALSE;
   BenchUut9.SensorFeed := FALSE;
   BenchUut9.SensorWash := FALSE;
   BenchUut9.SensorWeight := FALSE;
   BenchUut9.SensorFiring := FALSE;
   BenchUut9.SensorOutput := FALSE;
   BenchUut9.washComplete := FALSE;
   BenchUut9.weightComplete := FALSE;
   BenchUut9.weight := REAL#150.0;
   BenchUut9.firingComplete := FALSE;
   TraceIn_Mode[106] := BenchUut9.Mode;
   TraceIn_ForwardButton[106] := BenchUut9.ForwardButton;
   TraceIn_ReverseButton[106] := BenchUut9.ReverseButton;
   TraceIn_SensorFeed[106] := BenchUut9.SensorFeed;
   TraceIn_SensorWash[106] := BenchUut9.SensorWash;
   TraceIn_SensorWeight[106] := BenchUut9.SensorWeight;
   TraceIn_SensorFiring[106] := BenchUut9.SensorFiring;
   TraceIn_SensorOutput[106] := BenchUut9.SensorOutput;
   TraceIn_washComplete[106] := BenchUut9.washComplete;
   TraceIn_weightComplete[106] := BenchUut9.weightComplete;
   TraceIn_weight[106] := BenchUut9.weight;
   TraceIn_firingComplete[106] := BenchUut9.firingComplete;
   BenchUut9();
   TraceOut_MotorForward[106] := BenchUut9.MotorForward;
   TraceOut_MotorReverse[106] := BenchUut9.MotorReverse;
   TraceOut_kick[106] := BenchUut9.kick;
   TraceOut_CompletionLight[106] := BenchUut9.CompletionLight;
   TraceOut_firingTemp[106] := BenchUut9.firingTemp;
   BenchCalls := BenchCalls + 1;
 107:
   BenchUut9.Mode := TRUE;
   BenchUut9.ForwardButton := FALSE;
   BenchUut9.ReverseButton := FALSE;
   BenchUut9.SensorFeed := FALSE;
   BenchUut9.SensorWash := FALSE;
   BenchUut9.SensorWeight := FALSE;
   BenchUut9.SensorFiring := TRUE;
   BenchUut9.SensorOutput := FALSE;
   BenchUut9.washComplete := FALSE;
   BenchUut9.weightComplete := FALSE;
   BenchUut9.weight := REAL#150.0;
   BenchUut9.firingComplete := FALSE;
   TraceIn_Mode[107] := BenchUut9.Mode;
   TraceIn_ForwardButton[107] := BenchUut9.ForwardButton;
   TraceIn_ReverseButton[107] := BenchUut9.ReverseButton;
   TraceIn_SensorFeed[107] := BenchUut9.SensorFeed;
   TraceIn_SensorWash[107] := BenchUut9.SensorWash;
   TraceIn_SensorWeight[107] := BenchUut9.SensorWeight;
   TraceIn_SensorFiring[107] := BenchUut9.SensorFiring;
   TraceIn_SensorOutput[107] := BenchUut9.SensorOutput;
   TraceIn_washComplete[107] := BenchUut9.washComplete;
   TraceIn_weightComplete[107] := BenchUut9.weightComplete;
   TraceIn_weight[107] := BenchUut9.weight;
   TraceIn_firingComplete[107] := BenchUut9.firingComplete;
   BenchUut9();
   TraceOut_MotorForward[107] := BenchUut9.MotorForward;
   TraceOut_MotorReverse[107] := BenchUut9.MotorReverse;
   TraceOut_kick[107] := BenchUut9.kick;
   TraceOut_CompletionLight[107] := BenchUut9.CompletionLight;
   TraceOut_firingTemp[107] := BenchUut9.firingTemp;
   BenchCalls := BenchCalls + 1;
 108:
   BenchUut9.Mode := TRUE;
   BenchUut9.ForwardButton := FALSE;
   BenchUut9.ReverseButton := FALSE;
   BenchUut9.SensorFeed := FALSE;
   BenchUut9.SensorWash := FALSE;
   BenchUut9.SensorWeight := FALSE;
   BenchUut9.SensorFiring := TRUE;
   BenchUut9.SensorOutput := FALSE;
   BenchUut9.washComplete := FALSE;
   BenchUut9.weightComplete := FALSE;
   BenchUut9.weight := REAL#150.0;
   BenchUut9.firingComplete := FALSE;
   TraceIn_Mode[108] := BenchUut9.Mode;
   TraceIn_ForwardButton[108] := BenchUut9.ForwardButton;
   TraceIn_ReverseButton[108] := BenchUut9.ReverseButton;
   TraceIn_SensorFeed[108] := BenchUut9.SensorFeed;
   TraceIn_SensorWash[108] := BenchUut9.SensorWash;
   TraceIn_SensorWeight[108] := BenchUut9.SensorWeight;
   TraceIn_SensorFiring[108] := BenchUut9.SensorFiring;
   TraceIn_SensorOutput[108] := BenchUut9.SensorOutput;
   TraceIn_washComplete[108] := BenchUut9.washComplete;
   TraceIn_weightComplete[108] := BenchUut9.weightComplete;
   TraceIn_weight[108] := BenchUut9.weight;
   TraceIn_firingComplete[108] := BenchUut9.firingComplete;
   BenchUut9();
   TraceOut_MotorForward[108] := BenchUut9.MotorForward;
   TraceOut_MotorReverse[108] := BenchUut9.MotorReverse;
   TraceOut_kick[108] := BenchUut9.kick;
   TraceOut_CompletionLight[108] := BenchUut9.CompletionLight;
   TraceOut_firingTemp[108] := BenchUut9.firingTemp;
   BenchCalls := BenchCalls + 1;
 109:
   BenchUut9.Mode := TRUE;
   BenchUut9.ForwardButton := FALSE;
   BenchUut9.ReverseButton := FALSE;
   BenchUut9.SensorFeed := FALSE;
   BenchUut9.SensorWash := FALSE;
   BenchUut9.SensorWeight := FALSE;
   BenchUut9.SensorFiring := TRUE;
   BenchUut9.SensorOutput := FALSE;
   BenchUut9.washComplete := FALSE;
   BenchUut9.weightComplete := FALSE;
   BenchUut9.weight := REAL#150.0;
   BenchUut9.firingComplete := FALSE;
   TraceIn_Mode[109] := BenchUut9.Mode;
   TraceIn_ForwardButton[109] := BenchUut9.ForwardButton;
   TraceIn_ReverseButton[109] := BenchUut9.ReverseButton;
   TraceIn_SensorFeed[109] := BenchUut9.SensorFeed;
   TraceIn_SensorWash[109] := BenchUut9.SensorWash;
   TraceIn_SensorWeight[109] := BenchUut9.SensorWeight;
   TraceIn_SensorFiring[109] := BenchUut9.SensorFiring;
   TraceIn_SensorOutput[109] := BenchUut9.SensorOutput;
   TraceIn_washComplete[109] := BenchUut9.washComplete;
   TraceIn_weightComplete[109] := BenchUut9.weightComplete;
   TraceIn_weight[109] := BenchUut9.weight;
   TraceIn_firingComplete[109] := BenchUut9.firingComplete;
   BenchUut9();
   TraceOut_MotorForward[109] := BenchUut9.MotorForward;
   TraceOut_MotorReverse[109] := BenchUut9.MotorReverse;
   TraceOut_kick[109] := BenchUut9.kick;
   TraceOut_CompletionLight[109] := BenchUut9.CompletionLight;
   TraceOut_firingTemp[109] := BenchUut9.firingTemp;
   BenchCalls := BenchCalls + 1;
 110:
   BenchUut9.Mode := TRUE;
   BenchUut9.ForwardButton := FALSE;
   BenchUut9.ReverseButton := FALSE;
   BenchUut9.SensorFeed := FALSE;
   BenchUut9.SensorWash := FALSE;
   BenchUut9.SensorWeight := FALSE;
   BenchUut9.SensorFiring := TRUE;
   BenchUut9.SensorOutput := FALSE;
   BenchUut9.washComplete := FALSE;
   BenchUut9.weightComplete := FALSE;
   BenchUut9.weight := REAL#150.0;
   BenchUut9.firingComplete := TRUE;
   TraceIn_Mode[110] := BenchUut9.Mode;
   TraceIn_ForwardButton[110] := BenchUut9.ForwardButton;
   TraceIn_ReverseButton[110] := BenchUut9.ReverseButton;
   TraceIn_SensorFeed[110] := BenchUut9.SensorFeed;
   TraceIn_SensorWash[110] := BenchUut9.SensorWash;
   TraceIn_SensorWeight[110] := BenchUut9.SensorWeight;
   TraceIn_SensorFiring[110] := BenchUut9.SensorFiring;
   TraceIn_SensorOutput[110] := BenchUut9.SensorOutput;
   TraceIn_washComplete[110] := BenchUut9.washComplete;
   TraceIn_weightComplete[110] := BenchUut9.weightComplete;
   TraceIn_weight[110] := BenchUut9.weight;
   TraceIn_firingComplete[110] := BenchUut9.firingComplete;
   BenchUut9();
   TraceOut_MotorForward[110] := BenchUut9.MotorForward;
   TraceOut_MotorReverse[110] := BenchUut9.MotorReverse;
   TraceOut_kick[110] := BenchUut9.kick;
   TraceOut_CompletionLight[110] := BenchUut9.CompletionLight;
   TraceOut_firingTemp[110] := BenchUut9.firingTemp;
   BenchCalls := BenchCalls + 1;
 111:
   BenchUut9.Mode := TRUE;
   BenchUut9.ForwardButton := FALSE;
   BenchUut9.ReverseButton := FALSE;
   BenchUut9.SensorFeed := FALSE;
   BenchUut9.SensorWash := FALSE;
   BenchUut9.SensorWeight := FALSE;
   BenchUut9.SensorFiring := FALSE;
   BenchUut9.SensorOutput := FALSE;
   BenchUut9.washComplete := FALSE;
   BenchUut9.weightComplete := FALSE;
   BenchUut9.weight := REAL#150.0;
   BenchUut9.firingComplete := FALSE;
   TraceIn_Mode[111] := BenchUut9.Mode;
   TraceIn_ForwardButton[111] := BenchUut9.ForwardButton;
   TraceIn_ReverseButton[111] := BenchUut9.ReverseButton;
   TraceIn_SensorFeed[111] := BenchUut9.SensorFeed;
   TraceIn_SensorWash[111] := BenchUut9.SensorWash;
   TraceIn_SensorWeight[111] := BenchUut9.SensorWeight;
   TraceIn_SensorFiring[111] := BenchUut9.SensorFiring;
   TraceIn_SensorOutput[111] := BenchUut9.SensorOutput;
   TraceIn_washComplete[111] := BenchUut9.washComplete;
   TraceIn_weightComplete[111] := BenchUut9.weightComplete;
   TraceIn_weight[111] := BenchUut9.weight;
   TraceIn_firingComplete[111] := BenchUut9.firingComplete;
   BenchUut9();
   TraceOut_MotorForward[111] := BenchUut9.MotorForward;
   TraceOut_MotorReverse[111] := BenchUut9.MotorReverse;
   TraceOut_kick[111] := BenchUut9.kick;
   TraceOut_CompletionLight[111] := BenchUut9.CompletionLight;
   TraceOut_firingTemp[111] := BenchUut9.firingTemp;
   BenchCalls := BenchCalls + 1;
 112:
   BenchUut9.Mode := TRUE;
   BenchUut9.ForwardButton := FALSE;
   BenchUut9.ReverseButton := FALSE;
   BenchUut9.SensorFeed := FALSE;
   BenchUut9.SensorWash := FALSE;
   BenchUut9.SensorWeight := FALSE;
   BenchUut9.SensorFiring := FALSE;
   BenchUut9.SensorOutput := FALSE;
   BenchUut9.washComplete := FALSE;
   BenchUut9.weightComplete := FALSE;
   BenchUut9.weight := REAL#150.0;
   BenchUut9.firingComplete := FALSE;
   TraceIn_Mode[112] := BenchUut9.Mode;
   TraceIn_ForwardButton[112] := BenchUut9.ForwardButton;
   TraceIn_ReverseButton[112] := BenchUut9.ReverseButton;
   TraceIn_SensorFeed[112] := BenchUut9.SensorFeed;
   TraceIn_SensorWash[112] := BenchUut9.SensorWash;
   TraceIn_SensorWeight[112] := BenchUut9.SensorWeight;
   TraceIn_SensorFiring[112] := BenchUut9.SensorFiring;
   TraceIn_SensorOutput[112] := BenchUut9.SensorOutput;
   TraceIn_washComplete[112] := BenchUut9.washComplete;
   TraceIn_weightComplete[112] := BenchUut9.weightComplete;
   TraceIn_weight[112] := BenchUut9.weight;
   TraceIn_firingComplete[112] := BenchUut9.firingComplete;
   BenchUut9();
   TraceOut_MotorForward[112] := BenchUut9.MotorForward;
   TraceOut_MotorReverse[112] := BenchUut9.MotorReverse;
   TraceOut_kick[112] := BenchUut9.kick;
   TraceOut_CompletionLight[112] := BenchUut9.CompletionLight;
   TraceOut_firingTemp[112] := BenchUut9.firingTemp;
   BenchCalls := BenchCalls + 1;
 113:
   BenchUut9.Mode := TRUE;
   BenchUut9.ForwardButton := FALSE;
   BenchUut9.ReverseButton := FALSE;
   BenchUut9.SensorFeed := FALSE;
   BenchUut9.SensorWash := FALSE;
   BenchUut9.SensorWeight := FALSE;
   BenchUut9.SensorFiring := FALSE;
   BenchUut9.SensorOutput := FALSE;
   BenchUut9.washComplete := FALSE;
   BenchUut9.weightComplete := FALSE;
   BenchUut9.weight := REAL#150.0;
   BenchUut9.firingComplete := FALSE;
   TraceIn_Mode[113] := BenchUut9.Mode;
   TraceIn_ForwardButton[113] := BenchUut9.ForwardButton;
   TraceIn_ReverseButton[113] := BenchUut9.ReverseButton;
   TraceIn_SensorFeed[113] := BenchUut9.SensorFeed;
   TraceIn_SensorWash[113] := BenchUut9.SensorWash;
   TraceIn_SensorWeight[113] := BenchUut9.SensorWeight;
   TraceIn_SensorFiring[113] := BenchUut9.SensorFiring;
   TraceIn_SensorOutput[113] := BenchUut9.SensorOutput;
   TraceIn_washComplete[113] := BenchUut9.washComplete;
   TraceIn_weightComplete[113] := BenchUut9.weightComplete;
   TraceIn_weight[113] := BenchUut9.weight;
   TraceIn_firingComplete[113] := BenchUut9.firingComplete;
   BenchUut9();
   TraceOut_MotorForward[113] := BenchUut9.MotorForward;
   TraceOut_MotorReverse[113] := BenchUut9.MotorReverse;
   TraceOut_kick[113] := BenchUut9.kick;
   TraceOut_CompletionLight[113] := BenchUut9.CompletionLight;
   TraceOut_firingTemp[113] := BenchUut9.firingTemp;
   BenchCalls := BenchCalls + 1;
 114:
   BenchUut9.Mode := TRUE;
   BenchUut9.ForwardButton := FALSE;
   BenchUut9.ReverseButton := FALSE;
   BenchUut9.SensorFeed := FALSE;
   BenchUut9.SensorWash := FALSE;
   BenchUut9.SensorWeight := FALSE;
   BenchUut9.SensorFiring := FALSE;
   BenchUut9.SensorOutput := TRUE;
   BenchUut9.washComplete := FALSE;
   BenchUut9.weightComplete := FALSE;
   BenchUut9.weight := REAL#150.0;
   BenchUut9.firingComplete := FALSE;
   TraceIn_Mode[114] := BenchUut9.Mode;
   TraceIn_ForwardButton[114] := BenchUut9.ForwardButton;
   TraceIn_ReverseButton[114] := BenchUut9.ReverseButton;
   TraceIn_SensorFeed[114] := BenchUut9.SensorFeed;
   TraceIn_SensorWash[114] := BenchUut9.SensorWash;
   TraceIn_SensorWeight[114] := BenchUut9.SensorWeight;
   TraceIn_SensorFiring[114] := BenchUut9.SensorFiring;
   TraceIn_SensorOutput[114] := BenchUut9.SensorOutput;
   TraceIn_washComplete[114] := BenchUut9.washComplete;
   TraceIn_weightComplete[114] := BenchUut9.weightComplete;
   TraceIn_weight[114] := BenchUut9.weight;
   TraceIn_firingComplete[114] := BenchUut9.firingComplete;
   BenchUut9();
   TraceOut_MotorForward[114] := BenchUut9.MotorForward;
   TraceOut_MotorReverse[114] := BenchUut9.MotorReverse;
   TraceOut_kick[114] := BenchUut9.kick;
   TraceOut_CompletionLight[114] := BenchUut9.CompletionLight;
   TraceOut_firingTemp[114] := BenchUut9.firingTemp;
   BenchCalls := BenchCalls + 1;
 115:
   BenchUut9.Mode := TRUE;
   BenchUut9.ForwardButton := FALSE;
   BenchUut9.ReverseButton := FALSE;
   BenchUut9.SensorFeed := FALSE;
   BenchUut9.SensorWash := FALSE;
   BenchUut9.SensorWeight := FALSE;
   BenchUut9.SensorFiring := FALSE;
   BenchUut9.SensorOutput := TRUE;
   BenchUut9.washComplete := FALSE;
   BenchUut9.weightComplete := FALSE;
   BenchUut9.weight := REAL#150.0;
   BenchUut9.firingComplete := FALSE;
   TraceIn_Mode[115] := BenchUut9.Mode;
   TraceIn_ForwardButton[115] := BenchUut9.ForwardButton;
   TraceIn_ReverseButton[115] := BenchUut9.ReverseButton;
   TraceIn_SensorFeed[115] := BenchUut9.SensorFeed;
   TraceIn_SensorWash[115] := BenchUut9.SensorWash;
   TraceIn_SensorWeight[115] := BenchUut9.SensorWeight;
   TraceIn_SensorFiring[115] := BenchUut9.SensorFiring;
   TraceIn_SensorOutput[115] := BenchUut9.SensorOutput;
   TraceIn_washComplete[115] := BenchUut9.washComplete;
   TraceIn_weightComplete[115] := BenchUut9.weightComplete;
   TraceIn_weight[115] := BenchUut9.weight;
   TraceIn_firingComplete[115] := BenchUut9.firingComplete;
   BenchUut9();
   TraceOut_MotorForward[115] := BenchUut9.MotorForward;
   TraceOut_MotorReverse[115] := BenchUut9.MotorReverse;
   TraceOut_kick[115] := BenchUut9.kick;
   TraceOut_CompletionLight[115] := BenchUut9.CompletionLight;
   TraceOut_firingTemp[115] := BenchUut9.firingTemp;
   BenchCalls := BenchCalls + 1;
 116:
   BenchUut9.Mode := TRUE;
   BenchUut9.ForwardButton := FALSE;
   BenchUut9.ReverseButton := FALSE;
   BenchUut9.SensorFeed := FALSE;
   BenchUut9.SensorWash := FALSE;
   BenchUut9.SensorWeight := FALSE;
   BenchUut9.SensorFiring := FALSE;
   BenchUut9.SensorOutput := TRUE;
   BenchUut9.washComplete := FALSE;
   BenchUut9.weightComplete := FALSE;
   BenchUut9.weight := REAL#150.0;
   BenchUut9.firingComplete := FALSE;
   TraceIn_Mode[116] := BenchUut9.Mode;
   TraceIn_ForwardButton[116] := BenchUut9.ForwardButton;
   TraceIn_ReverseButton[116] := BenchUut9.ReverseButton;
   TraceIn_SensorFeed[116] := BenchUut9.SensorFeed;
   TraceIn_SensorWash[116] := BenchUut9.SensorWash;
   TraceIn_SensorWeight[116] := BenchUut9.SensorWeight;
   TraceIn_SensorFiring[116] := BenchUut9.SensorFiring;
   TraceIn_SensorOutput[116] := BenchUut9.SensorOutput;
   TraceIn_washComplete[116] := BenchUut9.washComplete;
   TraceIn_weightComplete[116] := BenchUut9.weightComplete;
   TraceIn_weight[116] := BenchUut9.weight;
   TraceIn_firingComplete[116] := BenchUut9.firingComplete;
   BenchUut9();
   TraceOut_MotorForward[116] := BenchUut9.MotorForward;
   TraceOut_MotorReverse[116] := BenchUut9.MotorReverse;
   TraceOut_kick[116] := BenchUut9.kick;
   TraceOut_CompletionLight[116] := BenchUut9.CompletionLight;
   TraceOut_firingTemp[116] := BenchUut9.firingTemp;
   BenchCalls := BenchCalls + 1;
 117:
   BenchUut9.Mode := TRUE;
   BenchUut9.ForwardButton := FALSE;
   BenchUut9.ReverseButton := FALSE;
   BenchUut9.SensorFeed := FALSE;
   BenchUut9.SensorWash := FALSE;
   BenchUut9.SensorWeight := FALSE;
   BenchUut9.SensorFiring := FALSE;
   BenchUut9.SensorOutput := FALSE;
   BenchUut9.washComplete := FALSE;
   BenchUut9.weightComplete := FALSE;
   BenchUut9.weight := REAL#150.0;
   BenchUut9.firingComplete := FALSE;
   TraceIn_Mode[117] := BenchUut9.Mode;
   TraceIn_ForwardButton[117] := BenchUut9.ForwardButton;
   TraceIn_ReverseButton[117] := BenchUut9.ReverseButton;
   TraceIn_SensorFeed[117] := BenchUut9.SensorFeed;
   TraceIn_SensorWash[117] := BenchUut9.SensorWash;
   TraceIn_SensorWeight[117] := BenchUut9.SensorWeight;
   TraceIn_SensorFiring[117] := BenchUut9.SensorFiring;
   TraceIn_SensorOutput[117] := BenchUut9.SensorOutput;
   TraceIn_washComplete[117] := BenchUut9.washComplete;
   TraceIn_weightComplete[117] := BenchUut9.weightComplete;
   TraceIn_weight[117] := BenchUut9.weight;
   TraceIn_firingComplete[117] := BenchUut9.firingComplete;
   BenchUut9();
   TraceOut_MotorForward[117] := BenchUut9.MotorForward;
   TraceOut_MotorReverse[117] := BenchUut9.MotorReverse;
   TraceOut_kick[117] := BenchUut9.kick;
   TraceOut_CompletionLight[117] := BenchUut9.CompletionLight;
   TraceOut_firingTemp[117] := BenchUut9.firingTemp;
   BenchCalls := BenchCalls + 1;
 118:
   BenchUut9.Mode := TRUE;
   BenchUut9.ForwardButton := FALSE;
   BenchUut9.ReverseButton := FALSE;
   BenchUut9.SensorFeed := TRUE;
   BenchUut9.SensorWash := FALSE;
   BenchUut9.SensorWeight := FALSE;
   BenchUut9.SensorFiring := FALSE;
   BenchUut9.SensorOutput := FALSE;
   BenchUut9.washComplete := FALSE;
   BenchUut9.weightComplete := FALSE;
   BenchUut9.weight := REAL#150.0;
   BenchUut9.firingComplete := FALSE;
   TraceIn_Mode[118] := BenchUut9.Mode;
   TraceIn_ForwardButton[118] := BenchUut9.ForwardButton;
   TraceIn_ReverseButton[118] := BenchUut9.ReverseButton;
   TraceIn_SensorFeed[118] := BenchUut9.SensorFeed;
   TraceIn_SensorWash[118] := BenchUut9.SensorWash;
   TraceIn_SensorWeight[118] := BenchUut9.SensorWeight;
   TraceIn_SensorFiring[118] := BenchUut9.SensorFiring;
   TraceIn_SensorOutput[118] := BenchUut9.SensorOutput;
   TraceIn_washComplete[118] := BenchUut9.washComplete;
   TraceIn_weightComplete[118] := BenchUut9.weightComplete;
   TraceIn_weight[118] := BenchUut9.weight;
   TraceIn_firingComplete[118] := BenchUut9.firingComplete;
   BenchUut9();
   TraceOut_MotorForward[118] := BenchUut9.MotorForward;
   TraceOut_MotorReverse[118] := BenchUut9.MotorReverse;
   TraceOut_kick[118] := BenchUut9.kick;
   TraceOut_CompletionLight[118] := BenchUut9.CompletionLight;
   TraceOut_firingTemp[118] := BenchUut9.firingTemp;
   BenchCalls := BenchCalls + 1;
 119:
   BenchUut9.Mode := TRUE;
   BenchUut9.ForwardButton := FALSE;
   BenchUut9.ReverseButton := FALSE;
   BenchUut9.SensorFeed := FALSE;
   BenchUut9.SensorWash := FALSE;
   BenchUut9.SensorWeight := FALSE;
   BenchUut9.SensorFiring := FALSE;
   BenchUut9.SensorOutput := FALSE;
   BenchUut9.washComplete := FALSE;
   BenchUut9.weightComplete := FALSE;
   BenchUut9.weight := REAL#150.0;
   BenchUut9.firingComplete := FALSE;
   TraceIn_Mode[119] := BenchUut9.Mode;
   TraceIn_ForwardButton[119] := BenchUut9.ForwardButton;
   TraceIn_ReverseButton[119] := BenchUut9.ReverseButton;
   TraceIn_SensorFeed[119] := BenchUut9.SensorFeed;
   TraceIn_SensorWash[119] := BenchUut9.SensorWash;
   TraceIn_SensorWeight[119] := BenchUut9.SensorWeight;
   TraceIn_SensorFiring[119] := BenchUut9.SensorFiring;
   TraceIn_SensorOutput[119] := BenchUut9.SensorOutput;
   TraceIn_washComplete[119] := BenchUut9.washComplete;
   TraceIn_weightComplete[119] := BenchUut9.weightComplete;
   TraceIn_weight[119] := BenchUut9.weight;
   TraceIn_firingComplete[119] := BenchUut9.firingComplete;
   BenchUut9();
   TraceOut_MotorForward[119] := BenchUut9.MotorForward;
   TraceOut_MotorReverse[119] := BenchUut9.MotorReverse;
   TraceOut_kick[119] := BenchUut9.kick;
   TraceOut_CompletionLight[119] := BenchUut9.CompletionLight;
   TraceOut_firingTemp[119] := BenchUut9.firingTemp;
   BenchCalls := BenchCalls + 1;
 120:
   BenchUut9.Mode := TRUE;
   BenchUut9.ForwardButton := FALSE;
   BenchUut9.ReverseButton := FALSE;
   BenchUut9.SensorFeed := FALSE;
   BenchUut9.SensorWash := FALSE;
   BenchUut9.SensorWeight := FALSE;
   BenchUut9.SensorFiring := FALSE;
   BenchUut9.SensorOutput := FALSE;
   BenchUut9.washComplete := FALSE;
   BenchUut9.weightComplete := FALSE;
   BenchUut9.weight := REAL#150.0;
   BenchUut9.firingComplete := FALSE;
   TraceIn_Mode[120] := BenchUut9.Mode;
   TraceIn_ForwardButton[120] := BenchUut9.ForwardButton;
   TraceIn_ReverseButton[120] := BenchUut9.ReverseButton;
   TraceIn_SensorFeed[120] := BenchUut9.SensorFeed;
   TraceIn_SensorWash[120] := BenchUut9.SensorWash;
   TraceIn_SensorWeight[120] := BenchUut9.SensorWeight;
   TraceIn_SensorFiring[120] := BenchUut9.SensorFiring;
   TraceIn_SensorOutput[120] := BenchUut9.SensorOutput;
   TraceIn_washComplete[120] := BenchUut9.washComplete;
   TraceIn_weightComplete[120] := BenchUut9.weightComplete;
   TraceIn_weight[120] := BenchUut9.weight;
   TraceIn_firingComplete[120] := BenchUut9.firingComplete;
   BenchUut9();
   TraceOut_MotorForward[120] := BenchUut9.MotorForward;
   TraceOut_MotorReverse[120] := BenchUut9.MotorReverse;
   TraceOut_kick[120] := BenchUut9.kick;
   TraceOut_CompletionLight[120] := BenchUut9.CompletionLight;
   TraceOut_firingTemp[120] := BenchUut9.firingTemp;
   BenchCalls := BenchCalls + 1;
 121:
   BenchUut9.Mode := TRUE;
   BenchUut9.ForwardButton := FALSE;
   BenchUut9.ReverseButton := FALSE;
   BenchUut9.SensorFeed := FALSE;
   BenchUut9.SensorWash := FALSE;
   BenchUut9.SensorWeight := FALSE;
   BenchUut9.SensorFiring := FALSE;
   BenchUut9.SensorOutput := FALSE;
   BenchUut9.washComplete := FALSE;
   BenchUut9.weightComplete := FALSE;
   BenchUut9.weight := REAL#150.0;
   BenchUut9.firingComplete := FALSE;
   TraceIn_Mode[121] := BenchUut9.Mode;
   TraceIn_ForwardButton[121] := BenchUut9.ForwardButton;
   TraceIn_ReverseButton[121] := BenchUut9.ReverseButton;
   TraceIn_SensorFeed[121] := BenchUut9.SensorFeed;
   TraceIn_SensorWash[121] := BenchUut9.SensorWash;
   TraceIn_SensorWeight[121] := BenchUut9.SensorWeight;
   TraceIn_SensorFiring[121] := BenchUut9.SensorFiring;
   TraceIn_SensorOutput[121] := BenchUut9.SensorOutput;
   TraceIn_washComplete[121] := BenchUut9.washComplete;
   TraceIn_weightComplete[121] := BenchUut9.weightComplete;
   TraceIn_weight[121] := BenchUut9.weight;
   TraceIn_firingComplete[121] := BenchUut9.firingComplete;
   BenchUut9();
   TraceOut_MotorForward[121] := BenchUut9.MotorForward;
   TraceOut_MotorReverse[121] := BenchUut9.MotorReverse;
   TraceOut_kick[121] := BenchUut9.kick;
   TraceOut_CompletionLight[121] := BenchUut9.CompletionLight;
   TraceOut_firingTemp[121] := BenchUut9.firingTemp;
   BenchCalls := BenchCalls + 1;
 122:
   BenchUut9.Mode := TRUE;
   BenchUut9.ForwardButton := FALSE;
   BenchUut9.ReverseButton := FALSE;
   BenchUut9.SensorFeed := FALSE;
   BenchUut9.SensorWash := TRUE;
   BenchUut9.SensorWeight := FALSE;
   BenchUut9.SensorFiring := FALSE;
   BenchUut9.SensorOutput := FALSE;
   BenchUut9.washComplete := FALSE;
   BenchUut9.weightComplete := FALSE;
   BenchUut9.weight := REAL#150.0;
   BenchUut9.firingComplete := FALSE;
   TraceIn_Mode[122] := BenchUut9.Mode;
   TraceIn_ForwardButton[122] := BenchUut9.ForwardButton;
   TraceIn_ReverseButton[122] := BenchUut9.ReverseButton;
   TraceIn_SensorFeed[122] := BenchUut9.SensorFeed;
   TraceIn_SensorWash[122] := BenchUut9.SensorWash;
   TraceIn_SensorWeight[122] := BenchUut9.SensorWeight;
   TraceIn_SensorFiring[122] := BenchUut9.SensorFiring;
   TraceIn_SensorOutput[122] := BenchUut9.SensorOutput;
   TraceIn_washComplete[122] := BenchUut9.washComplete;
   TraceIn_weightComplete[122] := BenchUut9.weightComplete;
   TraceIn_weight[122] := BenchUut9.weight;
   TraceIn_firingComplete[122] := BenchUut9.firingComplete;
   BenchUut9();
   TraceOut_MotorForward[122] := BenchUut9.MotorForward;
   TraceOut_MotorReverse[122] := BenchUut9.MotorReverse;
   TraceOut_kick[122] := BenchUut9.kick;
   TraceOut_CompletionLight[122] := BenchUut9.CompletionLight;
   TraceOut_firingTemp[122] := BenchUut9.firingTemp;
   BenchCalls := BenchCalls + 1;
 123:
   BenchUut9.Mode := TRUE;
   BenchUut9.ForwardButton := FALSE;
   BenchUut9.ReverseButton := FALSE;
   BenchUut9.SensorFeed := FALSE;
   BenchUut9.SensorWash := TRUE;
   BenchUut9.SensorWeight := FALSE;
   BenchUut9.SensorFiring := FALSE;
   BenchUut9.SensorOutput := FALSE;
   BenchUut9.washComplete := FALSE;
   BenchUut9.weightComplete := FALSE;
   BenchUut9.weight := REAL#150.0;
   BenchUut9.firingComplete := FALSE;
   TraceIn_Mode[123] := BenchUut9.Mode;
   TraceIn_ForwardButton[123] := BenchUut9.ForwardButton;
   TraceIn_ReverseButton[123] := BenchUut9.ReverseButton;
   TraceIn_SensorFeed[123] := BenchUut9.SensorFeed;
   TraceIn_SensorWash[123] := BenchUut9.SensorWash;
   TraceIn_SensorWeight[123] := BenchUut9.SensorWeight;
   TraceIn_SensorFiring[123] := BenchUut9.SensorFiring;
   TraceIn_SensorOutput[123] := BenchUut9.SensorOutput;
   TraceIn_washComplete[123] := BenchUut9.washComplete;
   TraceIn_weightComplete[123] := BenchUut9.weightComplete;
   TraceIn_weight[123] := BenchUut9.weight;
   TraceIn_firingComplete[123] := BenchUut9.firingComplete;
   BenchUut9();
   TraceOut_MotorForward[123] := BenchUut9.MotorForward;
   TraceOut_MotorReverse[123] := BenchUut9.MotorReverse;
   TraceOut_kick[123] := BenchUut9.kick;
   TraceOut_CompletionLight[123] := BenchUut9.CompletionLight;
   TraceOut_firingTemp[123] := BenchUut9.firingTemp;
   BenchCalls := BenchCalls + 1;
 124:
   BenchUut9.Mode := TRUE;
   BenchUut9.ForwardButton := FALSE;
   BenchUut9.ReverseButton := FALSE;
   BenchUut9.SensorFeed := FALSE;
   BenchUut9.SensorWash := TRUE;
   BenchUut9.SensorWeight := FALSE;
   BenchUut9.SensorFiring := FALSE;
   BenchUut9.SensorOutput := FALSE;
   BenchUut9.washComplete := FALSE;
   BenchUut9.weightComplete := FALSE;
   BenchUut9.weight := REAL#150.0;
   BenchUut9.firingComplete := FALSE;
   TraceIn_Mode[124] := BenchUut9.Mode;
   TraceIn_ForwardButton[124] := BenchUut9.ForwardButton;
   TraceIn_ReverseButton[124] := BenchUut9.ReverseButton;
   TraceIn_SensorFeed[124] := BenchUut9.SensorFeed;
   TraceIn_SensorWash[124] := BenchUut9.SensorWash;
   TraceIn_SensorWeight[124] := BenchUut9.SensorWeight;
   TraceIn_SensorFiring[124] := BenchUut9.SensorFiring;
   TraceIn_SensorOutput[124] := BenchUut9.SensorOutput;
   TraceIn_washComplete[124] := BenchUut9.washComplete;
   TraceIn_weightComplete[124] := BenchUut9.weightComplete;
   TraceIn_weight[124] := BenchUut9.weight;
   TraceIn_firingComplete[124] := BenchUut9.firingComplete;
   BenchUut9();
   TraceOut_MotorForward[124] := BenchUut9.MotorForward;
   TraceOut_MotorReverse[124] := BenchUut9.MotorReverse;
   TraceOut_kick[124] := BenchUut9.kick;
   TraceOut_CompletionLight[124] := BenchUut9.CompletionLight;
   TraceOut_firingTemp[124] := BenchUut9.firingTemp;
   BenchCalls := BenchCalls + 1;
 125:
   BenchUut9.Mode := TRUE;
   BenchUut9.ForwardButton := FALSE;
   BenchUut9.ReverseButton := FALSE;
   BenchUut9.SensorFeed := FALSE;
   BenchUut9.SensorWash := TRUE;
   BenchUut9.SensorWeight := FALSE;
   BenchUut9.SensorFiring := FALSE;
   BenchUut9.SensorOutput := FALSE;
   BenchUut9.washComplete := TRUE;
   BenchUut9.weightComplete := FALSE;
   BenchUut9.weight := REAL#150.0;
   BenchUut9.firingComplete := FALSE;
   TraceIn_Mode[125] := BenchUut9.Mode;
   TraceIn_ForwardButton[125] := BenchUut9.ForwardButton;
   TraceIn_ReverseButton[125] := BenchUut9.ReverseButton;
   TraceIn_SensorFeed[125] := BenchUut9.SensorFeed;
   TraceIn_SensorWash[125] := BenchUut9.SensorWash;
   TraceIn_SensorWeight[125] := BenchUut9.SensorWeight;
   TraceIn_SensorFiring[125] := BenchUut9.SensorFiring;
   TraceIn_SensorOutput[125] := BenchUut9.SensorOutput;
   TraceIn_washComplete[125] := BenchUut9.washComplete;
   TraceIn_weightComplete[125] := BenchUut9.weightComplete;
   TraceIn_weight[125] := BenchUut9.weight;
   TraceIn_firingComplete[125] := BenchUut9.firingComplete;
   BenchUut9();
   TraceOut_MotorForward[125] := BenchUut9.MotorForward;
   TraceOut_MotorReverse[125] := BenchUut9.MotorReverse;
   TraceOut_kick[125] := BenchUut9.kick;
   TraceOut_CompletionLight[125] := BenchUut9.CompletionLight;
   TraceOut_firingTemp[125] := BenchUut9.firingTemp;
   BenchCalls := BenchCalls + 1;
 126:
   BenchUut9.Mode := TRUE;
   BenchUut9.ForwardButton := FALSE;
   BenchUut9.ReverseButton := FALSE;
   BenchUut9.SensorFeed := FALSE;
   BenchUut9.SensorWash := FALSE;
   BenchUut9.SensorWeight := FALSE;
   BenchUut9.SensorFiring := FALSE;
   BenchUut9.SensorOutput := FALSE;
   BenchUut9.washComplete := FALSE;
   BenchUut9.weightComplete := FALSE;
   BenchUut9.weight := REAL#150.0;
   BenchUut9.firingComplete := FALSE;
   TraceIn_Mode[126] := BenchUut9.Mode;
   TraceIn_ForwardButton[126] := BenchUut9.ForwardButton;
   TraceIn_ReverseButton[126] := BenchUut9.ReverseButton;
   TraceIn_SensorFeed[126] := BenchUut9.SensorFeed;
   TraceIn_SensorWash[126] := BenchUut9.SensorWash;
   TraceIn_SensorWeight[126] := BenchUut9.SensorWeight;
   TraceIn_SensorFiring[126] := BenchUut9.SensorFiring;
   TraceIn_SensorOutput[126] := BenchUut9.SensorOutput;
   TraceIn_washComplete[126] := BenchUut9.washComplete;
   TraceIn_weightComplete[126] := BenchUut9.weightComplete;
   TraceIn_weight[126] := BenchUut9.weight;
   TraceIn_firingComplete[126] := BenchUut9.firingComplete;
   BenchUut9();
   TraceOut_MotorForward[126] := BenchUut9.MotorForward;
   TraceOut_MotorReverse[126] := BenchUut9.MotorReverse;
   TraceOut_kick[126] := BenchUut9.kick;
   TraceOut_CompletionLight[126] := BenchUut9.CompletionLight;
   TraceOut_firingTemp[126] := BenchUut9.firingTemp;
   BenchCalls := BenchCalls + 1;
 127:
   BenchUut9.Mode := TRUE;
   BenchUut9.ForwardButton := FALSE;
   BenchUut9.ReverseButton := FALSE;
   BenchUut9.SensorFeed := FALSE;
   BenchUut9.SensorWash := FALSE;
   BenchUut9.SensorWeight := FALSE;
   BenchUut9.SensorFiring := FALSE;
   BenchUut9.SensorOutput := FALSE;
   BenchUut9.washComplete := FALSE;
   BenchUut9.weightComplete := FALSE;
   BenchUut9.weight := REAL#150.0;
   BenchUut9.firingComplete := FALSE;
   TraceIn_Mode[127] := BenchUut9.Mode;
   TraceIn_ForwardButton[127] := BenchUut9.ForwardButton;
   TraceIn_ReverseButton[127] := BenchUut9.ReverseButton;
   TraceIn_SensorFeed[127] := BenchUut9.SensorFeed;
   TraceIn_SensorWash[127] := BenchUut9.SensorWash;
   TraceIn_SensorWeight[127] := BenchUut9.SensorWeight;
   TraceIn_SensorFiring[127] := BenchUut9.SensorFiring;
   TraceIn_SensorOutput[127] := BenchUut9.SensorOutput;
   TraceIn_washComplete[127] := BenchUut9.washComplete;
   TraceIn_weightComplete[127] := BenchUut9.weightComplete;
   TraceIn_weight[127] := BenchUut9.weight;
   TraceIn_firingComplete[127] := BenchUut9.firingComplete;
   BenchUut9();
   TraceOut_MotorForward[127] := BenchUut9.MotorForward;
   TraceOut_MotorReverse[127] := BenchUut9.MotorReverse;
   TraceOut_kick[127] := BenchUut9.kick;
   TraceOut_CompletionLight[127] := BenchUut9.CompletionLight;
   TraceOut_firingTemp[127] := BenchUut9.firingTemp;
   BenchCalls := BenchCalls + 1;
 128:
   BenchUut9.Mode := TRUE;
   BenchUut9.ForwardButton := FALSE;
   BenchUut9.ReverseButton := FALSE;
   BenchUut9.SensorFeed := FALSE;
   BenchUut9.SensorWash := FALSE;
   BenchUut9.SensorWeight := FALSE;
   BenchUut9.SensorFiring := FALSE;
   BenchUut9.SensorOutput := FALSE;
   BenchUut9.washComplete := FALSE;
   BenchUut9.weightComplete := FALSE;
   BenchUut9.weight := REAL#150.0;
   BenchUut9.firingComplete := FALSE;
   TraceIn_Mode[128] := BenchUut9.Mode;
   TraceIn_ForwardButton[128] := BenchUut9.ForwardButton;
   TraceIn_ReverseButton[128] := BenchUut9.ReverseButton;
   TraceIn_SensorFeed[128] := BenchUut9.SensorFeed;
   TraceIn_SensorWash[128] := BenchUut9.SensorWash;
   TraceIn_SensorWeight[128] := BenchUut9.SensorWeight;
   TraceIn_SensorFiring[128] := BenchUut9.SensorFiring;
   TraceIn_SensorOutput[128] := BenchUut9.SensorOutput;
   TraceIn_washComplete[128] := BenchUut9.washComplete;
   TraceIn_weightComplete[128] := BenchUut9.weightComplete;
   TraceIn_weight[128] := BenchUut9.weight;
   TraceIn_firingComplete[128] := BenchUut9.firingComplete;
   BenchUut9();
   TraceOut_MotorForward[128] := BenchUut9.MotorForward;
   TraceOut_MotorReverse[128] := BenchUut9.MotorReverse;
   TraceOut_kick[128] := BenchUut9.kick;
   TraceOut_CompletionLight[128] := BenchUut9.CompletionLight;
   TraceOut_firingTemp[128] := BenchUut9.firingTemp;
   BenchCalls := BenchCalls + 1;
 129:
   BenchUut9.Mode := TRUE;
   BenchUut9.ForwardButton := FALSE;
   BenchUut9.ReverseButton := FALSE;
   BenchUut9.SensorFeed := FALSE;
   BenchUut9.SensorWash := FALSE;
   BenchUut9.SensorWeight := TRUE;
   BenchUut9.SensorFiring := FALSE;
   BenchUut9.SensorOutput := FALSE;
   BenchUut9.washComplete := FALSE;
   BenchUut9.weightComplete := FALSE;
   BenchUut9.weight := REAL#150.0;
   BenchUut9.firingComplete := FALSE;
   TraceIn_Mode[129] := BenchUut9.Mode;
   TraceIn_ForwardButton[129] := BenchUut9.ForwardButton;
   TraceIn_ReverseButton[129] := BenchUut9.ReverseButton;
   TraceIn_SensorFeed[129] := BenchUut9.SensorFeed;
   TraceIn_SensorWash[129] := BenchUut9.SensorWash;
   TraceIn_SensorWeight[129] := BenchUut9.SensorWeight;
   TraceIn_SensorFiring[129] := BenchUut9.SensorFiring;
   TraceIn_SensorOutput[129] := BenchUut9.SensorOutput;
   TraceIn_washComplete[129] := BenchUut9.washComplete;
   TraceIn_weightComplete[129] := BenchUut9.weightComplete;
   TraceIn_weight[129] := BenchUut9.weight;
   TraceIn_firingComplete[129] := BenchUut9.firingComplete;
   BenchUut9();
   TraceOut_MotorForward[129] := BenchUut9.MotorForward;
   TraceOut_MotorReverse[129] := BenchUut9.MotorReverse;
   TraceOut_kick[129] := BenchUut9.kick;
   TraceOut_CompletionLight[129] := BenchUut9.CompletionLight;
   TraceOut_firingTemp[129] := BenchUut9.firingTemp;
   BenchCalls := BenchCalls + 1;
 130:
   BenchUut9.Mode := TRUE;
   BenchUut9.ForwardButton := FALSE;
   BenchUut9.ReverseButton := FALSE;
   BenchUut9.SensorFeed := FALSE;
   BenchUut9.SensorWash := FALSE;
   BenchUut9.SensorWeight := TRUE;
   BenchUut9.SensorFiring := FALSE;
   BenchUut9.SensorOutput := FALSE;
   BenchUut9.washComplete := FALSE;
   BenchUut9.weightComplete := FALSE;
   BenchUut9.weight := REAL#150.0;
   BenchUut9.firingComplete := FALSE;
   TraceIn_Mode[130] := BenchUut9.Mode;
   TraceIn_ForwardButton[130] := BenchUut9.ForwardButton;
   TraceIn_ReverseButton[130] := BenchUut9.ReverseButton;
   TraceIn_SensorFeed[130] := BenchUut9.SensorFeed;
   TraceIn_SensorWash[130] := BenchUut9.SensorWash;
   TraceIn_SensorWeight[130] := BenchUut9.SensorWeight;
   TraceIn_SensorFiring[130] := BenchUut9.SensorFiring;
   TraceIn_SensorOutput[130] := BenchUut9.SensorOutput;
   TraceIn_washComplete[130] := BenchUut9.washComplete;
   TraceIn_weightComplete[130] := BenchUut9.weightComplete;
   TraceIn_weight[130] := BenchUut9.weight;
   TraceIn_firingComplete[130] := BenchUut9.firingComplete;
   BenchUut9();
   TraceOut_MotorForward[130] := BenchUut9.MotorForward;
   TraceOut_MotorReverse[130] := BenchUut9.MotorReverse;
   TraceOut_kick[130] := BenchUut9.kick;
   TraceOut_CompletionLight[130] := BenchUut9.CompletionLight;
   TraceOut_firingTemp[130] := BenchUut9.firingTemp;
   BenchCalls := BenchCalls + 1;
 131:
   BenchUut9.Mode := TRUE;
   BenchUut9.ForwardButton := FALSE;
   BenchUut9.ReverseButton := FALSE;
   BenchUut9.SensorFeed := FALSE;
   BenchUut9.SensorWash := FALSE;
   BenchUut9.SensorWeight := TRUE;
   BenchUut9.SensorFiring := FALSE;
   BenchUut9.SensorOutput := FALSE;
   BenchUut9.washComplete := FALSE;
   BenchUut9.weightComplete := FALSE;
   BenchUut9.weight := REAL#150.0;
   BenchUut9.firingComplete := FALSE;
   TraceIn_Mode[131] := BenchUut9.Mode;
   TraceIn_ForwardButton[131] := BenchUut9.ForwardButton;
   TraceIn_ReverseButton[131] := BenchUut9.ReverseButton;
   TraceIn_SensorFeed[131] := BenchUut9.SensorFeed;
   TraceIn_SensorWash[131] := BenchUut9.SensorWash;
   TraceIn_SensorWeight[131] := BenchUut9.SensorWeight;
   TraceIn_SensorFiring[131] := BenchUut9.SensorFiring;
   TraceIn_SensorOutput[131] := BenchUut9.SensorOutput;
   TraceIn_washComplete[131] := BenchUut9.washComplete;
   TraceIn_weightComplete[131] := BenchUut9.weightComplete;
   TraceIn_weight[131] := BenchUut9.weight;
   TraceIn_firingComplete[131] := BenchUut9.firingComplete;
   BenchUut9();
   TraceOut_MotorForward[131] := BenchUut9.MotorForward;
   TraceOut_MotorReverse[131] := BenchUut9.MotorReverse;
   TraceOut_kick[131] := BenchUut9.kick;
   TraceOut_CompletionLight[131] := BenchUut9.CompletionLight;
   TraceOut_firingTemp[131] := BenchUut9.firingTemp;
   BenchCalls := BenchCalls + 1;
 132:
   BenchUut9.Mode := TRUE;
   BenchUut9.ForwardButton := FALSE;
   BenchUut9.ReverseButton := FALSE;
   BenchUut9.SensorFeed := FALSE;
   BenchUut9.SensorWash := FALSE;
   BenchUut9.SensorWeight := TRUE;
   BenchUut9.SensorFiring := FALSE;
   BenchUut9.SensorOutput := FALSE;
   BenchUut9.washComplete := FALSE;
   BenchUut9.weightComplete := TRUE;
   BenchUut9.weight := REAL#150.0;
   BenchUut9.firingComplete := FALSE;
   TraceIn_Mode[132] := BenchUut9.Mode;
   TraceIn_ForwardButton[132] := BenchUut9.ForwardButton;
   TraceIn_ReverseButton[132] := BenchUut9.ReverseButton;
   TraceIn_SensorFeed[132] := BenchUut9.SensorFeed;
   TraceIn_SensorWash[132] := BenchUut9.SensorWash;
   TraceIn_SensorWeight[132] := BenchUut9.SensorWeight;
   TraceIn_SensorFiring[132] := BenchUut9.SensorFiring;
   TraceIn_SensorOutput[132] := BenchUut9.SensorOutput;
   TraceIn_washComplete[132] := BenchUut9.washComplete;
   TraceIn_weightComplete[132] := BenchUut9.weightComplete;
   TraceIn_weight[132] := BenchUut9.weight;
   TraceIn_firingComplete[132] := BenchUut9.firingComplete;
   BenchUut9();
   TraceOut_MotorForward[132] := BenchUut9.MotorForward;
   TraceOut_MotorReverse[132] := BenchUut9.MotorReverse;
   TraceOut_kick[132] := BenchUut9.kick;
   TraceOut_CompletionLight[132] := BenchUut9.CompletionLight;
   TraceOut_firingTemp[132] := BenchUut9.firingTemp;
   BenchCalls := BenchCalls + 1;
 133:
   BenchUut9.Mode := TRUE;
   BenchUut9.ForwardButton := FALSE;
   BenchUut9.ReverseButton := FALSE;
   BenchUut9.SensorFeed := FALSE;
   BenchUut9.SensorWash := FALSE;
   BenchUut9.SensorWeight := FALSE;
   BenchUut9.SensorFiring := FALSE;
   BenchUut9.SensorOutput := FALSE;
   BenchUut9.washComplete := FALSE;
   BenchUut9.weightComplete := FALSE;
   BenchUut9.weight := REAL#150.0;
   BenchUut9.firingComplete := FALSE;
   TraceIn_Mode[133] := BenchUut9.Mode;
   TraceIn_ForwardButton[133] := BenchUut9.ForwardButton;
   TraceIn_ReverseButton[133] := BenchUut9.ReverseButton;
   TraceIn_SensorFeed[133] := BenchUut9.SensorFeed;
   TraceIn_SensorWash[133] := BenchUut9.SensorWash;
   TraceIn_SensorWeight[133] := BenchUut9.SensorWeight;
   TraceIn_SensorFiring[133] := BenchUut9.SensorFiring;
   TraceIn_SensorOutput[133] := BenchUut9.SensorOutput;
   TraceIn_washComplete[133] := BenchUut9.washComplete;
   TraceIn_weightComplete[133] := BenchUut9.weightComplete;
   TraceIn_weight[133] := BenchUut9.weight;
   TraceIn_firingComplete[133] := BenchUut9.firingComplete;
   BenchUut9();
   TraceOut_MotorForward[133] := BenchUut9.MotorForward;
   TraceOut_MotorReverse[133] := BenchUut9.MotorReverse;
   TraceOut_kick[133] := BenchUut9.kick;
   TraceOut_CompletionLight[133] := BenchUut9.CompletionLight;
   TraceOut_firingTemp[133] := BenchUut9.firingTemp;
   BenchCalls := BenchCalls + 1;
 134:
   BenchUut9.Mode := TRUE;
   BenchUut9.ForwardButton := FALSE;
   BenchUut9.ReverseButton := FALSE;
   BenchUut9.SensorFeed := FALSE;
   BenchUut9.SensorWash := FALSE;
   BenchUut9.SensorWeight := FALSE;
   BenchUut9.SensorFiring := FALSE;
   BenchUut9.SensorOutput := FALSE;
   BenchUut9.washComplete := FALSE;
   BenchUut9.weightComplete := FALSE;
   BenchUut9.weight := REAL#150.0;
   BenchUut9.firingComplete := FALSE;
   TraceIn_Mode[134] := BenchUut9.Mode;
   TraceIn_ForwardButton[134] := BenchUut9.ForwardButton;
   TraceIn_ReverseButton[134] := BenchUut9.ReverseButton;
   TraceIn_SensorFeed[134] := BenchUut9.SensorFeed;
   TraceIn_SensorWash[134] := BenchUut9.SensorWash;
   TraceIn_SensorWeight[134] := BenchUut9.SensorWeight;
   TraceIn_SensorFiring[134] := BenchUut9.SensorFiring;
   TraceIn_SensorOutput[134] := BenchUut9.SensorOutput;
   TraceIn_washComplete[134] := BenchUut9.washComplete;
   TraceIn_weightComplete[134] := BenchUut9.weightComplete;
   TraceIn_weight[134] := BenchUut9.weight;
   TraceIn_firingComplete[134] := BenchUut9.firingComplete;
   BenchUut9();
   TraceOut_MotorForward[134] := BenchUut9.MotorForward;
   TraceOut_MotorReverse[134] := BenchUut9.MotorReverse;
   TraceOut_kick[134] := BenchUut9.kick;
   TraceOut_CompletionLight[134] := BenchUut9.CompletionLight;
   TraceOut_firingTemp[134] := BenchUut9.firingTemp;
   BenchCalls := BenchCalls + 1;
 135:
   BenchUut9.Mode := TRUE;
   BenchUut9.ForwardButton := FALSE;
   BenchUut9.ReverseButton := FALSE;
   BenchUut9.SensorFeed := FALSE;
   BenchUut9.SensorWash := FALSE;
   BenchUut9.SensorWeight := FALSE;
   BenchUut9.SensorFiring := FALSE;
   BenchUut9.SensorOutput := FALSE;
   BenchUut9.washComplete := FALSE;
   BenchUut9.weightComplete := FALSE;
   BenchUut9.weight := REAL#150.0;
   BenchUut9.firingComplete := FALSE;
   TraceIn_Mode[135] := BenchUut9.Mode;
   TraceIn_ForwardButton[135] := BenchUut9.ForwardButton;
   TraceIn_ReverseButton[135] := BenchUut9.ReverseButton;
   TraceIn_SensorFeed[135] := BenchUut9.SensorFeed;
   TraceIn_SensorWash[135] := BenchUut9.SensorWash;
   TraceIn_SensorWeight[135] := BenchUut9.SensorWeight;
   TraceIn_SensorFiring[135] := BenchUut9.SensorFiring;
   TraceIn_SensorOutput[135] := BenchUut9.SensorOutput;
   TraceIn_washComplete[135] := BenchUut9.washComplete;
   TraceIn_weightComplete[135] := BenchUut9.weightComplete;
   TraceIn_weight[135] := BenchUut9.weight;
   TraceIn_firingComplete[135] := BenchUut9.firingComplete;
   BenchUut9();
   TraceOut_MotorForward[135] := BenchUut9.MotorForward;
   TraceOut_MotorReverse[135] := BenchUut9.MotorReverse;
   TraceOut_kick[135] := BenchUut9.kick;
   TraceOut_CompletionLight[135] := BenchUut9.CompletionLight;
   TraceOut_firingTemp[135] := BenchUut9.firingTemp;
   BenchCalls := BenchCalls + 1;
 136:
   BenchUut9.Mode := TRUE;
   BenchUut9.ForwardButton := FALSE;
   BenchUut9.ReverseButton := FALSE;
   BenchUut9.SensorFeed := FALSE;
   BenchUut9.SensorWash := FALSE;
   BenchUut9.SensorWeight := FALSE;
   BenchUut9.SensorFiring := TRUE;
   BenchUut9.SensorOutput := FALSE;
   BenchUut9.washComplete := FALSE;
   BenchUut9.weightComplete := FALSE;
   BenchUut9.weight := REAL#150.0;
   BenchUut9.firingComplete := FALSE;
   TraceIn_Mode[136] := BenchUut9.Mode;
   TraceIn_ForwardButton[136] := BenchUut9.ForwardButton;
   TraceIn_ReverseButton[136] := BenchUut9.ReverseButton;
   TraceIn_SensorFeed[136] := BenchUut9.SensorFeed;
   TraceIn_SensorWash[136] := BenchUut9.SensorWash;
   TraceIn_SensorWeight[136] := BenchUut9.SensorWeight;
   TraceIn_SensorFiring[136] := BenchUut9.SensorFiring;
   TraceIn_SensorOutput[136] := BenchUut9.SensorOutput;
   TraceIn_washComplete[136] := BenchUut9.washComplete;
   TraceIn_weightComplete[136] := BenchUut9.weightComplete;
   TraceIn_weight[136] := BenchUut9.weight;
   TraceIn_firingComplete[136] := BenchUut9.firingComplete;
   BenchUut9();
   TraceOut_MotorForward[136] := BenchUut9.MotorForward;
   TraceOut_MotorReverse[136] := BenchUut9.MotorReverse;
   TraceOut_kick[136] := BenchUut9.kick;
   TraceOut_CompletionLight[136] := BenchUut9.CompletionLight;
   TraceOut_firingTemp[136] := BenchUut9.firingTemp;
   BenchCalls := BenchCalls + 1;
 137:
   BenchUut9.Mode := TRUE;
   BenchUut9.ForwardButton := FALSE;
   BenchUut9.ReverseButton := FALSE;
   BenchUut9.SensorFeed := FALSE;
   BenchUut9.SensorWash := FALSE;
   BenchUut9.SensorWeight := FALSE;
   BenchUut9.SensorFiring := TRUE;
   BenchUut9.SensorOutput := FALSE;
   BenchUut9.washComplete := FALSE;
   BenchUut9.weightComplete := FALSE;
   BenchUut9.weight := REAL#150.0;
   BenchUut9.firingComplete := FALSE;
   TraceIn_Mode[137] := BenchUut9.Mode;
   TraceIn_ForwardButton[137] := BenchUut9.ForwardButton;
   TraceIn_ReverseButton[137] := BenchUut9.ReverseButton;
   TraceIn_SensorFeed[137] := BenchUut9.SensorFeed;
   TraceIn_SensorWash[137] := BenchUut9.SensorWash;
   TraceIn_SensorWeight[137] := BenchUut9.SensorWeight;
   TraceIn_SensorFiring[137] := BenchUut9.SensorFiring;
   TraceIn_SensorOutput[137] := BenchUut9.SensorOutput;
   TraceIn_washComplete[137] := BenchUut9.washComplete;
   TraceIn_weightComplete[137] := BenchUut9.weightComplete;
   TraceIn_weight[137] := BenchUut9.weight;
   TraceIn_firingComplete[137] := BenchUut9.firingComplete;
   BenchUut9();
   TraceOut_MotorForward[137] := BenchUut9.MotorForward;
   TraceOut_MotorReverse[137] := BenchUut9.MotorReverse;
   TraceOut_kick[137] := BenchUut9.kick;
   TraceOut_CompletionLight[137] := BenchUut9.CompletionLight;
   TraceOut_firingTemp[137] := BenchUut9.firingTemp;
   BenchCalls := BenchCalls + 1;
 138:
   BenchUut9.Mode := TRUE;
   BenchUut9.ForwardButton := FALSE;
   BenchUut9.ReverseButton := FALSE;
   BenchUut9.SensorFeed := FALSE;
   BenchUut9.SensorWash := FALSE;
   BenchUut9.SensorWeight := FALSE;
   BenchUut9.SensorFiring := TRUE;
   BenchUut9.SensorOutput := FALSE;
   BenchUut9.washComplete := FALSE;
   BenchUut9.weightComplete := FALSE;
   BenchUut9.weight := REAL#150.0;
   BenchUut9.firingComplete := FALSE;
   TraceIn_Mode[138] := BenchUut9.Mode;
   TraceIn_ForwardButton[138] := BenchUut9.ForwardButton;
   TraceIn_ReverseButton[138] := BenchUut9.ReverseButton;
   TraceIn_SensorFeed[138] := BenchUut9.SensorFeed;
   TraceIn_SensorWash[138] := BenchUut9.SensorWash;
   TraceIn_SensorWeight[138] := BenchUut9.SensorWeight;
   TraceIn_SensorFiring[138] := BenchUut9.SensorFiring;
   TraceIn_SensorOutput[138] := BenchUut9.SensorOutput;
   TraceIn_washComplete[138] := BenchUut9.washComplete;
   TraceIn_weightComplete[138] := BenchUut9.weightComplete;
   TraceIn_weight[138] := BenchUut9.weight;
   TraceIn_firingComplete[138] := BenchUut9.firingComplete;
   BenchUut9();
   TraceOut_MotorForward[138] := BenchUut9.MotorForward;
   TraceOut_MotorReverse[138] := BenchUut9.MotorReverse;
   TraceOut_kick[138] := BenchUut9.kick;
   TraceOut_CompletionLight[138] := BenchUut9.CompletionLight;
   TraceOut_firingTemp[138] := BenchUut9.firingTemp;
   BenchCalls := BenchCalls + 1;
 139:
   BenchUut9.Mode := TRUE;
   BenchUut9.ForwardButton := FALSE;
   BenchUut9.ReverseButton := FALSE;
   BenchUut9.SensorFeed := FALSE;
   BenchUut9.SensorWash := FALSE;
   BenchUut9.SensorWeight := FALSE;
   BenchUut9.SensorFiring := TRUE;
   BenchUut9.SensorOutput := FALSE;
   BenchUut9.washComplete := FALSE;
   BenchUut9.weightComplete := FALSE;
   BenchUut9.weight := REAL#150.0;
   BenchUut9.firingComplete := TRUE;
   TraceIn_Mode[139] := BenchUut9.Mode;
   TraceIn_ForwardButton[139] := BenchUut9.ForwardButton;
   TraceIn_ReverseButton[139] := BenchUut9.ReverseButton;
   TraceIn_SensorFeed[139] := BenchUut9.SensorFeed;
   TraceIn_SensorWash[139] := BenchUut9.SensorWash;
   TraceIn_SensorWeight[139] := BenchUut9.SensorWeight;
   TraceIn_SensorFiring[139] := BenchUut9.SensorFiring;
   TraceIn_SensorOutput[139] := BenchUut9.SensorOutput;
   TraceIn_washComplete[139] := BenchUut9.washComplete;
   TraceIn_weightComplete[139] := BenchUut9.weightComplete;
   TraceIn_weight[139] := BenchUut9.weight;
   TraceIn_firingComplete[139] := BenchUut9.firingComplete;
   BenchUut9();
   TraceOut_MotorForward[139] := BenchUut9.MotorForward;
   TraceOut_MotorReverse[139] := BenchUut9.MotorReverse;
   TraceOut_kick[139] := BenchUut9.kick;
   TraceOut_CompletionLight[139] := BenchUut9.CompletionLight;
   TraceOut_firingTemp[139] := BenchUut9.firingTemp;
   BenchCalls := BenchCalls + 1;
 140:
   BenchUut9.Mode := TRUE;
   BenchUut9.ForwardButton := FALSE;
   BenchUut9.ReverseButton := FALSE;
   BenchUut9.SensorFeed := FALSE;
   BenchUut9.SensorWash := FALSE;
   BenchUut9.SensorWeight := FALSE;
   BenchUut9.SensorFiring := FALSE;
   BenchUut9.SensorOutput := FALSE;
   BenchUut9.washComplete := FALSE;
   BenchUut9.weightComplete := FALSE;
   BenchUut9.weight := REAL#150.0;
   BenchUut9.firingComplete := FALSE;
   TraceIn_Mode[140] := BenchUut9.Mode;
   TraceIn_ForwardButton[140] := BenchUut9.ForwardButton;
   TraceIn_ReverseButton[140] := BenchUut9.ReverseButton;
   TraceIn_SensorFeed[140] := BenchUut9.SensorFeed;
   TraceIn_SensorWash[140] := BenchUut9.SensorWash;
   TraceIn_SensorWeight[140] := BenchUut9.SensorWeight;
   TraceIn_SensorFiring[140] := BenchUut9.SensorFiring;
   TraceIn_SensorOutput[140] := BenchUut9.SensorOutput;
   TraceIn_washComplete[140] := BenchUut9.washComplete;
   TraceIn_weightComplete[140] := BenchUut9.weightComplete;
   TraceIn_weight[140] := BenchUut9.weight;
   TraceIn_firingComplete[140] := BenchUut9.firingComplete;
   BenchUut9();
   TraceOut_MotorForward[140] := BenchUut9.MotorForward;
   TraceOut_MotorReverse[140] := BenchUut9.MotorReverse;
   TraceOut_kick[140] := BenchUut9.kick;
   TraceOut_CompletionLight[140] := BenchUut9.CompletionLight;
   TraceOut_firingTemp[140] := BenchUut9.firingTemp;
   BenchCalls := BenchCalls + 1;
 141:
   BenchUut9.Mode := TRUE;
   BenchUut9.ForwardButton := FALSE;
   BenchUut9.ReverseButton := FALSE;
   BenchUut9.SensorFeed := FALSE;
   BenchUut9.SensorWash := FALSE;
   BenchUut9.SensorWeight := FALSE;
   BenchUut9.SensorFiring := FALSE;
   BenchUut9.SensorOutput := FALSE;
   BenchUut9.washComplete := FALSE;
   BenchUut9.weightComplete := FALSE;
   BenchUut9.weight := REAL#150.0;
   BenchUut9.firingComplete := FALSE;
   TraceIn_Mode[141] := BenchUut9.Mode;
   TraceIn_ForwardButton[141] := BenchUut9.ForwardButton;
   TraceIn_ReverseButton[141] := BenchUut9.ReverseButton;
   TraceIn_SensorFeed[141] := BenchUut9.SensorFeed;
   TraceIn_SensorWash[141] := BenchUut9.SensorWash;
   TraceIn_SensorWeight[141] := BenchUut9.SensorWeight;
   TraceIn_SensorFiring[141] := BenchUut9.SensorFiring;
   TraceIn_SensorOutput[141] := BenchUut9.SensorOutput;
   TraceIn_washComplete[141] := BenchUut9.washComplete;
   TraceIn_weightComplete[141] := BenchUut9.weightComplete;
   TraceIn_weight[141] := BenchUut9.weight;
   TraceIn_firingComplete[141] := BenchUut9.firingComplete;
   BenchUut9();
   TraceOut_MotorForward[141] := BenchUut9.MotorForward;
   TraceOut_MotorReverse[141] := BenchUut9.MotorReverse;
   TraceOut_kick[141] := BenchUut9.kick;
   TraceOut_CompletionLight[141] := BenchUut9.CompletionLight;
   TraceOut_firingTemp[141] := BenchUut9.firingTemp;
   BenchCalls := BenchCalls + 1;
 142:
   BenchUut9.Mode := TRUE;
   BenchUut9.ForwardButton := FALSE;
   BenchUut9.ReverseButton := FALSE;
   BenchUut9.SensorFeed := FALSE;
   BenchUut9.SensorWash := FALSE;
   BenchUut9.SensorWeight := FALSE;
   BenchUut9.SensorFiring := FALSE;
   BenchUut9.SensorOutput := FALSE;
   BenchUut9.washComplete := FALSE;
   BenchUut9.weightComplete := FALSE;
   BenchUut9.weight := REAL#150.0;
   BenchUut9.firingComplete := FALSE;
   TraceIn_Mode[142] := BenchUut9.Mode;
   TraceIn_ForwardButton[142] := BenchUut9.ForwardButton;
   TraceIn_ReverseButton[142] := BenchUut9.ReverseButton;
   TraceIn_SensorFeed[142] := BenchUut9.SensorFeed;
   TraceIn_SensorWash[142] := BenchUut9.SensorWash;
   TraceIn_SensorWeight[142] := BenchUut9.SensorWeight;
   TraceIn_SensorFiring[142] := BenchUut9.SensorFiring;
   TraceIn_SensorOutput[142] := BenchUut9.SensorOutput;
   TraceIn_washComplete[142] := BenchUut9.washComplete;
   TraceIn_weightComplete[142] := BenchUut9.weightComplete;
   TraceIn_weight[142] := BenchUut9.weight;
   TraceIn_firingComplete[142] := BenchUut9.firingComplete;
   BenchUut9();
   TraceOut_MotorForward[142] := BenchUut9.MotorForward;
   TraceOut_MotorReverse[142] := BenchUut9.MotorReverse;
   TraceOut_kick[142] := BenchUut9.kick;
   TraceOut_CompletionLight[142] := BenchUut9.CompletionLight;
   TraceOut_firingTemp[142] := BenchUut9.firingTemp;
   BenchCalls := BenchCalls + 1;
 143:
   BenchUut9.Mode := TRUE;
   BenchUut9.ForwardButton := FALSE;
   BenchUut9.ReverseButton := FALSE;
   BenchUut9.SensorFeed := FALSE;
   BenchUut9.SensorWash := FALSE;
   BenchUut9.SensorWeight := FALSE;
   BenchUut9.SensorFiring := FALSE;
   BenchUut9.SensorOutput := TRUE;
   BenchUut9.washComplete := FALSE;
   BenchUut9.weightComplete := FALSE;
   BenchUut9.weight := REAL#150.0;
   BenchUut9.firingComplete := FALSE;
   TraceIn_Mode[143] := BenchUut9.Mode;
   TraceIn_ForwardButton[143] := BenchUut9.ForwardButton;
   TraceIn_ReverseButton[143] := BenchUut9.ReverseButton;
   TraceIn_SensorFeed[143] := BenchUut9.SensorFeed;
   TraceIn_SensorWash[143] := BenchUut9.SensorWash;
   TraceIn_SensorWeight[143] := BenchUut9.SensorWeight;
   TraceIn_SensorFiring[143] := BenchUut9.SensorFiring;
   TraceIn_SensorOutput[143] := BenchUut9.SensorOutput;
   TraceIn_washComplete[143] := BenchUut9.washComplete;
   TraceIn_weightComplete[143] := BenchUut9.weightComplete;
   TraceIn_weight[143] := BenchUut9.weight;
   TraceIn_firingComplete[143] := BenchUut9.firingComplete;
   BenchUut9();
   TraceOut_MotorForward[143] := BenchUut9.MotorForward;
   TraceOut_MotorReverse[143] := BenchUut9.MotorReverse;
   TraceOut_kick[143] := BenchUut9.kick;
   TraceOut_CompletionLight[143] := BenchUut9.CompletionLight;
   TraceOut_firingTemp[143] := BenchUut9.firingTemp;
   BenchCalls := BenchCalls + 1;
 144:
   BenchUut9.Mode := TRUE;
   BenchUut9.ForwardButton := FALSE;
   BenchUut9.ReverseButton := FALSE;
   BenchUut9.SensorFeed := FALSE;
   BenchUut9.SensorWash := FALSE;
   BenchUut9.SensorWeight := FALSE;
   BenchUut9.SensorFiring := FALSE;
   BenchUut9.SensorOutput := TRUE;
   BenchUut9.washComplete := FALSE;
   BenchUut9.weightComplete := FALSE;
   BenchUut9.weight := REAL#150.0;
   BenchUut9.firingComplete := FALSE;
   TraceIn_Mode[144] := BenchUut9.Mode;
   TraceIn_ForwardButton[144] := BenchUut9.ForwardButton;
   TraceIn_ReverseButton[144] := BenchUut9.ReverseButton;
   TraceIn_SensorFeed[144] := BenchUut9.SensorFeed;
   TraceIn_SensorWash[144] := BenchUut9.SensorWash;
   TraceIn_SensorWeight[144] := BenchUut9.SensorWeight;
   TraceIn_SensorFiring[144] := BenchUut9.SensorFiring;
   TraceIn_SensorOutput[144] := BenchUut9.SensorOutput;
   TraceIn_washComplete[144] := BenchUut9.washComplete;
   TraceIn_weightComplete[144] := BenchUut9.weightComplete;
   TraceIn_weight[144] := BenchUut9.weight;
   TraceIn_firingComplete[144] := BenchUut9.firingComplete;
   BenchUut9();
   TraceOut_MotorForward[144] := BenchUut9.MotorForward;
   TraceOut_MotorReverse[144] := BenchUut9.MotorReverse;
   TraceOut_kick[144] := BenchUut9.kick;
   TraceOut_CompletionLight[144] := BenchUut9.CompletionLight;
   TraceOut_firingTemp[144] := BenchUut9.firingTemp;
   BenchCalls := BenchCalls + 1;
 145:
   BenchUut9.Mode := TRUE;
   BenchUut9.ForwardButton := FALSE;
   BenchUut9.ReverseButton := FALSE;
   BenchUut9.SensorFeed := FALSE;
   BenchUut9.SensorWash := FALSE;
   BenchUut9.SensorWeight := FALSE;
   BenchUut9.SensorFiring := FALSE;
   BenchUut9.SensorOutput := TRUE;
   BenchUut9.washComplete := FALSE;
   BenchUut9.weightComplete := FALSE;
   BenchUut9.weight := REAL#150.0;
   BenchUut9.firingComplete := FALSE;
   TraceIn_Mode[145] := BenchUut9.Mode;
   TraceIn_ForwardButton[145] := BenchUut9.ForwardButton;
   TraceIn_ReverseButton[145] := BenchUut9.ReverseButton;
   TraceIn_SensorFeed[145] := BenchUut9.SensorFeed;
   TraceIn_SensorWash[145] := BenchUut9.SensorWash;
   TraceIn_SensorWeight[145] := BenchUut9.SensorWeight;
   TraceIn_SensorFiring[145] := BenchUut9.SensorFiring;
   TraceIn_SensorOutput[145] := BenchUut9.SensorOutput;
   TraceIn_washComplete[145] := BenchUut9.washComplete;
   TraceIn_weightComplete[145] := BenchUut9.weightComplete;
   TraceIn_weight[145] := BenchUut9.weight;
   TraceIn_firingComplete[145] := BenchUut9.firingComplete;
   BenchUut9();
   TraceOut_MotorForward[145] := BenchUut9.MotorForward;
   TraceOut_MotorReverse[145] := BenchUut9.MotorReverse;
   TraceOut_kick[145] := BenchUut9.kick;
   TraceOut_CompletionLight[145] := BenchUut9.CompletionLight;
   TraceOut_firingTemp[145] := BenchUut9.firingTemp;
   BenchCalls := BenchCalls + 1;
 146:
   BenchUut9.Mode := TRUE;
   BenchUut9.ForwardButton := FALSE;
   BenchUut9.ReverseButton := FALSE;
   BenchUut9.SensorFeed := FALSE;
   BenchUut9.SensorWash := FALSE;
   BenchUut9.SensorWeight := FALSE;
   BenchUut9.SensorFiring := FALSE;
   BenchUut9.SensorOutput := FALSE;
   BenchUut9.washComplete := FALSE;
   BenchUut9.weightComplete := FALSE;
   BenchUut9.weight := REAL#150.0;
   BenchUut9.firingComplete := FALSE;
   TraceIn_Mode[146] := BenchUut9.Mode;
   TraceIn_ForwardButton[146] := BenchUut9.ForwardButton;
   TraceIn_ReverseButton[146] := BenchUut9.ReverseButton;
   TraceIn_SensorFeed[146] := BenchUut9.SensorFeed;
   TraceIn_SensorWash[146] := BenchUut9.SensorWash;
   TraceIn_SensorWeight[146] := BenchUut9.SensorWeight;
   TraceIn_SensorFiring[146] := BenchUut9.SensorFiring;
   TraceIn_SensorOutput[146] := BenchUut9.SensorOutput;
   TraceIn_washComplete[146] := BenchUut9.washComplete;
   TraceIn_weightComplete[146] := BenchUut9.weightComplete;
   TraceIn_weight[146] := BenchUut9.weight;
   TraceIn_firingComplete[146] := BenchUut9.firingComplete;
   BenchUut9();
   TraceOut_MotorForward[146] := BenchUut9.MotorForward;
   TraceOut_MotorReverse[146] := BenchUut9.MotorReverse;
   TraceOut_kick[146] := BenchUut9.kick;
   TraceOut_CompletionLight[146] := BenchUut9.CompletionLight;
   TraceOut_firingTemp[146] := BenchUut9.firingTemp;
   BenchCalls := BenchCalls + 1;
 147:
   BenchUut10.Mode := TRUE;
   BenchUut10.ForwardButton := FALSE;
   BenchUut10.ReverseButton := FALSE;
   BenchUut10.SensorFeed := TRUE;
   BenchUut10.SensorWash := FALSE;
   BenchUut10.SensorWeight := FALSE;
   BenchUut10.SensorFiring := FALSE;
   BenchUut10.SensorOutput := FALSE;
   BenchUut10.washComplete := FALSE;
   BenchUut10.weightComplete := FALSE;
   BenchUut10.weight := REAL#150.0;
   BenchUut10.firingComplete := FALSE;
   TraceIn_Mode[147] := BenchUut10.Mode;
   TraceIn_ForwardButton[147] := BenchUut10.ForwardButton;
   TraceIn_ReverseButton[147] := BenchUut10.ReverseButton;
   TraceIn_SensorFeed[147] := BenchUut10.SensorFeed;
   TraceIn_SensorWash[147] := BenchUut10.SensorWash;
   TraceIn_SensorWeight[147] := BenchUut10.SensorWeight;
   TraceIn_SensorFiring[147] := BenchUut10.SensorFiring;
   TraceIn_SensorOutput[147] := BenchUut10.SensorOutput;
   TraceIn_washComplete[147] := BenchUut10.washComplete;
   TraceIn_weightComplete[147] := BenchUut10.weightComplete;
   TraceIn_weight[147] := BenchUut10.weight;
   TraceIn_firingComplete[147] := BenchUut10.firingComplete;
   BenchUut10();
   TraceOut_MotorForward[147] := BenchUut10.MotorForward;
   TraceOut_MotorReverse[147] := BenchUut10.MotorReverse;
   TraceOut_kick[147] := BenchUut10.kick;
   TraceOut_CompletionLight[147] := BenchUut10.CompletionLight;
   TraceOut_firingTemp[147] := BenchUut10.firingTemp;
   BenchCalls := BenchCalls + 1;
 148:
   BenchUut10.Mode := TRUE;
   BenchUut10.ForwardButton := FALSE;
   BenchUut10.ReverseButton := FALSE;
   BenchUut10.SensorFeed := FALSE;
   BenchUut10.SensorWash := FALSE;
   BenchUut10.SensorWeight := FALSE;
   BenchUut10.SensorFiring := FALSE;
   BenchUut10.SensorOutput := FALSE;
   BenchUut10.washComplete := FALSE;
   BenchUut10.weightComplete := FALSE;
   BenchUut10.weight := REAL#150.0;
   BenchUut10.firingComplete := FALSE;
   TraceIn_Mode[148] := BenchUut10.Mode;
   TraceIn_ForwardButton[148] := BenchUut10.ForwardButton;
   TraceIn_ReverseButton[148] := BenchUut10.ReverseButton;
   TraceIn_SensorFeed[148] := BenchUut10.SensorFeed;
   TraceIn_SensorWash[148] := BenchUut10.SensorWash;
   TraceIn_SensorWeight[148] := BenchUut10.SensorWeight;
   TraceIn_SensorFiring[148] := BenchUut10.SensorFiring;
   TraceIn_SensorOutput[148] := BenchUut10.SensorOutput;
   TraceIn_washComplete[148] := BenchUut10.washComplete;
   TraceIn_weightComplete[148] := BenchUut10.weightComplete;
   TraceIn_weight[148] := BenchUut10.weight;
   TraceIn_firingComplete[148] := BenchUut10.firingComplete;
   BenchUut10();
   TraceOut_MotorForward[148] := BenchUut10.MotorForward;
   TraceOut_MotorReverse[148] := BenchUut10.MotorReverse;
   TraceOut_kick[148] := BenchUut10.kick;
   TraceOut_CompletionLight[148] := BenchUut10.CompletionLight;
   TraceOut_firingTemp[148] := BenchUut10.firingTemp;
   BenchCalls := BenchCalls + 1;
 149:
   BenchUut10.Mode := TRUE;
   BenchUut10.ForwardButton := FALSE;
   BenchUut10.ReverseButton := FALSE;
   BenchUut10.SensorFeed := FALSE;
   BenchUut10.SensorWash := FALSE;
   BenchUut10.SensorWeight := FALSE;
   BenchUut10.SensorFiring := FALSE;
   BenchUut10.SensorOutput := FALSE;
   BenchUut10.washComplete := FALSE;
   BenchUut10.weightComplete := FALSE;
   BenchUut10.weight := REAL#150.0;
   BenchUut10.firingComplete := FALSE;
   TraceIn_Mode[149] := BenchUut10.Mode;
   TraceIn_ForwardButton[149] := BenchUut10.ForwardButton;
   TraceIn_ReverseButton[149] := BenchUut10.ReverseButton;
   TraceIn_SensorFeed[149] := BenchUut10.SensorFeed;
   TraceIn_SensorWash[149] := BenchUut10.SensorWash;
   TraceIn_SensorWeight[149] := BenchUut10.SensorWeight;
   TraceIn_SensorFiring[149] := BenchUut10.SensorFiring;
   TraceIn_SensorOutput[149] := BenchUut10.SensorOutput;
   TraceIn_washComplete[149] := BenchUut10.washComplete;
   TraceIn_weightComplete[149] := BenchUut10.weightComplete;
   TraceIn_weight[149] := BenchUut10.weight;
   TraceIn_firingComplete[149] := BenchUut10.firingComplete;
   BenchUut10();
   TraceOut_MotorForward[149] := BenchUut10.MotorForward;
   TraceOut_MotorReverse[149] := BenchUut10.MotorReverse;
   TraceOut_kick[149] := BenchUut10.kick;
   TraceOut_CompletionLight[149] := BenchUut10.CompletionLight;
   TraceOut_firingTemp[149] := BenchUut10.firingTemp;
   BenchCalls := BenchCalls + 1;
 150:
   BenchUut10.Mode := TRUE;
   BenchUut10.ForwardButton := FALSE;
   BenchUut10.ReverseButton := FALSE;
   BenchUut10.SensorFeed := FALSE;
   BenchUut10.SensorWash := FALSE;
   BenchUut10.SensorWeight := FALSE;
   BenchUut10.SensorFiring := FALSE;
   BenchUut10.SensorOutput := FALSE;
   BenchUut10.washComplete := FALSE;
   BenchUut10.weightComplete := FALSE;
   BenchUut10.weight := REAL#150.0;
   BenchUut10.firingComplete := FALSE;
   TraceIn_Mode[150] := BenchUut10.Mode;
   TraceIn_ForwardButton[150] := BenchUut10.ForwardButton;
   TraceIn_ReverseButton[150] := BenchUut10.ReverseButton;
   TraceIn_SensorFeed[150] := BenchUut10.SensorFeed;
   TraceIn_SensorWash[150] := BenchUut10.SensorWash;
   TraceIn_SensorWeight[150] := BenchUut10.SensorWeight;
   TraceIn_SensorFiring[150] := BenchUut10.SensorFiring;
   TraceIn_SensorOutput[150] := BenchUut10.SensorOutput;
   TraceIn_washComplete[150] := BenchUut10.washComplete;
   TraceIn_weightComplete[150] := BenchUut10.weightComplete;
   TraceIn_weight[150] := BenchUut10.weight;
   TraceIn_firingComplete[150] := BenchUut10.firingComplete;
   BenchUut10();
   TraceOut_MotorForward[150] := BenchUut10.MotorForward;
   TraceOut_MotorReverse[150] := BenchUut10.MotorReverse;
   TraceOut_kick[150] := BenchUut10.kick;
   TraceOut_CompletionLight[150] := BenchUut10.CompletionLight;
   TraceOut_firingTemp[150] := BenchUut10.firingTemp;
   BenchCalls := BenchCalls + 1;
 151:
   BenchUut10.Mode := TRUE;
   BenchUut10.ForwardButton := FALSE;
   BenchUut10.ReverseButton := FALSE;
   BenchUut10.SensorFeed := FALSE;
   BenchUut10.SensorWash := TRUE;
   BenchUut10.SensorWeight := FALSE;
   BenchUut10.SensorFiring := FALSE;
   BenchUut10.SensorOutput := FALSE;
   BenchUut10.washComplete := FALSE;
   BenchUut10.weightComplete := FALSE;
   BenchUut10.weight := REAL#150.0;
   BenchUut10.firingComplete := FALSE;
   TraceIn_Mode[151] := BenchUut10.Mode;
   TraceIn_ForwardButton[151] := BenchUut10.ForwardButton;
   TraceIn_ReverseButton[151] := BenchUut10.ReverseButton;
   TraceIn_SensorFeed[151] := BenchUut10.SensorFeed;
   TraceIn_SensorWash[151] := BenchUut10.SensorWash;
   TraceIn_SensorWeight[151] := BenchUut10.SensorWeight;
   TraceIn_SensorFiring[151] := BenchUut10.SensorFiring;
   TraceIn_SensorOutput[151] := BenchUut10.SensorOutput;
   TraceIn_washComplete[151] := BenchUut10.washComplete;
   TraceIn_weightComplete[151] := BenchUut10.weightComplete;
   TraceIn_weight[151] := BenchUut10.weight;
   TraceIn_firingComplete[151] := BenchUut10.firingComplete;
   BenchUut10();
   TraceOut_MotorForward[151] := BenchUut10.MotorForward;
   TraceOut_MotorReverse[151] := BenchUut10.MotorReverse;
   TraceOut_kick[151] := BenchUut10.kick;
   TraceOut_CompletionLight[151] := BenchUut10.CompletionLight;
   TraceOut_firingTemp[151] := BenchUut10.firingTemp;
   BenchCalls := BenchCalls + 1;
 152:
   BenchUut10.Mode := TRUE;
   BenchUut10.ForwardButton := FALSE;
   BenchUut10.ReverseButton := FALSE;
   BenchUut10.SensorFeed := FALSE;
   BenchUut10.SensorWash := TRUE;
   BenchUut10.SensorWeight := FALSE;
   BenchUut10.SensorFiring := FALSE;
   BenchUut10.SensorOutput := FALSE;
   BenchUut10.washComplete := FALSE;
   BenchUut10.weightComplete := FALSE;
   BenchUut10.weight := REAL#150.0;
   BenchUut10.firingComplete := FALSE;
   TraceIn_Mode[152] := BenchUut10.Mode;
   TraceIn_ForwardButton[152] := BenchUut10.ForwardButton;
   TraceIn_ReverseButton[152] := BenchUut10.ReverseButton;
   TraceIn_SensorFeed[152] := BenchUut10.SensorFeed;
   TraceIn_SensorWash[152] := BenchUut10.SensorWash;
   TraceIn_SensorWeight[152] := BenchUut10.SensorWeight;
   TraceIn_SensorFiring[152] := BenchUut10.SensorFiring;
   TraceIn_SensorOutput[152] := BenchUut10.SensorOutput;
   TraceIn_washComplete[152] := BenchUut10.washComplete;
   TraceIn_weightComplete[152] := BenchUut10.weightComplete;
   TraceIn_weight[152] := BenchUut10.weight;
   TraceIn_firingComplete[152] := BenchUut10.firingComplete;
   BenchUut10();
   TraceOut_MotorForward[152] := BenchUut10.MotorForward;
   TraceOut_MotorReverse[152] := BenchUut10.MotorReverse;
   TraceOut_kick[152] := BenchUut10.kick;
   TraceOut_CompletionLight[152] := BenchUut10.CompletionLight;
   TraceOut_firingTemp[152] := BenchUut10.firingTemp;
   BenchCalls := BenchCalls + 1;
 153:
   BenchUut10.Mode := FALSE;
   BenchUut10.ForwardButton := FALSE;
   BenchUut10.ReverseButton := FALSE;
   BenchUut10.SensorFeed := FALSE;
   BenchUut10.SensorWash := TRUE;
   BenchUut10.SensorWeight := FALSE;
   BenchUut10.SensorFiring := FALSE;
   BenchUut10.SensorOutput := FALSE;
   BenchUut10.washComplete := FALSE;
   BenchUut10.weightComplete := FALSE;
   BenchUut10.weight := REAL#150.0;
   BenchUut10.firingComplete := FALSE;
   TraceIn_Mode[153] := BenchUut10.Mode;
   TraceIn_ForwardButton[153] := BenchUut10.ForwardButton;
   TraceIn_ReverseButton[153] := BenchUut10.ReverseButton;
   TraceIn_SensorFeed[153] := BenchUut10.SensorFeed;
   TraceIn_SensorWash[153] := BenchUut10.SensorWash;
   TraceIn_SensorWeight[153] := BenchUut10.SensorWeight;
   TraceIn_SensorFiring[153] := BenchUut10.SensorFiring;
   TraceIn_SensorOutput[153] := BenchUut10.SensorOutput;
   TraceIn_washComplete[153] := BenchUut10.washComplete;
   TraceIn_weightComplete[153] := BenchUut10.weightComplete;
   TraceIn_weight[153] := BenchUut10.weight;
   TraceIn_firingComplete[153] := BenchUut10.firingComplete;
   BenchUut10();
   TraceOut_MotorForward[153] := BenchUut10.MotorForward;
   TraceOut_MotorReverse[153] := BenchUut10.MotorReverse;
   TraceOut_kick[153] := BenchUut10.kick;
   TraceOut_CompletionLight[153] := BenchUut10.CompletionLight;
   TraceOut_firingTemp[153] := BenchUut10.firingTemp;
   BenchCalls := BenchCalls + 1;
 154:
   BenchUut10.Mode := TRUE;
   BenchUut10.ForwardButton := FALSE;
   BenchUut10.ReverseButton := FALSE;
   BenchUut10.SensorFeed := FALSE;
   BenchUut10.SensorWash := TRUE;
   BenchUut10.SensorWeight := FALSE;
   BenchUut10.SensorFiring := FALSE;
   BenchUut10.SensorOutput := FALSE;
   BenchUut10.washComplete := FALSE;
   BenchUut10.weightComplete := FALSE;
   BenchUut10.weight := REAL#150.0;
   BenchUut10.firingComplete := FALSE;
   TraceIn_Mode[154] := BenchUut10.Mode;
   TraceIn_ForwardButton[154] := BenchUut10.ForwardButton;
   TraceIn_ReverseButton[154] := BenchUut10.ReverseButton;
   TraceIn_SensorFeed[154] := BenchUut10.SensorFeed;
   TraceIn_SensorWash[154] := BenchUut10.SensorWash;
   TraceIn_SensorWeight[154] := BenchUut10.SensorWeight;
   TraceIn_SensorFiring[154] := BenchUut10.SensorFiring;
   TraceIn_SensorOutput[154] := BenchUut10.SensorOutput;
   TraceIn_washComplete[154] := BenchUut10.washComplete;
   TraceIn_weightComplete[154] := BenchUut10.weightComplete;
   TraceIn_weight[154] := BenchUut10.weight;
   TraceIn_firingComplete[154] := BenchUut10.firingComplete;
   BenchUut10();
   TraceOut_MotorForward[154] := BenchUut10.MotorForward;
   TraceOut_MotorReverse[154] := BenchUut10.MotorReverse;
   TraceOut_kick[154] := BenchUut10.kick;
   TraceOut_CompletionLight[154] := BenchUut10.CompletionLight;
   TraceOut_firingTemp[154] := BenchUut10.firingTemp;
   BenchCalls := BenchCalls + 1;
 155:
   BenchUut10.Mode := TRUE;
   BenchUut10.ForwardButton := FALSE;
   BenchUut10.ReverseButton := FALSE;
   BenchUut10.SensorFeed := TRUE;
   BenchUut10.SensorWash := TRUE;
   BenchUut10.SensorWeight := FALSE;
   BenchUut10.SensorFiring := FALSE;
   BenchUut10.SensorOutput := FALSE;
   BenchUut10.washComplete := FALSE;
   BenchUut10.weightComplete := FALSE;
   BenchUut10.weight := REAL#150.0;
   BenchUut10.firingComplete := FALSE;
   TraceIn_Mode[155] := BenchUut10.Mode;
   TraceIn_ForwardButton[155] := BenchUut10.ForwardButton;
   TraceIn_ReverseButton[155] := BenchUut10.ReverseButton;
   TraceIn_SensorFeed[155] := BenchUut10.SensorFeed;
   TraceIn_SensorWash[155] := BenchUut10.SensorWash;
   TraceIn_SensorWeight[155] := BenchUut10.SensorWeight;
   TraceIn_SensorFiring[155] := BenchUut10.SensorFiring;
   TraceIn_SensorOutput[155] := BenchUut10.SensorOutput;
   TraceIn_washComplete[155] := BenchUut10.washComplete;
   TraceIn_weightComplete[155] := BenchUut10.weightComplete;
   TraceIn_weight[155] := BenchUut10.weight;
   TraceIn_firingComplete[155] := BenchUut10.firingComplete;
   BenchUut10();
   TraceOut_MotorForward[155] := BenchUut10.MotorForward;
   TraceOut_MotorReverse[155] := BenchUut10.MotorReverse;
   TraceOut_kick[155] := BenchUut10.kick;
   TraceOut_CompletionLight[155] := BenchUut10.CompletionLight;
   TraceOut_firingTemp[155] := BenchUut10.firingTemp;
   BenchCalls := BenchCalls + 1;
 END_CASE;
 BenchStep := BenchStep + 1;
 IF BenchStep >= 156 THEN BenchDone := TRUE; END_IF;
END_IF;
END_PROGRAM
